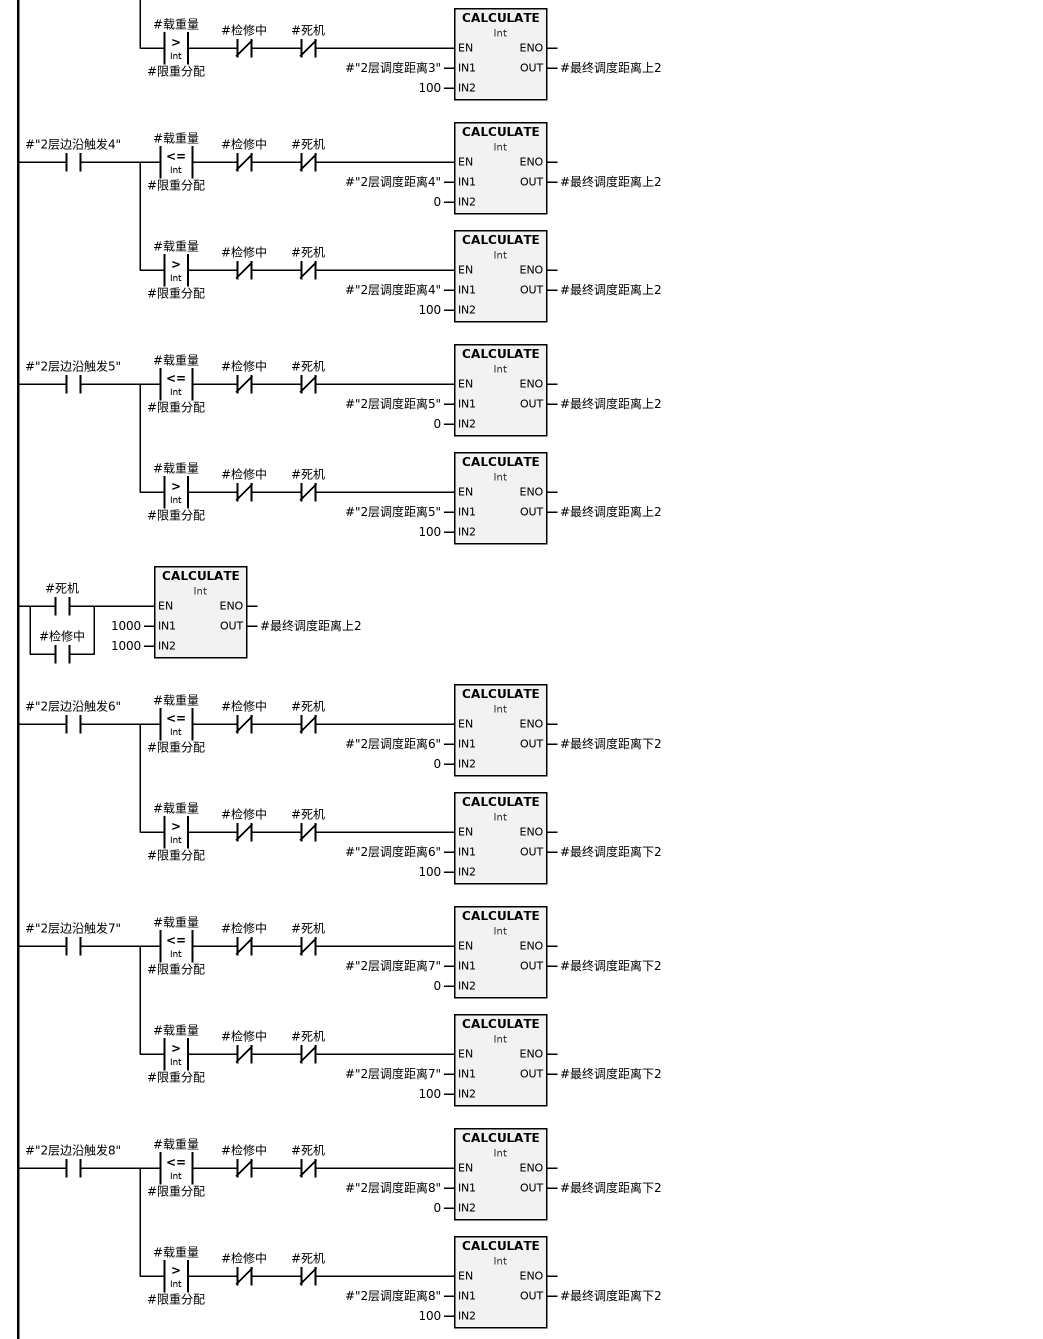
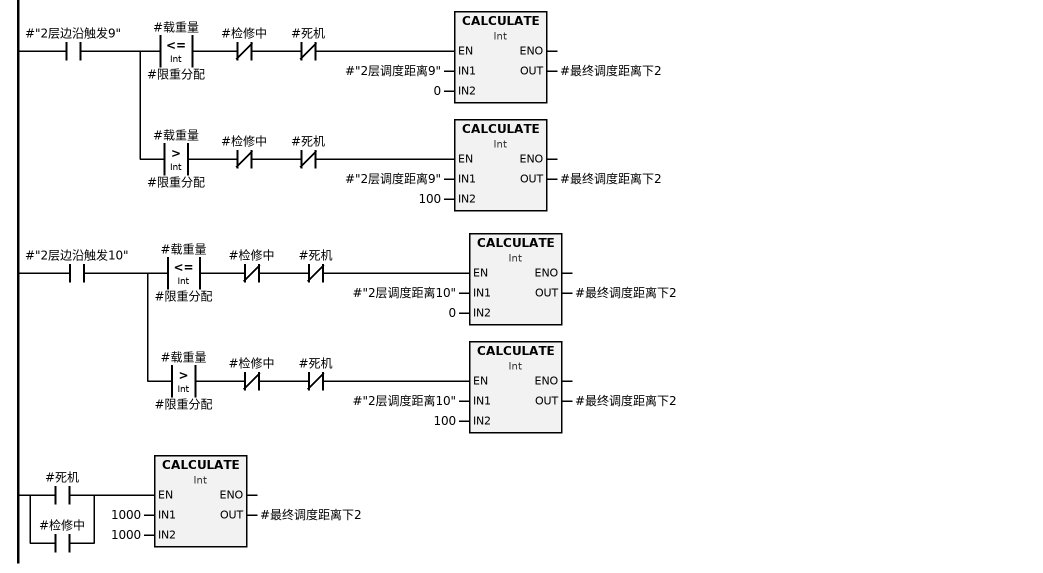
   RUNG wire#powerrail
      Contact( #上呼灯2 )
      wire#w1
      I_Contact( #上行指示 )
      I_Contact( #下行指示 )
      { S7_Templates := "SrcType := Int" } LE_Contact(in1 := #当前楼层, in2 := 2)
      wire#w2
      { S7_Templates := "SrcType := Int"; S7_Expression := "ABS(IN1-IN2)" } Calculate(in1 := #当前楼层, in2 := 2, in3 := 0, out => #"2层调度距离1")
      Coil( #"2层边沿触发1" )
   END_RUNG
   RUNG wire#w1
      Contact( #上行指示 )
      wire#w3
      { S7_Templates := "SrcType := Int" } EQ_Contact(in1 := 2, in2 := #当前楼层)
      Contact( #上下平层都为1 )
   END_RUNG wire#w2
   RUNG wire#w3
      { S7_Templates := "SrcType := Int" } GT_Contact(in1 := 2, in2 := #当前楼层)
   END_RUNG wire#w2
   RUNG wire#w1
      Contact( #下行指示 )
      wire#w4
      Contact( #外呼下面无目标2 )
      { S7_Templates := "SrcType := Int"; S7_Expression := "ABS(IN1-IN2)+IN3+IN3" } Calculate(in1 := #当前楼层, in2 := 2, in3 := #下行停站次数2, out => #"2层调度距离2")
      Coil( #"2层边沿触发2" )
   END_RUNG
   RUNG wire#w1
      I_Contact( #上行指示 )
      I_Contact( #下行指示 )
      { S7_Templates := "SrcType := Int" } GT_Contact(in1 := #当前楼层, in2 := 2)
   END_RUNG wire#w4
   RUNG wire#w1
      Contact( #下行指示 )
      Contact( #外呼下面有目标2 )
      { S7_Templates := "SrcType := Int"; S7_Expression := "ABS(IN3+IN3-IN1-IN2)+IN5+IN4+IN4+IN5+IN6" } Calculate(in1 := #当前楼层, in2 := 2, in3 := #外呼下面有目标最小数2, in4 := 0, in5 := #下行停站次数1, in6 := 2, out => #"2层调度距离3")
      Coil( #"2层边沿触发3" )
   END_RUNG
   RUNG wire#w1
      Contact( #上行指示 )
      wire#w5
      { S7_Templates := "SrcType := Int" } EQ_Contact(in1 := 2, in2 := #当前楼层)
      I_Contact( #上下平层都为1 )
      wire#w6
      Contact( #外呼下面有目标2 )
      { S7_Templates := "SrcType := Int"; S7_Expression := "ABS(IN3-IN1+IN3-IN6+IN2-IN6)+IN5+IN4+IN4+IN5+IN7+IN7+IN8+IN8" } Calculate(in1 := #当前楼层, in2 := 2, in3 := #外呼上面有目标最大数2, in4 := #上行停站次数10, in5 := 0, in6 := #外呼下面有目标最小数2, in7 := #下行停站次数1, in8 := 2, out => #"2层调度距离4")
      Coil( #"2层边沿触发4" )
   END_RUNG
   RUNG wire#w5
      { S7_Templates := "SrcType := Int" } GT_Contact(in1 := #当前楼层, in2 := 2)
   END_RUNG wire#w6
   RUNG wire#w6
      Contact( #外呼下面无目标2 )
      { S7_Templates := "SrcType := Int"; S7_Expression := "ABS(IN3-IN1+IN3-IN2)+IN5+IN4+IN4+IN5+IN6" } Calculate(in1 := #当前楼层, in2 := 2, in3 := #外呼上面有目标最大数2, in4 := #上行停站次数10, in5 := #下行停站次数2, in6 := 2, out => #"2层调度距离5")
      Coil( #"2层边沿触发5" )
   END_RUNG
   RUNG wire#powerrail
      Contact( #下呼灯2 )
      wire#w7
      I_Contact( #上行指示 )
      I_Contact( #下行指示 )
      { S7_Templates := "SrcType := Int" } GE_Contact(in1 := #当前楼层, in2 := 2)
      wire#w8
      { S7_Templates := "SrcType := Int"; S7_Expression := "ABS(IN1-IN2)+IN3+IN3" } Calculate(in1 := #当前楼层, in2 := 2, in3 := #下行停站次数2, out => #"2层调度距离6")
      Coil( #"2层边沿触发6" )
   END_RUNG
   RUNG wire#w7
      Contact( #下行指示 )
      wire#w9
      { S7_Templates := "SrcType := Int" } EQ_Contact(in1 := 2, in2 := #当前楼层)
      Contact( #上下平层都为1 )
   END_RUNG wire#w8
   RUNG wire#w9
      { S7_Templates := "SrcType := Int" } GT_Contact(in1 := #当前楼层, in2 := 2)
   END_RUNG wire#w8
   RUNG wire#w7
      Contact( #上行指示 )
      wire#w10
      Contact( #外呼上面无目标2 )
      { S7_Templates := "SrcType := Int"; S7_Expression := "ABS(IN1-IN2)+IN3+IN3" } Calculate(in1 := #当前楼层, in2 := 2, in3 := 0, out => #"2层调度距离7")
      Coil( #"2层边沿触发7" )
   END_RUNG
   RUNG wire#w7
      I_Contact( #上行指示 )
      I_Contact( #下行指示 )
      { S7_Templates := "SrcType := Int" } LT_Contact(in1 := #当前楼层, in2 := 2)
   END_RUNG wire#w10
   RUNG wire#w7
      Contact( #上行指示 )
      Contact( #外呼上面有目标2 )
      { S7_Templates := "SrcType := Int"; S7_Expression := "ABS(IN3+IN3-IN1-IN2)+IN4+IN5+IN4+IN5+IN6" } Calculate(in1 := #当前楼层, in2 := 2, in3 := #外呼上面有目标最大数2, in4 := #下行停站次数2, in5 := #上行停站次数10, in6 := 2, out => #"2层调度距离8")
      Coil( #"2层边沿触发8" )
   END_RUNG
   RUNG wire#w7
      Contact( #下行指示 )
      wire#w11
      { S7_Templates := "SrcType := Int" } EQ_Contact(in1 := 2, in2 := #当前楼层)
      I_Contact( #上下平层都为1 )
      wire#w12
      Contact( #外呼上面有目标2 )
      { S7_Templates := "SrcType := Int"; S7_Expression := "ABS(IN1-IN6+IN3-IN6+IN3-IN2)+IN5+IN4+IN4+IN5+IN7+IN7+IN8" } Calculate(in1 := #当前楼层, in2 := 2, in3 := #外呼上面有目标最大数2, in4 := #下行停站次数2, in5 := #下行停站次数1, in6 := #外呼下面有目标最小数2, in7 := #上行停站次数10, in8 := 4, out => #"2层调度距离9")
      Coil( #"2层边沿触发9" )
   END_RUNG
   RUNG wire#w11
      { S7_Templates := "SrcType := Int" } GT_Contact(in1 := 2, in2 := #当前楼层)
   END_RUNG wire#w12
   RUNG wire#w12
      Contact( #外呼上面无目标2 )
      { S7_Templates := "SrcType := Int"; S7_Expression := "ABS(IN1-IN3+IN2-IN3)+IN5+IN4+IN4+IN5+IN6" } Calculate(in1 := #当前楼层, in2 := 2, in3 := #外呼下面有目标最小数2, in4 := 0, in5 := #下行停站次数1, in6 := 2, out => #"2层调度距离10")
      Coil( #"2层边沿触发10" )
   END_RUNG
   RUNG wire#powerrail
      Contact( #"2层边沿触发1" )
      wire#w13
      { S7_Templates := "SrcType := Int" } LE_Contact(in1 := #载重量, in2 := #限重分配)
      I_Contact( #检修中 )
      I_Contact( #死机 )
      { S7_Templates := "SrcType := Int"; S7_Expression := "ABS(IN1+IN2)" } Calculate(in1 := #"2层调度距离1", in2 := 0, out => #最终调度距离上2)
   END_RUNG
   RUNG wire#w13
      { S7_Templates := "SrcType := Int" } GT_Contact(in1 := #载重量, in2 := #限重分配)
      I_Contact( #检修中 )
      I_Contact( #死机 )
      { S7_Templates := "SrcType := Int"; S7_Expression := "ABS(IN1+IN2)" } Calculate(in1 := #"2层调度距离1", in2 := 100, out => #最终调度距离上2)
   END_RUNG
   RUNG wire#powerrail
      Contact( #"2层边沿触发2" )
      wire#w14
      { S7_Templates := "SrcType := Int" } LE_Contact(in1 := #载重量, in2 := #限重分配)
      I_Contact( #检修中 )
      I_Contact( #死机 )
      { S7_Templates := "SrcType := Int"; S7_Expression := "ABS(IN1+IN2)" } Calculate(in1 := #"2层调度距离2", in2 := 0, out => #最终调度距离上2)
   END_RUNG
   RUNG wire#w14
      { S7_Templates := "SrcType := Int" } GT_Contact(in1 := #载重量, in2 := #限重分配)
      I_Contact( #检修中 )
      I_Contact( #死机 )
      { S7_Templates := "SrcType := Int"; S7_Expression := "ABS(IN1+IN2)" } Calculate(in1 := #"2层调度距离2", in2 := 100, out => #最终调度距离上2)
   END_RUNG
   RUNG wire#powerrail
      Contact( #"2层边沿触发3" )
      wire#w15
      { S7_Templates := "SrcType := Int" } LE_Contact(in1 := #载重量, in2 := #限重分配)
      I_Contact( #检修中 )
      I_Contact( #死机 )
      { S7_Templates := "SrcType := Int"; S7_Expression := "ABS(IN1+IN2)" } Calculate(in1 := #"2层调度距离3", in2 := 0, out => #最终调度距离上2)
   END_RUNG
   RUNG wire#w15
      { S7_Templates := "SrcType := Int" } GT_Contact(in1 := #载重量, in2 := #限重分配)
      I_Contact( #检修中 )
      I_Contact( #死机 )
      { S7_Templates := "SrcType := Int"; S7_Expression := "ABS(IN1+IN2)" } Calculate(in1 := #"2层调度距离3", in2 := 100, out => #最终调度距离上2)
   END_RUNG
   RUNG wire#powerrail
      Contact( #"2层边沿触发4" )
      wire#w16
      { S7_Templates := "SrcType := Int" } LE_Contact(in1 := #载重量, in2 := #限重分配)
      I_Contact( #检修中 )
      I_Contact( #死机 )
      { S7_Templates := "SrcType := Int"; S7_Expression := "ABS(IN1+IN2)" } Calculate(in1 := #"2层调度距离4", in2 := 0, out => #最终调度距离上2)
   END_RUNG
   RUNG wire#w16
      { S7_Templates := "SrcType := Int" } GT_Contact(in1 := #载重量, in2 := #限重分配)
      I_Contact( #检修中 )
      I_Contact( #死机 )
      { S7_Templates := "SrcType := Int"; S7_Expression := "ABS(IN1+IN2)" } Calculate(in1 := #"2层调度距离4", in2 := 100, out => #最终调度距离上2)
   END_RUNG
   RUNG wire#powerrail
      Contact( #"2层边沿触发5" )
      wire#w17
      { S7_Templates := "SrcType := Int" } LE_Contact(in1 := #载重量, in2 := #限重分配)
      I_Contact( #检修中 )
      I_Contact( #死机 )
      { S7_Templates := "SrcType := Int"; S7_Expression := "ABS(IN1+IN2)" } Calculate(in1 := #"2层调度距离5", in2 := 0, out => #最终调度距离上2)
   END_RUNG
   RUNG wire#w17
      { S7_Templates := "SrcType := Int" } GT_Contact(in1 := #载重量, in2 := #限重分配)
      I_Contact( #检修中 )
      I_Contact( #死机 )
      { S7_Templates := "SrcType := Int"; S7_Expression := "ABS(IN1+IN2)" } Calculate(in1 := #"2层调度距离5", in2 := 100, out => #最终调度距离上2)
   END_RUNG
   RUNG wire#powerrail
      Contact( #死机 )
      wire#w18
      { S7_Templates := "SrcType := Int"; S7_Expression := "ABS(IN1+IN2)" } Calculate(in1 := 1000, in2 := 1000, out => #最终调度距离上2)
   END_RUNG
   RUNG wire#powerrail
      Contact( #检修中 )
   END_RUNG wire#w18
   RUNG wire#powerrail
      Contact( #"2层边沿触发6" )
      wire#w19
      { S7_Templates := "SrcType := Int" } LE_Contact(in1 := #载重量, in2 := #限重分配)
      I_Contact( #检修中 )
      I_Contact( #死机 )
      { S7_Templates := "SrcType := Int"; S7_Expression := "ABS(IN1+IN2)" } Calculate(in1 := #"2层调度距离6", in2 := 0, out => #最终调度距离下2)
   END_RUNG
   RUNG wire#w19
      { S7_Templates := "SrcType := Int" } GT_Contact(in1 := #载重量, in2 := #限重分配)
      I_Contact( #检修中 )
      I_Contact( #死机 )
      { S7_Templates := "SrcType := Int"; S7_Expression := "ABS(IN1+IN2)" } Calculate(in1 := #"2层调度距离6", in2 := 100, out => #最终调度距离下2)
   END_RUNG
   RUNG wire#powerrail
      Contact( #"2层边沿触发7" )
      wire#w20
      { S7_Templates := "SrcType := Int" } LE_Contact(in1 := #载重量, in2 := #限重分配)
      I_Contact( #检修中 )
      I_Contact( #死机 )
      { S7_Templates := "SrcType := Int"; S7_Expression := "ABS(IN1+IN2)" } Calculate(in1 := #"2层调度距离7", in2 := 0, out => #最终调度距离下2)
   END_RUNG
   RUNG wire#w20
      { S7_Templates := "SrcType := Int" } GT_Contact(in1 := #载重量, in2 := #限重分配)
      I_Contact( #检修中 )
      I_Contact( #死机 )
      { S7_Templates := "SrcType := Int"; S7_Expression := "ABS(IN1+IN2)" } Calculate(in1 := #"2层调度距离7", in2 := 100, out => #最终调度距离下2)
   END_RUNG
   RUNG wire#powerrail
      Contact( #"2层边沿触发8" )
      wire#w21
      { S7_Templates := "SrcType := Int" } LE_Contact(in1 := #载重量, in2 := #限重分配)
      I_Contact( #检修中 )
      I_Contact( #死机 )
      { S7_Templates := "SrcType := Int"; S7_Expression := "ABS(IN1+IN2)" } Calculate(in1 := #"2层调度距离8", in2 := 0, out => #最终调度距离下2)
   END_RUNG
   RUNG wire#w21
      { S7_Templates := "SrcType := Int" } GT_Contact(in1 := #载重量, in2 := #限重分配)
      I_Contact( #检修中 )
      I_Contact( #死机 )
      { S7_Templates := "SrcType := Int"; S7_Expression := "ABS(IN1+IN2)" } Calculate(in1 := #"2层调度距离8", in2 := 100, out => #最终调度距离下2)
   END_RUNG
   RUNG wire#powerrail
      Contact( #"2层边沿触发9" )
      wire#w22
      { S7_Templates := "SrcType := Int" } LE_Contact(in1 := #载重量, in2 := #限重分配)
      I_Contact( #检修中 )
      I_Contact( #死机 )
      { S7_Templates := "SrcType := Int"; S7_Expression := "ABS(IN1+IN2)" } Calculate(in1 := #"2层调度距离9", in2 := 0, out => #最终调度距离下2)
   END_RUNG
   RUNG wire#w22
      { S7_Templates := "SrcType := Int" } GT_Contact(in1 := #载重量, in2 := #限重分配)
      I_Contact( #检修中 )
      I_Contact( #死机 )
      { S7_Templates := "SrcType := Int"; S7_Expression := "ABS(IN1+IN2)" } Calculate(in1 := #"2层调度距离9", in2 := 100, out => #最终调度距离下2)
   END_RUNG
   RUNG wire#powerrail
      Contact( #"2层边沿触发10" )
      wire#w23
      { S7_Templates := "SrcType := Int" } LE_Contact(in1 := #载重量, in2 := #限重分配)
      I_Contact( #检修中 )
      I_Contact( #死机 )
      { S7_Templates := "SrcType := Int"; S7_Expression := "ABS(IN1+IN2)" } Calculate(in1 := #"2层调度距离10", in2 := 0, out => #最终调度距离下2)
   END_RUNG
   RUNG wire#w23
      { S7_Templates := "SrcType := Int" } GT_Contact(in1 := #载重量, in2 := #限重分配)
      I_Contact( #检修中 )
      I_Contact( #死机 )
      { S7_Templates := "SrcType := Int"; S7_Expression := "ABS(IN1+IN2)" } Calculate(in1 := #"2层调度距离10", in2 := 100, out => #最终调度距离下2)
   END_RUNG
   RUNG wire#powerrail
      Contact( #死机 )
      wire#w24
      { S7_Templates := "SrcType := Int"; S7_Expression := "ABS(IN1+IN2)" } Calculate(in1 := 1000, in2 := 1000, out => #最终调度距离下2)
   END_RUNG
   RUNG wire#powerrail
      Contact( #检修中 )
   END_RUNG wire#w24
   // the same network as SCL:
   #_w1 := #上呼灯2 AND ((NOT #上行指示 AND NOT #下行指示 AND (#当前楼层 <= 2)) OR (#上行指示 AND (((2 = #当前楼层) AND #上下平层都为1) OR (2 > #当前楼层))));
   IF #_w1 THEN #"2层调度距离1" := ABS(#当前楼层-2); END_IF;
   #"2层边沿触发1" := #_w1;
   #_w2 := #上呼灯2 AND (#下行指示 OR (NOT #上行指示 AND NOT #下行指示 AND (#当前楼层 > 2))) AND #外呼下面无目标2;
   IF #_w2 THEN #"2层调度距离2" := ABS(#当前楼层-2)+#下行停站次数2+#下行停站次数2; END_IF;
   #"2层边沿触发2" := #_w2;
   #_w3 := #上呼灯2 AND #下行指示 AND #外呼下面有目标2;
   IF #_w3 THEN #"2层调度距离3" := ABS(#外呼下面有目标最小数2+#外呼下面有目标最小数2-#当前楼层-2)+#下行停站次数1+0+0+#下行停站次数1+2; END_IF;
   #"2层边沿触发3" := #_w3;
   #_w4 := #上呼灯2 AND #上行指示 AND (((2 = #当前楼层) AND NOT #上下平层都为1) OR (#当前楼层 > 2));
   #_w5 := #_w4 AND #外呼下面有目标2;
   IF #_w5 THEN
       #"2层调度距离4" := ABS(#外呼上面有目标最大数2-#当前楼层+#外呼上面有目标最大数2-#外呼下面有目标最小数2+2-#外呼下面有目标最小数2)+0+#上行停站次数10+#上行停站次数10+0+#下行停站次数1+#下行停站次数1+2+2;
   END_IF;
   #"2层边沿触发4" := #_w5;
   #_w6 := #_w4 AND #外呼下面无目标2;
   IF #_w6 THEN
       #"2层调度距离5" := ABS(#外呼上面有目标最大数2-#当前楼层+#外呼上面有目标最大数2-2)+#下行停站次数2+#上行停站次数10+#上行停站次数10+#下行停站次数2+2;
   END_IF;
   #"2层边沿触发5" := #_w6;
   #_w7 := #下呼灯2 AND ((NOT #上行指示 AND NOT #下行指示 AND (#当前楼层 >= 2)) OR (#下行指示 AND (((2 = #当前楼层) AND #上下平层都为1) OR (#当前楼层 > 2))));
   IF #_w7 THEN #"2层调度距离6" := ABS(#当前楼层-2)+#下行停站次数2+#下行停站次数2; END_IF;
   #"2层边沿触发6" := #_w7;
   #_w8 := #下呼灯2 AND (#上行指示 OR (NOT #上行指示 AND NOT #下行指示 AND (#当前楼层 < 2))) AND #外呼上面无目标2;
   IF #_w8 THEN #"2层调度距离7" := ABS(#当前楼层-2)+0+0; END_IF;
   #"2层边沿触发7" := #_w8;
   #_w9 := #下呼灯2 AND #上行指示 AND #外呼上面有目标2;
   IF #_w9 THEN
       #"2层调度距离8" := ABS(#外呼上面有目标最大数2+#外呼上面有目标最大数2-#当前楼层-2)+#下行停站次数2+#上行停站次数10+#下行停站次数2+#上行停站次数10+2;
   END_IF;
   #"2层边沿触发8" := #_w9;
   #_w10 := #下呼灯2 AND #下行指示 AND (((2 = #当前楼层) AND NOT #上下平层都为1) OR (2 > #当前楼层));
   #_w11 := #_w10 AND #外呼上面有目标2;
   IF #_w11 THEN
       #"2层调度距离9" := ABS(#当前楼层-#外呼下面有目标最小数2+#外呼上面有目标最大数2-#外呼下面有目标最小数2+#外呼上面有目标最大数2-2)+#下行停站次数1+#下行停站次数2+#下行停站次数2+#下行停站次数1+#上行停站次数10+#上行停站次数10+4;
   END_IF;
   #"2层边沿触发9" := #_w11;
   #_w12 := #_w10 AND #外呼上面无目标2;
   IF #_w12 THEN #"2层调度距离10" := ABS(#当前楼层-#外呼下面有目标最小数2+2-#外呼下面有目标最小数2)+#下行停站次数1+0+0+#下行停站次数1+2; END_IF;
   #"2层边沿触发10" := #_w12;
   IF #"2层边沿触发1" AND (#载重量 <= #限重分配) AND NOT #检修中 AND NOT #死机 THEN #最终调度距离上2 := ABS(#"2层调度距离1"+0); END_IF;
   IF #"2层边沿触发1" AND (#载重量 > #限重分配) AND NOT #检修中 AND NOT #死机 THEN #最终调度距离上2 := ABS(#"2层调度距离1"+100); END_IF;
   IF #"2层边沿触发2" AND (#载重量 <= #限重分配) AND NOT #检修中 AND NOT #死机 THEN #最终调度距离上2 := ABS(#"2层调度距离2"+0); END_IF;
   IF #"2层边沿触发2" AND (#载重量 > #限重分配) AND NOT #检修中 AND NOT #死机 THEN #最终调度距离上2 := ABS(#"2层调度距离2"+100); END_IF;
   IF #"2层边沿触发3" AND (#载重量 <= #限重分配) AND NOT #检修中 AND NOT #死机 THEN #最终调度距离上2 := ABS(#"2层调度距离3"+0); END_IF;
   IF #"2层边沿触发3" AND (#载重量 > #限重分配) AND NOT #检修中 AND NOT #死机 THEN #最终调度距离上2 := ABS(#"2层调度距离3"+100); END_IF;
   IF #"2层边沿触发4" AND (#载重量 <= #限重分配) AND NOT #检修中 AND NOT #死机 THEN #最终调度距离上2 := ABS(#"2层调度距离4"+0); END_IF;
   IF #"2层边沿触发4" AND (#载重量 > #限重分配) AND NOT #检修中 AND NOT #死机 THEN #最终调度距离上2 := ABS(#"2层调度距离4"+100); END_IF;
   IF #"2层边沿触发5" AND (#载重量 <= #限重分配) AND NOT #检修中 AND NOT #死机 THEN #最终调度距离上2 := ABS(#"2层调度距离5"+0); END_IF;
   IF #"2层边沿触发5" AND (#载重量 > #限重分配) AND NOT #检修中 AND NOT #死机 THEN #最终调度距离上2 := ABS(#"2层调度距离5"+100); END_IF;
   IF #死机 OR #检修中 THEN #最终调度距离上2 := ABS(1000+1000); END_IF;
   IF #"2层边沿触发6" AND (#载重量 <= #限重分配) AND NOT #检修中 AND NOT #死机 THEN #最终调度距离下2 := ABS(#"2层调度距离6"+0); END_IF;
   IF #"2层边沿触发6" AND (#载重量 > #限重分配) AND NOT #检修中 AND NOT #死机 THEN #最终调度距离下2 := ABS(#"2层调度距离6"+100); END_IF;
   IF #"2层边沿触发7" AND (#载重量 <= #限重分配) AND NOT #检修中 AND NOT #死机 THEN #最终调度距离下2 := ABS(#"2层调度距离7"+0); END_IF;
   IF #"2层边沿触发7" AND (#载重量 > #限重分配) AND NOT #检修中 AND NOT #死机 THEN #最终调度距离下2 := ABS(#"2层调度距离7"+100); END_IF;
   IF #"2层边沿触发8" AND (#载重量 <= #限重分配) AND NOT #检修中 AND NOT #死机 THEN #最终调度距离下2 := ABS(#"2层调度距离8"+0); END_IF;
   IF #"2层边沿触发8" AND (#载重量 > #限重分配) AND NOT #检修中 AND NOT #死机 THEN #最终调度距离下2 := ABS(#"2层调度距离8"+100); END_IF;
   IF #"2层边沿触发9" AND (#载重量 <= #限重分配) AND NOT #检修中 AND NOT #死机 THEN #最终调度距离下2 := ABS(#"2层调度距离9"+0); END_IF;
   IF #"2层边沿触发9" AND (#载重量 > #限重分配) AND NOT #检修中 AND NOT #死机 THEN #最终调度距离下2 := ABS(#"2层调度距离9"+100); END_IF;
   IF #"2层边沿触发10" AND (#载重量 <= #限重分配) AND NOT #检修中 AND NOT #死机 THEN #最终调度距离下2 := ABS(#"2层调度距离10"+0); END_IF;
   IF #"2层边沿触发10" AND (#载重量 > #限重分配) AND NOT #检修中 AND NOT #死机 THEN #最终调度距离下2 := ABS(#"2层调度距离10"+100); END_IF;
   IF #死机 OR #检修中 THEN #最终调度距离下2 := ABS(1000+1000); END_IF;
END_REGION

REGION Network 2: 3层调度距离
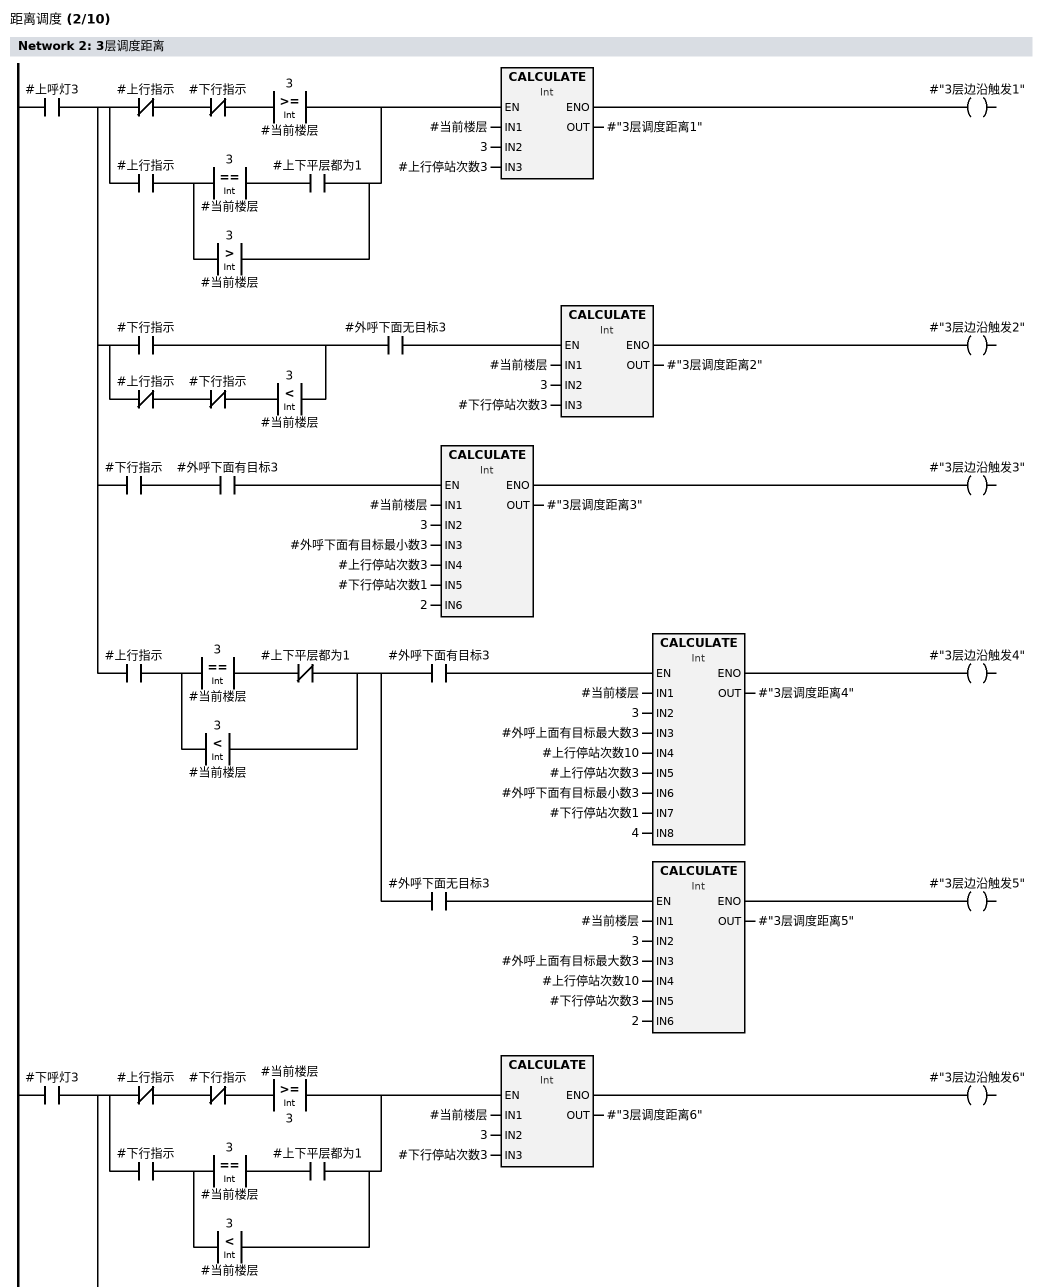
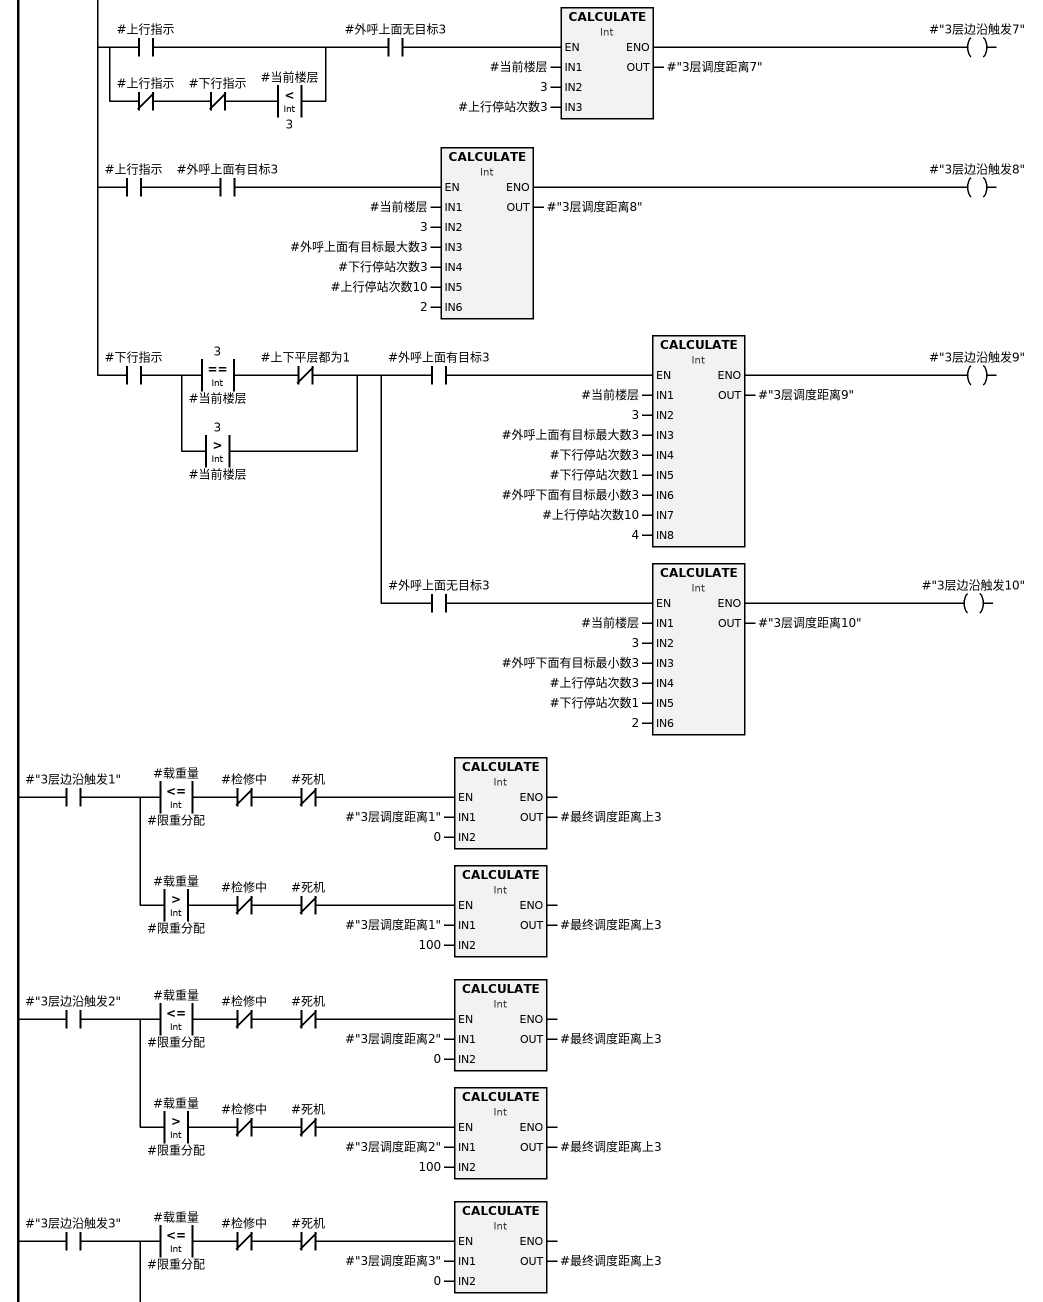
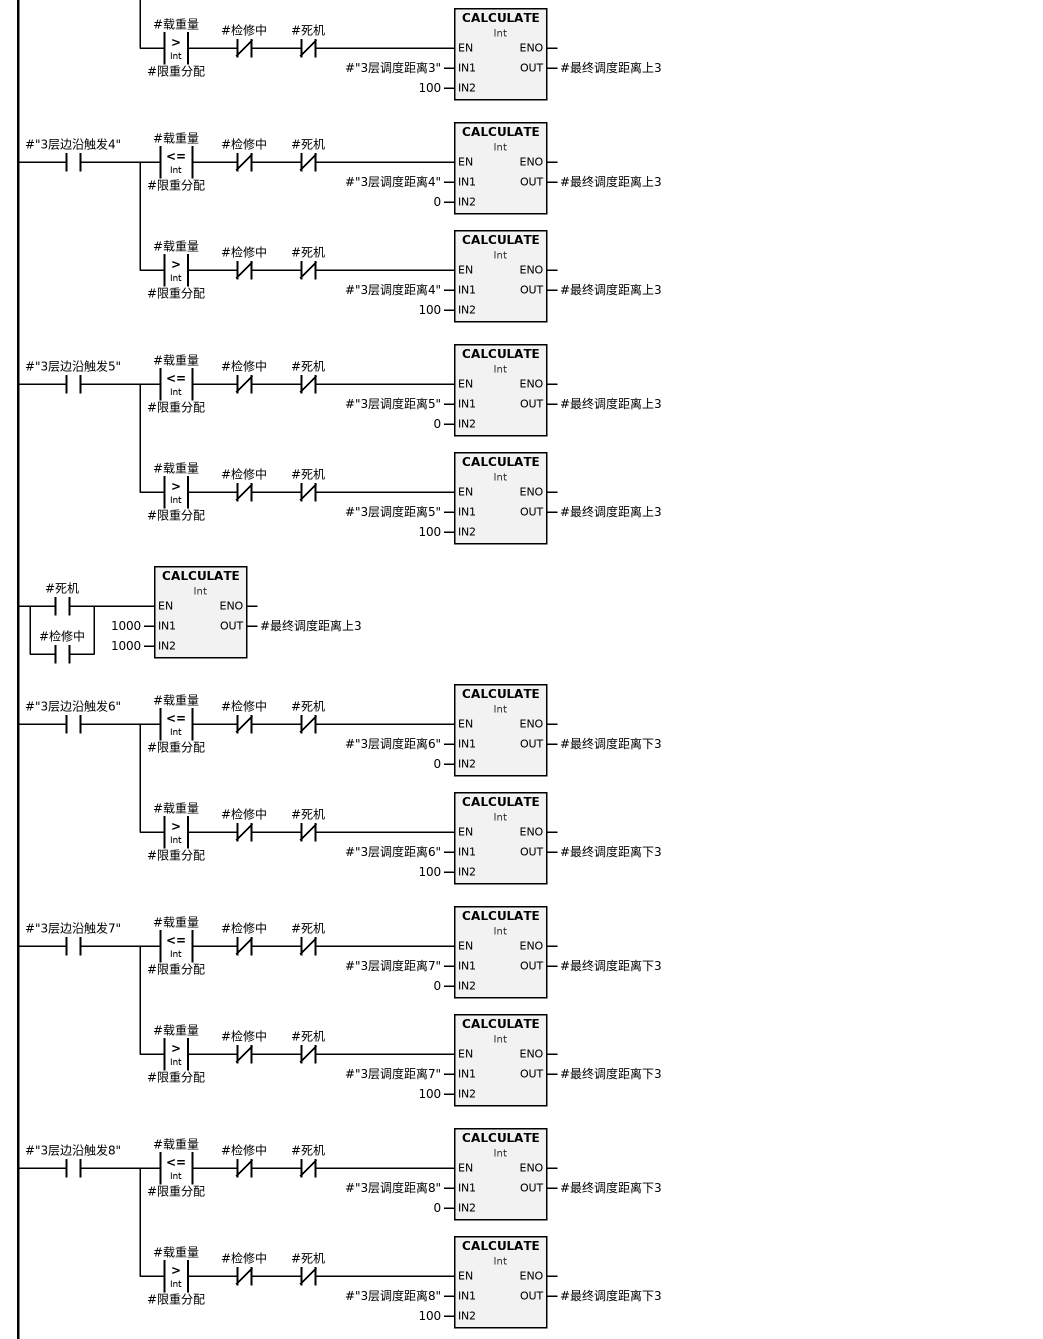
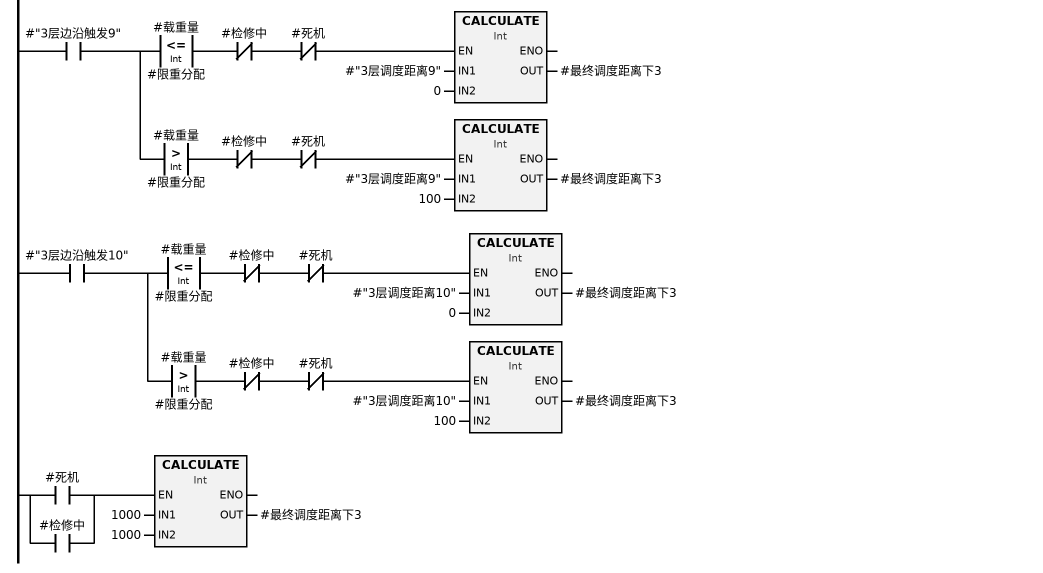
   RUNG wire#powerrail
      Contact( #上呼灯3 )
      wire#w1
      I_Contact( #上行指示 )
      I_Contact( #下行指示 )
      { S7_Templates := "SrcType := Int" } GE_Contact(in1 := 3, in2 := #当前楼层)
      wire#w2
      { S7_Templates := "SrcType := Int"; S7_Expression := "ABS(IN1-IN2)+IN3+IN3" } Calculate(in1 := #当前楼层, in2 := 3, in3 := #上行停站次数3, out => #"3层调度距离1")
      Coil( #"3层边沿触发1" )
   END_RUNG
   RUNG wire#w1
      Contact( #上行指示 )
      wire#w3
      { S7_Templates := "SrcType := Int" } EQ_Contact(in1 := 3, in2 := #当前楼层)
      Contact( #上下平层都为1 )
   END_RUNG wire#w2
   RUNG wire#w3
      { S7_Templates := "SrcType := Int" } GT_Contact(in1 := 3, in2 := #当前楼层)
   END_RUNG wire#w2
   RUNG wire#w1
      Contact( #下行指示 )
      wire#w4
      Contact( #外呼下面无目标3 )
      { S7_Templates := "SrcType := Int"; S7_Expression := "ABS(IN1-IN2)+IN3+IN3" } Calculate(in1 := #当前楼层, in2 := 3, in3 := #下行停站次数3, out => #"3层调度距离2")
      Coil( #"3层边沿触发2" )
   END_RUNG
   RUNG wire#w1
      I_Contact( #上行指示 )
      I_Contact( #下行指示 )
      { S7_Templates := "SrcType := Int" } LT_Contact(in1 := 3, in2 := #当前楼层)
   END_RUNG wire#w4
   RUNG wire#w1
      Contact( #下行指示 )
      Contact( #外呼下面有目标3 )
      { S7_Templates := "SrcType := Int"; S7_Expression := "ABS(IN3+IN3-IN1-IN2)+IN5+IN4+IN4+IN5+IN6" } Calculate(in1 := #当前楼层, in2 := 3, in3 := #外呼下面有目标最小数3, in4 := #上行停站次数3, in5 := #下行停站次数1, in6 := 2, out => #"3层调度距离3")
      Coil( #"3层边沿触发3" )
   END_RUNG
   RUNG wire#w1
      Contact( #上行指示 )
      wire#w5
      { S7_Templates := "SrcType := Int" } EQ_Contact(in1 := 3, in2 := #当前楼层)
      I_Contact( #上下平层都为1 )
      wire#w6
      Contact( #外呼下面有目标3 )
      { S7_Templates := "SrcType := Int"; S7_Expression := "ABS(IN3-IN1+IN3-IN6+IN2-IN6)+IN5+IN4+IN4+IN5+IN7+IN7+IN8" } Calculate(in1 := #当前楼层, in2 := 3, in3 := #外呼上面有目标最大数3, in4 := #上行停站次数10, in5 := #上行停站次数3, in6 := #外呼下面有目标最小数3, in7 := #下行停站次数1, in8 := 4, out => #"3层调度距离4")
      Coil( #"3层边沿触发4" )
   END_RUNG
   RUNG wire#w5
      { S7_Templates := "SrcType := Int" } LT_Contact(in1 := 3, in2 := #当前楼层)
   END_RUNG wire#w6
   RUNG wire#w6
      Contact( #外呼下面无目标3 )
      { S7_Templates := "SrcType := Int"; S7_Expression := "ABS(IN3-IN1+IN3-IN2)+IN5+IN4+IN4+IN5+IN6" } Calculate(in1 := #当前楼层, in2 := 3, in3 := #外呼上面有目标最大数3, in4 := #上行停站次数10, in5 := #下行停站次数3, in6 := 2, out => #"3层调度距离5")
      Coil( #"3层边沿触发5" )
   END_RUNG
   RUNG wire#powerrail
      Contact( #下呼灯3 )
      wire#w7
      I_Contact( #上行指示 )
      I_Contact( #下行指示 )
      { S7_Templates := "SrcType := Int" } GE_Contact(in1 := #当前楼层, in2 := 3)
      wire#w8
      { S7_Templates := "SrcType := Int"; S7_Expression := "ABS(IN1-IN2)+IN3+IN3" } Calculate(in1 := #当前楼层, in2 := 3, in3 := #下行停站次数3, out => #"3层调度距离6")
      Coil( #"3层边沿触发6" )
   END_RUNG
   RUNG wire#w7
      Contact( #下行指示 )
      wire#w9
      { S7_Templates := "SrcType := Int" } EQ_Contact(in1 := 3, in2 := #当前楼层)
      Contact( #上下平层都为1 )
   END_RUNG wire#w8
   RUNG wire#w9
      { S7_Templates := "SrcType := Int" } LT_Contact(in1 := 3, in2 := #当前楼层)
   END_RUNG wire#w8
   RUNG wire#w7
      Contact( #上行指示 )
      wire#w10
      Contact( #外呼上面无目标3 )
      { S7_Templates := "SrcType := Int"; S7_Expression := "ABS(IN1-IN2)+IN3+IN3" } Calculate(in1 := #当前楼层, in2 := 3, in3 := #上行停站次数3, out => #"3层调度距离7")
      Coil( #"3层边沿触发7" )
   END_RUNG
   RUNG wire#w7
      I_Contact( #上行指示 )
      I_Contact( #下行指示 )
      { S7_Templates := "SrcType := Int" } LT_Contact(in1 := #当前楼层, in2 := 3)
   END_RUNG wire#w10
   RUNG wire#w7
      Contact( #上行指示 )
      Contact( #外呼上面有目标3 )
      { S7_Templates := "SrcType := Int"; S7_Expression := "ABS(IN3+IN3-IN1-IN2)+IN4+IN5+IN4+IN5+IN6" } Calculate(in1 := #当前楼层, in2 := 3, in3 := #外呼上面有目标最大数3, in4 := #下行停站次数3, in5 := #上行停站次数10, in6 := 2, out => #"3层调度距离8")
      Coil( #"3层边沿触发8" )
   END_RUNG
   RUNG wire#w7
      Contact( #下行指示 )
      wire#w11
      { S7_Templates := "SrcType := Int" } EQ_Contact(in1 := 3, in2 := #当前楼层)
      I_Contact( #上下平层都为1 )
      wire#w12
      Contact( #外呼上面有目标3 )
      { S7_Templates := "SrcType := Int"; S7_Expression := "ABS(IN1-IN6+IN3-IN6+IN3-IN2)+IN5+IN4+IN4+IN5+IN7+IN7+IN8" } Calculate(in1 := #当前楼层, in2 := 3, in3 := #外呼上面有目标最大数3, in4 := #下行停站次数3, in5 := #下行停站次数1, in6 := #外呼下面有目标最小数3, in7 := #上行停站次数10, in8 := 4, out => #"3层调度距离9")
      Coil( #"3层边沿触发9" )
   END_RUNG
   RUNG wire#w11
      { S7_Templates := "SrcType := Int" } GT_Contact(in1 := 3, in2 := #当前楼层)
   END_RUNG wire#w12
   RUNG wire#w12
      Contact( #外呼上面无目标3 )
      { S7_Templates := "SrcType := Int"; S7_Expression := "ABS(IN1-IN3+IN2-IN3)+IN5+IN4+IN4+IN5+IN6" } Calculate(in1 := #当前楼层, in2 := 3, in3 := #外呼下面有目标最小数3, in4 := #上行停站次数3, in5 := #下行停站次数1, in6 := 2, out => #"3层调度距离10")
      Coil( #"3层边沿触发10" )
   END_RUNG
   RUNG wire#powerrail
      Contact( #"3层边沿触发1" )
      wire#w13
      { S7_Templates := "SrcType := Int" } LE_Contact(in1 := #载重量, in2 := #限重分配)
      I_Contact( #检修中 )
      I_Contact( #死机 )
      { S7_Templates := "SrcType := Int"; S7_Expression := "ABS(IN1+IN2)" } Calculate(in1 := #"3层调度距离1", in2 := 0, out => #最终调度距离上3)
   END_RUNG
   RUNG wire#w13
      { S7_Templates := "SrcType := Int" } GT_Contact(in1 := #载重量, in2 := #限重分配)
      I_Contact( #检修中 )
      I_Contact( #死机 )
      { S7_Templates := "SrcType := Int"; S7_Expression := "ABS(IN1+IN2)" } Calculate(in1 := #"3层调度距离1", in2 := 100, out => #最终调度距离上3)
   END_RUNG
   RUNG wire#powerrail
      Contact( #"3层边沿触发2" )
      wire#w14
      { S7_Templates := "SrcType := Int" } LE_Contact(in1 := #载重量, in2 := #限重分配)
      I_Contact( #检修中 )
      I_Contact( #死机 )
      { S7_Templates := "SrcType := Int"; S7_Expression := "ABS(IN1+IN2)" } Calculate(in1 := #"3层调度距离2", in2 := 0, out => #最终调度距离上3)
   END_RUNG
   RUNG wire#w14
      { S7_Templates := "SrcType := Int" } GT_Contact(in1 := #载重量, in2 := #限重分配)
      I_Contact( #检修中 )
      I_Contact( #死机 )
      { S7_Templates := "SrcType := Int"; S7_Expression := "ABS(IN1+IN2)" } Calculate(in1 := #"3层调度距离2", in2 := 100, out => #最终调度距离上3)
   END_RUNG
   RUNG wire#powerrail
      Contact( #"3层边沿触发3" )
      wire#w15
      { S7_Templates := "SrcType := Int" } LE_Contact(in1 := #载重量, in2 := #限重分配)
      I_Contact( #检修中 )
      I_Contact( #死机 )
      { S7_Templates := "SrcType := Int"; S7_Expression := "ABS(IN1+IN2)" } Calculate(in1 := #"3层调度距离3", in2 := 0, out => #最终调度距离上3)
   END_RUNG
   RUNG wire#w15
      { S7_Templates := "SrcType := Int" } GT_Contact(in1 := #载重量, in2 := #限重分配)
      I_Contact( #检修中 )
      I_Contact( #死机 )
      { S7_Templates := "SrcType := Int"; S7_Expression := "ABS(IN1+IN2)" } Calculate(in1 := #"3层调度距离3", in2 := 100, out => #最终调度距离上3)
   END_RUNG
   RUNG wire#powerrail
      Contact( #"3层边沿触发4" )
      wire#w16
      { S7_Templates := "SrcType := Int" } LE_Contact(in1 := #载重量, in2 := #限重分配)
      I_Contact( #检修中 )
      I_Contact( #死机 )
      { S7_Templates := "SrcType := Int"; S7_Expression := "ABS(IN1+IN2)" } Calculate(in1 := #"3层调度距离4", in2 := 0, out => #最终调度距离上3)
   END_RUNG
   RUNG wire#w16
      { S7_Templates := "SrcType := Int" } GT_Contact(in1 := #载重量, in2 := #限重分配)
      I_Contact( #检修中 )
      I_Contact( #死机 )
      { S7_Templates := "SrcType := Int"; S7_Expression := "ABS(IN1+IN2)" } Calculate(in1 := #"3层调度距离4", in2 := 100, out => #最终调度距离上3)
   END_RUNG
   RUNG wire#powerrail
      Contact( #"3层边沿触发5" )
      wire#w17
      { S7_Templates := "SrcType := Int" } LE_Contact(in1 := #载重量, in2 := #限重分配)
      I_Contact( #检修中 )
      I_Contact( #死机 )
      { S7_Templates := "SrcType := Int"; S7_Expression := "ABS(IN1+IN2)" } Calculate(in1 := #"3层调度距离5", in2 := 0, out => #最终调度距离上3)
   END_RUNG
   RUNG wire#w17
      { S7_Templates := "SrcType := Int" } GT_Contact(in1 := #载重量, in2 := #限重分配)
      I_Contact( #检修中 )
      I_Contact( #死机 )
      { S7_Templates := "SrcType := Int"; S7_Expression := "ABS(IN1+IN2)" } Calculate(in1 := #"3层调度距离5", in2 := 100, out => #最终调度距离上3)
   END_RUNG
   RUNG wire#powerrail
      Contact( #死机 )
      wire#w18
      { S7_Templates := "SrcType := Int"; S7_Expression := "ABS(IN1+IN2)" } Calculate(in1 := 1000, in2 := 1000, out => #最终调度距离上3)
   END_RUNG
   RUNG wire#powerrail
      Contact( #检修中 )
   END_RUNG wire#w18
   RUNG wire#powerrail
      Contact( #"3层边沿触发6" )
      wire#w19
      { S7_Templates := "SrcType := Int" } LE_Contact(in1 := #载重量, in2 := #限重分配)
      I_Contact( #检修中 )
      I_Contact( #死机 )
      { S7_Templates := "SrcType := Int"; S7_Expression := "ABS(IN1+IN2)" } Calculate(in1 := #"3层调度距离6", in2 := 0, out => #最终调度距离下3)
   END_RUNG
   RUNG wire#w19
      { S7_Templates := "SrcType := Int" } GT_Contact(in1 := #载重量, in2 := #限重分配)
      I_Contact( #检修中 )
      I_Contact( #死机 )
      { S7_Templates := "SrcType := Int"; S7_Expression := "ABS(IN1+IN2)" } Calculate(in1 := #"3层调度距离6", in2 := 100, out => #最终调度距离下3)
   END_RUNG
   RUNG wire#powerrail
      Contact( #"3层边沿触发7" )
      wire#w20
      { S7_Templates := "SrcType := Int" } LE_Contact(in1 := #载重量, in2 := #限重分配)
      I_Contact( #检修中 )
      I_Contact( #死机 )
      { S7_Templates := "SrcType := Int"; S7_Expression := "ABS(IN1+IN2)" } Calculate(in1 := #"3层调度距离7", in2 := 0, out => #最终调度距离下3)
   END_RUNG
   RUNG wire#w20
      { S7_Templates := "SrcType := Int" } GT_Contact(in1 := #载重量, in2 := #限重分配)
      I_Contact( #检修中 )
      I_Contact( #死机 )
      { S7_Templates := "SrcType := Int"; S7_Expression := "ABS(IN1+IN2)" } Calculate(in1 := #"3层调度距离7", in2 := 100, out => #最终调度距离下3)
   END_RUNG
   RUNG wire#powerrail
      Contact( #"3层边沿触发8" )
      wire#w21
      { S7_Templates := "SrcType := Int" } LE_Contact(in1 := #载重量, in2 := #限重分配)
      I_Contact( #检修中 )
      I_Contact( #死机 )
      { S7_Templates := "SrcType := Int"; S7_Expression := "ABS(IN1+IN2)" } Calculate(in1 := #"3层调度距离8", in2 := 0, out => #最终调度距离下3)
   END_RUNG
   RUNG wire#w21
      { S7_Templates := "SrcType := Int" } GT_Contact(in1 := #载重量, in2 := #限重分配)
      I_Contact( #检修中 )
      I_Contact( #死机 )
      { S7_Templates := "SrcType := Int"; S7_Expression := "ABS(IN1+IN2)" } Calculate(in1 := #"3层调度距离8", in2 := 100, out => #最终调度距离下3)
   END_RUNG
   RUNG wire#powerrail
      Contact( #"3层边沿触发9" )
      wire#w22
      { S7_Templates := "SrcType := Int" } LE_Contact(in1 := #载重量, in2 := #限重分配)
      I_Contact( #检修中 )
      I_Contact( #死机 )
      { S7_Templates := "SrcType := Int"; S7_Expression := "ABS(IN1+IN2)" } Calculate(in1 := #"3层调度距离9", in2 := 0, out => #最终调度距离下3)
   END_RUNG
   RUNG wire#w22
      { S7_Templates := "SrcType := Int" } GT_Contact(in1 := #载重量, in2 := #限重分配)
      I_Contact( #检修中 )
      I_Contact( #死机 )
      { S7_Templates := "SrcType := Int"; S7_Expression := "ABS(IN1+IN2)" } Calculate(in1 := #"3层调度距离9", in2 := 100, out => #最终调度距离下3)
   END_RUNG
   RUNG wire#powerrail
      Contact( #"3层边沿触发10" )
      wire#w23
      { S7_Templates := "SrcType := Int" } LE_Contact(in1 := #载重量, in2 := #限重分配)
      I_Contact( #检修中 )
      I_Contact( #死机 )
      { S7_Templates := "SrcType := Int"; S7_Expression := "ABS(IN1+IN2)" } Calculate(in1 := #"3层调度距离10", in2 := 0, out => #最终调度距离下3)
   END_RUNG
   RUNG wire#w23
      { S7_Templates := "SrcType := Int" } GT_Contact(in1 := #载重量, in2 := #限重分配)
      I_Contact( #检修中 )
      I_Contact( #死机 )
      { S7_Templates := "SrcType := Int"; S7_Expression := "ABS(IN1+IN2)" } Calculate(in1 := #"3层调度距离10", in2 := 100, out => #最终调度距离下3)
   END_RUNG
   RUNG wire#powerrail
      Contact( #死机 )
      wire#w24
      { S7_Templates := "SrcType := Int"; S7_Expression := "ABS(IN1+IN2)" } Calculate(in1 := 1000, in2 := 1000, out => #最终调度距离下3)
   END_RUNG
   RUNG wire#powerrail
      Contact( #检修中 )
   END_RUNG wire#w24
   // the same network as SCL:
   #_w1 := #上呼灯3 AND ((NOT #上行指示 AND NOT #下行指示 AND (3 >= #当前楼层)) OR (#上行指示 AND (((3 = #当前楼层) AND #上下平层都为1) OR (3 > #当前楼层))));
   IF #_w1 THEN #"3层调度距离1" := ABS(#当前楼层-3)+#上行停站次数3+#上行停站次数3; END_IF;
   #"3层边沿触发1" := #_w1;
   #_w2 := #上呼灯3 AND (#下行指示 OR (NOT #上行指示 AND NOT #下行指示 AND (3 < #当前楼层))) AND #外呼下面无目标3;
   IF #_w2 THEN #"3层调度距离2" := ABS(#当前楼层-3)+#下行停站次数3+#下行停站次数3; END_IF;
   #"3层边沿触发2" := #_w2;
   #_w3 := #上呼灯3 AND #下行指示 AND #外呼下面有目标3;
   IF #_w3 THEN
       #"3层调度距离3" := ABS(#外呼下面有目标最小数3+#外呼下面有目标最小数3-#当前楼层-3)+#下行停站次数1+#上行停站次数3+#上行停站次数3+#下行停站次数1+2;
   END_IF;
   #"3层边沿触发3" := #_w3;
   #_w4 := #上呼灯3 AND #上行指示 AND (((3 = #当前楼层) AND NOT #上下平层都为1) OR (3 < #当前楼层));
   #_w5 := #_w4 AND #外呼下面有目标3;
   IF #_w5 THEN
       #"3层调度距离4" := ABS(#外呼上面有目标最大数3-#当前楼层+#外呼上面有目标最大数3-#外呼下面有目标最小数3+3-#外呼下面有目标最小数3)+#上行停站次数3+#上行停站次数10+#上行停站次数10+#上行停站次数3+#下行停站次数1+#下行停站次数1+4;
   END_IF;
   #"3层边沿触发4" := #_w5;
   #_w6 := #_w4 AND #外呼下面无目标3;
   IF #_w6 THEN
       #"3层调度距离5" := ABS(#外呼上面有目标最大数3-#当前楼层+#外呼上面有目标最大数3-3)+#下行停站次数3+#上行停站次数10+#上行停站次数10+#下行停站次数3+2;
   END_IF;
   #"3层边沿触发5" := #_w6;
   #_w7 := #下呼灯3 AND ((NOT #上行指示 AND NOT #下行指示 AND (#当前楼层 >= 3)) OR (#下行指示 AND (((3 = #当前楼层) AND #上下平层都为1) OR (3 < #当前楼层))));
   IF #_w7 THEN #"3层调度距离6" := ABS(#当前楼层-3)+#下行停站次数3+#下行停站次数3; END_IF;
   #"3层边沿触发6" := #_w7;
   #_w8 := #下呼灯3 AND (#上行指示 OR (NOT #上行指示 AND NOT #下行指示 AND (#当前楼层 < 3))) AND #外呼上面无目标3;
   IF #_w8 THEN #"3层调度距离7" := ABS(#当前楼层-3)+#上行停站次数3+#上行停站次数3; END_IF;
   #"3层边沿触发7" := #_w8;
   #_w9 := #下呼灯3 AND #上行指示 AND #外呼上面有目标3;
   IF #_w9 THEN
       #"3层调度距离8" := ABS(#外呼上面有目标最大数3+#外呼上面有目标最大数3-#当前楼层-3)+#下行停站次数3+#上行停站次数10+#下行停站次数3+#上行停站次数10+2;
   END_IF;
   #"3层边沿触发8" := #_w9;
   #_w10 := #下呼灯3 AND #下行指示 AND (((3 = #当前楼层) AND NOT #上下平层都为1) OR (3 > #当前楼层));
   #_w11 := #_w10 AND #外呼上面有目标3;
   IF #_w11 THEN
       #"3层调度距离9" := ABS(#当前楼层-#外呼下面有目标最小数3+#外呼上面有目标最大数3-#外呼下面有目标最小数3+#外呼上面有目标最大数3-3)+#下行停站次数1+#下行停站次数3+#下行停站次数3+#下行停站次数1+#上行停站次数10+#上行停站次数10+4;
   END_IF;
   #"3层边沿触发9" := #_w11;
   #_w12 := #_w10 AND #外呼上面无目标3;
   IF #_w12 THEN
       #"3层调度距离10" := ABS(#当前楼层-#外呼下面有目标最小数3+3-#外呼下面有目标最小数3)+#下行停站次数1+#上行停站次数3+#上行停站次数3+#下行停站次数1+2;
   END_IF;
   #"3层边沿触发10" := #_w12;
   IF #"3层边沿触发1" AND (#载重量 <= #限重分配) AND NOT #检修中 AND NOT #死机 THEN #最终调度距离上3 := ABS(#"3层调度距离1"+0); END_IF;
   IF #"3层边沿触发1" AND (#载重量 > #限重分配) AND NOT #检修中 AND NOT #死机 THEN #最终调度距离上3 := ABS(#"3层调度距离1"+100); END_IF;
   IF #"3层边沿触发2" AND (#载重量 <= #限重分配) AND NOT #检修中 AND NOT #死机 THEN #最终调度距离上3 := ABS(#"3层调度距离2"+0); END_IF;
   IF #"3层边沿触发2" AND (#载重量 > #限重分配) AND NOT #检修中 AND NOT #死机 THEN #最终调度距离上3 := ABS(#"3层调度距离2"+100); END_IF;
   IF #"3层边沿触发3" AND (#载重量 <= #限重分配) AND NOT #检修中 AND NOT #死机 THEN #最终调度距离上3 := ABS(#"3层调度距离3"+0); END_IF;
   IF #"3层边沿触发3" AND (#载重量 > #限重分配) AND NOT #检修中 AND NOT #死机 THEN #最终调度距离上3 := ABS(#"3层调度距离3"+100); END_IF;
   IF #"3层边沿触发4" AND (#载重量 <= #限重分配) AND NOT #检修中 AND NOT #死机 THEN #最终调度距离上3 := ABS(#"3层调度距离4"+0); END_IF;
   IF #"3层边沿触发4" AND (#载重量 > #限重分配) AND NOT #检修中 AND NOT #死机 THEN #最终调度距离上3 := ABS(#"3层调度距离4"+100); END_IF;
   IF #"3层边沿触发5" AND (#载重量 <= #限重分配) AND NOT #检修中 AND NOT #死机 THEN #最终调度距离上3 := ABS(#"3层调度距离5"+0); END_IF;
   IF #"3层边沿触发5" AND (#载重量 > #限重分配) AND NOT #检修中 AND NOT #死机 THEN #最终调度距离上3 := ABS(#"3层调度距离5"+100); END_IF;
   IF #死机 OR #检修中 THEN #最终调度距离上3 := ABS(1000+1000); END_IF;
   IF #"3层边沿触发6" AND (#载重量 <= #限重分配) AND NOT #检修中 AND NOT #死机 THEN #最终调度距离下3 := ABS(#"3层调度距离6"+0); END_IF;
   IF #"3层边沿触发6" AND (#载重量 > #限重分配) AND NOT #检修中 AND NOT #死机 THEN #最终调度距离下3 := ABS(#"3层调度距离6"+100); END_IF;
   IF #"3层边沿触发7" AND (#载重量 <= #限重分配) AND NOT #检修中 AND NOT #死机 THEN #最终调度距离下3 := ABS(#"3层调度距离7"+0); END_IF;
   IF #"3层边沿触发7" AND (#载重量 > #限重分配) AND NOT #检修中 AND NOT #死机 THEN #最终调度距离下3 := ABS(#"3层调度距离7"+100); END_IF;
   IF #"3层边沿触发8" AND (#载重量 <= #限重分配) AND NOT #检修中 AND NOT #死机 THEN #最终调度距离下3 := ABS(#"3层调度距离8"+0); END_IF;
   IF #"3层边沿触发8" AND (#载重量 > #限重分配) AND NOT #检修中 AND NOT #死机 THEN #最终调度距离下3 := ABS(#"3层调度距离8"+100); END_IF;
   IF #"3层边沿触发9" AND (#载重量 <= #限重分配) AND NOT #检修中 AND NOT #死机 THEN #最终调度距离下3 := ABS(#"3层调度距离9"+0); END_IF;
   IF #"3层边沿触发9" AND (#载重量 > #限重分配) AND NOT #检修中 AND NOT #死机 THEN #最终调度距离下3 := ABS(#"3层调度距离9"+100); END_IF;
   IF #"3层边沿触发10" AND (#载重量 <= #限重分配) AND NOT #检修中 AND NOT #死机 THEN #最终调度距离下3 := ABS(#"3层调度距离10"+0); END_IF;
   IF #"3层边沿触发10" AND (#载重量 > #限重分配) AND NOT #检修中 AND NOT #死机 THEN #最终调度距离下3 := ABS(#"3层调度距离10"+100); END_IF;
   IF #死机 OR #检修中 THEN #最终调度距离下3 := ABS(1000+1000); END_IF;
END_REGION

REGION Network 3: 4层调度距离
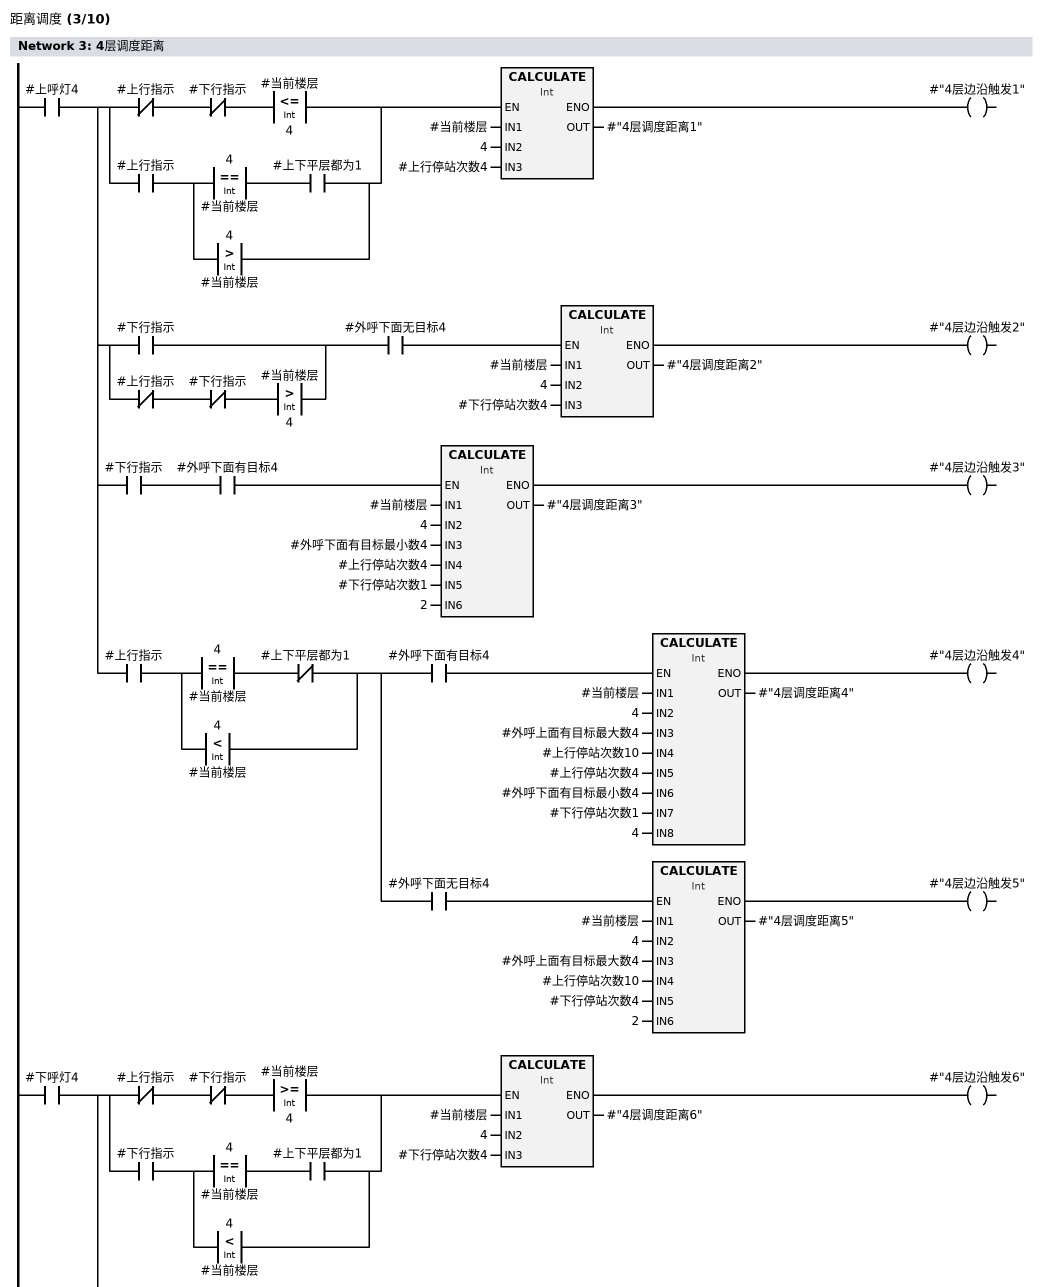
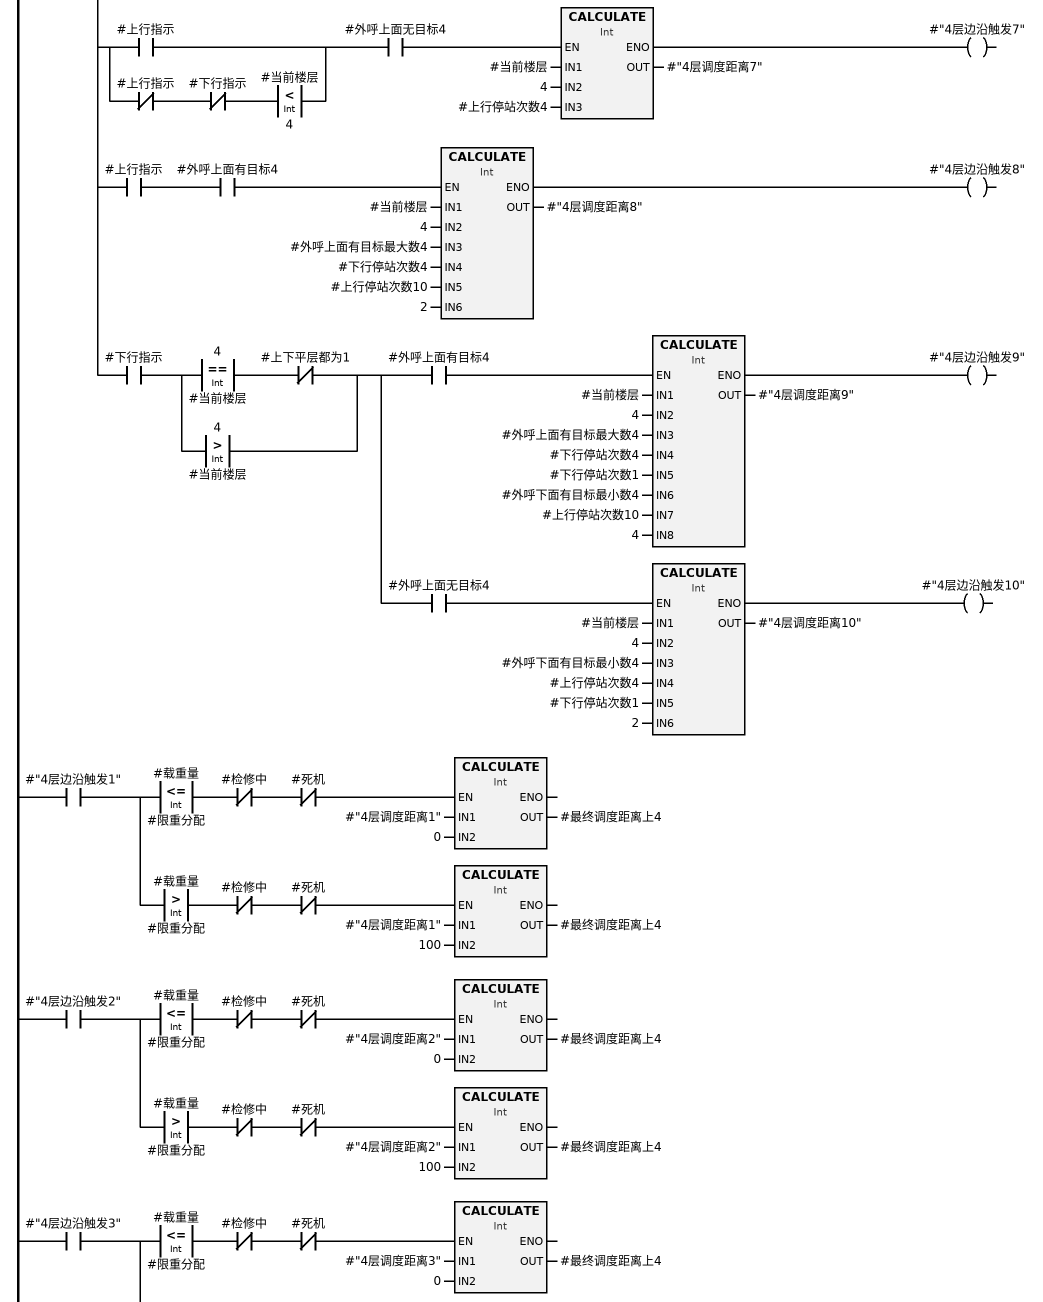
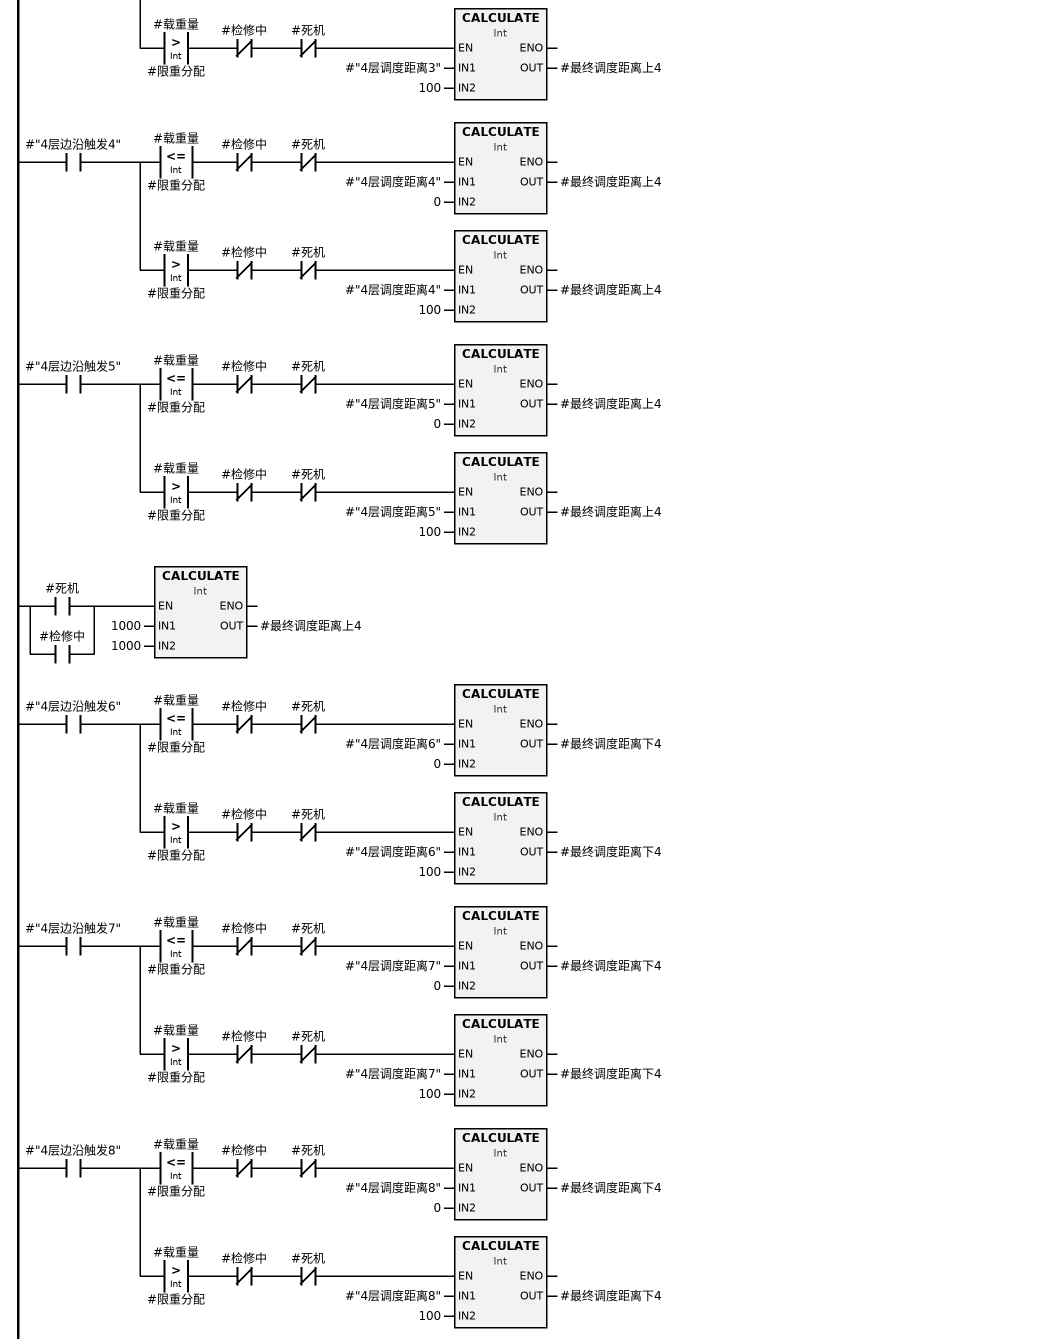
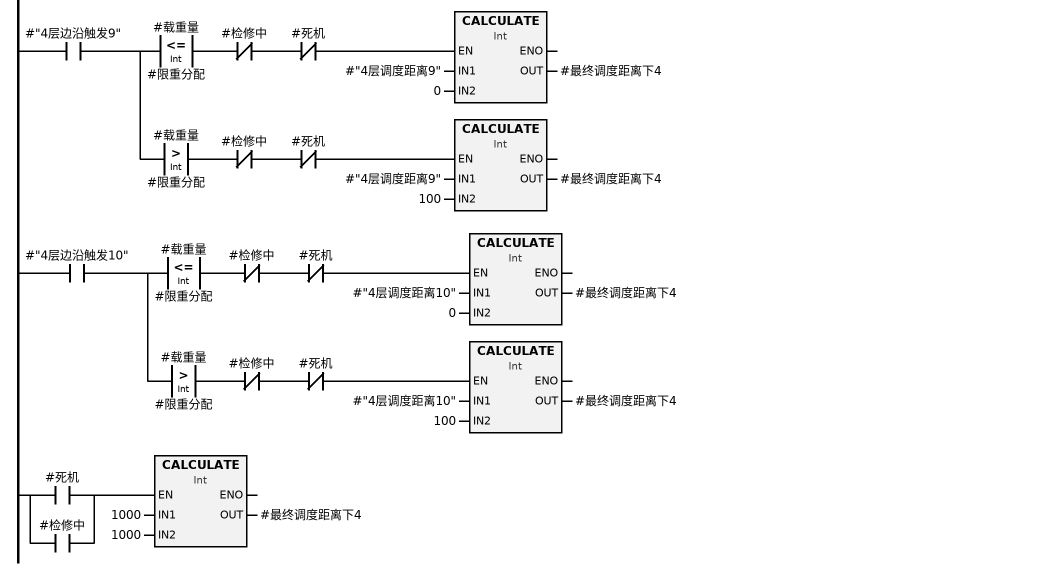
   RUNG wire#powerrail
      Contact( #上呼灯4 )
      wire#w1
      I_Contact( #上行指示 )
      I_Contact( #下行指示 )
      { S7_Templates := "SrcType := Int" } LE_Contact(in1 := #当前楼层, in2 := 4)
      wire#w2
      { S7_Templates := "SrcType := Int"; S7_Expression := "ABS(IN1-IN2)+IN3+IN3" } Calculate(in1 := #当前楼层, in2 := 4, in3 := #上行停站次数4, out => #"4层调度距离1")
      Coil( #"4层边沿触发1" )
   END_RUNG
   RUNG wire#w1
      Contact( #上行指示 )
      wire#w3
      { S7_Templates := "SrcType := Int" } EQ_Contact(in1 := 4, in2 := #当前楼层)
      Contact( #上下平层都为1 )
   END_RUNG wire#w2
   RUNG wire#w3
      { S7_Templates := "SrcType := Int" } GT_Contact(in1 := 4, in2 := #当前楼层)
   END_RUNG wire#w2
   RUNG wire#w1
      Contact( #下行指示 )
      wire#w4
      Contact( #外呼下面无目标4 )
      { S7_Templates := "SrcType := Int"; S7_Expression := "ABS(IN1-IN2)+IN3+IN3" } Calculate(in1 := #当前楼层, in2 := 4, in3 := #下行停站次数4, out => #"4层调度距离2")
      Coil( #"4层边沿触发2" )
   END_RUNG
   RUNG wire#w1
      I_Contact( #上行指示 )
      I_Contact( #下行指示 )
      { S7_Templates := "SrcType := Int" } GT_Contact(in1 := #当前楼层, in2 := 4)
   END_RUNG wire#w4
   RUNG wire#w1
      Contact( #下行指示 )
      Contact( #外呼下面有目标4 )
      { S7_Templates := "SrcType := Int"; S7_Expression := "ABS(IN3+IN3-IN1-IN2)+IN5+IN4+IN4+IN5+IN6" } Calculate(in1 := #当前楼层, in2 := 4, in3 := #外呼下面有目标最小数4, in4 := #上行停站次数4, in5 := #下行停站次数1, in6 := 2, out => #"4层调度距离3")
      Coil( #"4层边沿触发3" )
   END_RUNG
   RUNG wire#w1
      Contact( #上行指示 )
      wire#w5
      { S7_Templates := "SrcType := Int" } EQ_Contact(in1 := 4, in2 := #当前楼层)
      I_Contact( #上下平层都为1 )
      wire#w6
      Contact( #外呼下面有目标4 )
      { S7_Templates := "SrcType := Int"; S7_Expression := "ABS(IN3-IN1+IN3-IN6+IN2-IN6)+IN5+IN4+IN4+IN5+IN7+IN7+IN8" } Calculate(in1 := #当前楼层, in2 := 4, in3 := #外呼上面有目标最大数4, in4 := #上行停站次数10, in5 := #上行停站次数4, in6 := #外呼下面有目标最小数4, in7 := #下行停站次数1, in8 := 4, out => #"4层调度距离4")
      Coil( #"4层边沿触发4" )
   END_RUNG
   RUNG wire#w5
      { S7_Templates := "SrcType := Int" } LT_Contact(in1 := 4, in2 := #当前楼层)
   END_RUNG wire#w6
   RUNG wire#w6
      Contact( #外呼下面无目标4 )
      { S7_Templates := "SrcType := Int"; S7_Expression := "ABS(IN3-IN1+IN3-IN2)+IN5+IN4+IN4+IN5+IN6" } Calculate(in1 := #当前楼层, in2 := 4, in3 := #外呼上面有目标最大数4, in4 := #上行停站次数10, in5 := #下行停站次数4, in6 := 2, out => #"4层调度距离5")
      Coil( #"4层边沿触发5" )
   END_RUNG
   RUNG wire#powerrail
      Contact( #下呼灯4 )
      wire#w7
      I_Contact( #上行指示 )
      I_Contact( #下行指示 )
      { S7_Templates := "SrcType := Int" } GE_Contact(in1 := #当前楼层, in2 := 4)
      wire#w8
      { S7_Templates := "SrcType := Int"; S7_Expression := "ABS(IN1-IN2)+IN3+IN3" } Calculate(in1 := #当前楼层, in2 := 4, in3 := #下行停站次数4, out => #"4层调度距离6")
      Coil( #"4层边沿触发6" )
   END_RUNG
   RUNG wire#w7
      Contact( #下行指示 )
      wire#w9
      { S7_Templates := "SrcType := Int" } EQ_Contact(in1 := 4, in2 := #当前楼层)
      Contact( #上下平层都为1 )
   END_RUNG wire#w8
   RUNG wire#w9
      { S7_Templates := "SrcType := Int" } LT_Contact(in1 := 4, in2 := #当前楼层)
   END_RUNG wire#w8
   RUNG wire#w7
      Contact( #上行指示 )
      wire#w10
      Contact( #外呼上面无目标4 )
      { S7_Templates := "SrcType := Int"; S7_Expression := "ABS(IN1-IN2)+IN3+IN3" } Calculate(in1 := #当前楼层, in2 := 4, in3 := #上行停站次数4, out => #"4层调度距离7")
      Coil( #"4层边沿触发7" )
   END_RUNG
   RUNG wire#w7
      I_Contact( #上行指示 )
      I_Contact( #下行指示 )
      { S7_Templates := "SrcType := Int" } LT_Contact(in1 := #当前楼层, in2 := 4)
   END_RUNG wire#w10
   RUNG wire#w7
      Contact( #上行指示 )
      Contact( #外呼上面有目标4 )
      { S7_Templates := "SrcType := Int"; S7_Expression := "ABS(IN3+IN3-IN1-IN2)+IN4+IN5+IN4+IN5+IN6" } Calculate(in1 := #当前楼层, in2 := 4, in3 := #外呼上面有目标最大数4, in4 := #下行停站次数4, in5 := #上行停站次数10, in6 := 2, out => #"4层调度距离8")
      Coil( #"4层边沿触发8" )
   END_RUNG
   RUNG wire#w7
      Contact( #下行指示 )
      wire#w11
      { S7_Templates := "SrcType := Int" } EQ_Contact(in1 := 4, in2 := #当前楼层)
      I_Contact( #上下平层都为1 )
      wire#w12
      Contact( #外呼上面有目标4 )
      { S7_Templates := "SrcType := Int"; S7_Expression := "ABS(IN1-IN6+IN3-IN6+IN3-IN2)+IN5+IN4+IN4+IN5+IN7+IN7+IN8" } Calculate(in1 := #当前楼层, in2 := 4, in3 := #外呼上面有目标最大数4, in4 := #下行停站次数4, in5 := #下行停站次数1, in6 := #外呼下面有目标最小数4, in7 := #上行停站次数10, in8 := 4, out => #"4层调度距离9")
      Coil( #"4层边沿触发9" )
   END_RUNG
   RUNG wire#w11
      { S7_Templates := "SrcType := Int" } GT_Contact(in1 := 4, in2 := #当前楼层)
   END_RUNG wire#w12
   RUNG wire#w12
      Contact( #外呼上面无目标4 )
      { S7_Templates := "SrcType := Int"; S7_Expression := "ABS(IN1-IN3+IN2-IN3)+IN5+IN4+IN4+IN5+IN6" } Calculate(in1 := #当前楼层, in2 := 4, in3 := #外呼下面有目标最小数4, in4 := #上行停站次数4, in5 := #下行停站次数1, in6 := 2, out => #"4层调度距离10")
      Coil( #"4层边沿触发10" )
   END_RUNG
   RUNG wire#powerrail
      Contact( #"4层边沿触发1" )
      wire#w13
      { S7_Templates := "SrcType := Int" } LE_Contact(in1 := #载重量, in2 := #限重分配)
      I_Contact( #检修中 )
      I_Contact( #死机 )
      { S7_Templates := "SrcType := Int"; S7_Expression := "ABS(IN1+IN2)" } Calculate(in1 := #"4层调度距离1", in2 := 0, out => #最终调度距离上4)
   END_RUNG
   RUNG wire#w13
      { S7_Templates := "SrcType := Int" } GT_Contact(in1 := #载重量, in2 := #限重分配)
      I_Contact( #检修中 )
      I_Contact( #死机 )
      { S7_Templates := "SrcType := Int"; S7_Expression := "ABS(IN1+IN2)" } Calculate(in1 := #"4层调度距离1", in2 := 100, out => #最终调度距离上4)
   END_RUNG
   RUNG wire#powerrail
      Contact( #"4层边沿触发2" )
      wire#w14
      { S7_Templates := "SrcType := Int" } LE_Contact(in1 := #载重量, in2 := #限重分配)
      I_Contact( #检修中 )
      I_Contact( #死机 )
      { S7_Templates := "SrcType := Int"; S7_Expression := "ABS(IN1+IN2)" } Calculate(in1 := #"4层调度距离2", in2 := 0, out => #最终调度距离上4)
   END_RUNG
   RUNG wire#w14
      { S7_Templates := "SrcType := Int" } GT_Contact(in1 := #载重量, in2 := #限重分配)
      I_Contact( #检修中 )
      I_Contact( #死机 )
      { S7_Templates := "SrcType := Int"; S7_Expression := "ABS(IN1+IN2)" } Calculate(in1 := #"4层调度距离2", in2 := 100, out => #最终调度距离上4)
   END_RUNG
   RUNG wire#powerrail
      Contact( #"4层边沿触发3" )
      wire#w15
      { S7_Templates := "SrcType := Int" } LE_Contact(in1 := #载重量, in2 := #限重分配)
      I_Contact( #检修中 )
      I_Contact( #死机 )
      { S7_Templates := "SrcType := Int"; S7_Expression := "ABS(IN1+IN2)" } Calculate(in1 := #"4层调度距离3", in2 := 0, out => #最终调度距离上4)
   END_RUNG
   RUNG wire#w15
      { S7_Templates := "SrcType := Int" } GT_Contact(in1 := #载重量, in2 := #限重分配)
      I_Contact( #检修中 )
      I_Contact( #死机 )
      { S7_Templates := "SrcType := Int"; S7_Expression := "ABS(IN1+IN2)" } Calculate(in1 := #"4层调度距离3", in2 := 100, out => #最终调度距离上4)
   END_RUNG
   RUNG wire#powerrail
      Contact( #"4层边沿触发4" )
      wire#w16
      { S7_Templates := "SrcType := Int" } LE_Contact(in1 := #载重量, in2 := #限重分配)
      I_Contact( #检修中 )
      I_Contact( #死机 )
      { S7_Templates := "SrcType := Int"; S7_Expression := "ABS(IN1+IN2)" } Calculate(in1 := #"4层调度距离4", in2 := 0, out => #最终调度距离上4)
   END_RUNG
   RUNG wire#w16
      { S7_Templates := "SrcType := Int" } GT_Contact(in1 := #载重量, in2 := #限重分配)
      I_Contact( #检修中 )
      I_Contact( #死机 )
      { S7_Templates := "SrcType := Int"; S7_Expression := "ABS(IN1+IN2)" } Calculate(in1 := #"4层调度距离4", in2 := 100, out => #最终调度距离上4)
   END_RUNG
   RUNG wire#powerrail
      Contact( #"4层边沿触发5" )
      wire#w17
      { S7_Templates := "SrcType := Int" } LE_Contact(in1 := #载重量, in2 := #限重分配)
      I_Contact( #检修中 )
      I_Contact( #死机 )
      { S7_Templates := "SrcType := Int"; S7_Expression := "ABS(IN1+IN2)" } Calculate(in1 := #"4层调度距离5", in2 := 0, out => #最终调度距离上4)
   END_RUNG
   RUNG wire#w17
      { S7_Templates := "SrcType := Int" } GT_Contact(in1 := #载重量, in2 := #限重分配)
      I_Contact( #检修中 )
      I_Contact( #死机 )
      { S7_Templates := "SrcType := Int"; S7_Expression := "ABS(IN1+IN2)" } Calculate(in1 := #"4层调度距离5", in2 := 100, out => #最终调度距离上4)
   END_RUNG
   RUNG wire#powerrail
      Contact( #死机 )
      wire#w18
      { S7_Templates := "SrcType := Int"; S7_Expression := "ABS(IN1+IN2)" } Calculate(in1 := 1000, in2 := 1000, out => #最终调度距离上4)
   END_RUNG
   RUNG wire#powerrail
      Contact( #检修中 )
   END_RUNG wire#w18
   RUNG wire#powerrail
      Contact( #"4层边沿触发6" )
      wire#w19
      { S7_Templates := "SrcType := Int" } LE_Contact(in1 := #载重量, in2 := #限重分配)
      I_Contact( #检修中 )
      I_Contact( #死机 )
      { S7_Templates := "SrcType := Int"; S7_Expression := "ABS(IN1+IN2)" } Calculate(in1 := #"4层调度距离6", in2 := 0, out => #最终调度距离下4)
   END_RUNG
   RUNG wire#w19
      { S7_Templates := "SrcType := Int" } GT_Contact(in1 := #载重量, in2 := #限重分配)
      I_Contact( #检修中 )
      I_Contact( #死机 )
      { S7_Templates := "SrcType := Int"; S7_Expression := "ABS(IN1+IN2)" } Calculate(in1 := #"4层调度距离6", in2 := 100, out => #最终调度距离下4)
   END_RUNG
   RUNG wire#powerrail
      Contact( #"4层边沿触发7" )
      wire#w20
      { S7_Templates := "SrcType := Int" } LE_Contact(in1 := #载重量, in2 := #限重分配)
      I_Contact( #检修中 )
      I_Contact( #死机 )
      { S7_Templates := "SrcType := Int"; S7_Expression := "ABS(IN1+IN2)" } Calculate(in1 := #"4层调度距离7", in2 := 0, out => #最终调度距离下4)
   END_RUNG
   RUNG wire#w20
      { S7_Templates := "SrcType := Int" } GT_Contact(in1 := #载重量, in2 := #限重分配)
      I_Contact( #检修中 )
      I_Contact( #死机 )
      { S7_Templates := "SrcType := Int"; S7_Expression := "ABS(IN1+IN2)" } Calculate(in1 := #"4层调度距离7", in2 := 100, out => #最终调度距离下4)
   END_RUNG
   RUNG wire#powerrail
      Contact( #"4层边沿触发8" )
      wire#w21
      { S7_Templates := "SrcType := Int" } LE_Contact(in1 := #载重量, in2 := #限重分配)
      I_Contact( #检修中 )
      I_Contact( #死机 )
      { S7_Templates := "SrcType := Int"; S7_Expression := "ABS(IN1+IN2)" } Calculate(in1 := #"4层调度距离8", in2 := 0, out => #最终调度距离下4)
   END_RUNG
   RUNG wire#w21
      { S7_Templates := "SrcType := Int" } GT_Contact(in1 := #载重量, in2 := #限重分配)
      I_Contact( #检修中 )
      I_Contact( #死机 )
      { S7_Templates := "SrcType := Int"; S7_Expression := "ABS(IN1+IN2)" } Calculate(in1 := #"4层调度距离8", in2 := 100, out => #最终调度距离下4)
   END_RUNG
   RUNG wire#powerrail
      Contact( #"4层边沿触发9" )
      wire#w22
      { S7_Templates := "SrcType := Int" } LE_Contact(in1 := #载重量, in2 := #限重分配)
      I_Contact( #检修中 )
      I_Contact( #死机 )
      { S7_Templates := "SrcType := Int"; S7_Expression := "ABS(IN1+IN2)" } Calculate(in1 := #"4层调度距离9", in2 := 0, out => #最终调度距离下4)
   END_RUNG
   RUNG wire#w22
      { S7_Templates := "SrcType := Int" } GT_Contact(in1 := #载重量, in2 := #限重分配)
      I_Contact( #检修中 )
      I_Contact( #死机 )
      { S7_Templates := "SrcType := Int"; S7_Expression := "ABS(IN1+IN2)" } Calculate(in1 := #"4层调度距离9", in2 := 100, out => #最终调度距离下4)
   END_RUNG
   RUNG wire#powerrail
      Contact( #"4层边沿触发10" )
      wire#w23
      { S7_Templates := "SrcType := Int" } LE_Contact(in1 := #载重量, in2 := #限重分配)
      I_Contact( #检修中 )
      I_Contact( #死机 )
      { S7_Templates := "SrcType := Int"; S7_Expression := "ABS(IN1+IN2)" } Calculate(in1 := #"4层调度距离10", in2 := 0, out => #最终调度距离下4)
   END_RUNG
   RUNG wire#w23
      { S7_Templates := "SrcType := Int" } GT_Contact(in1 := #载重量, in2 := #限重分配)
      I_Contact( #检修中 )
      I_Contact( #死机 )
      { S7_Templates := "SrcType := Int"; S7_Expression := "ABS(IN1+IN2)" } Calculate(in1 := #"4层调度距离10", in2 := 100, out => #最终调度距离下4)
   END_RUNG
   RUNG wire#powerrail
      Contact( #死机 )
      wire#w24
      { S7_Templates := "SrcType := Int"; S7_Expression := "ABS(IN1+IN2)" } Calculate(in1 := 1000, in2 := 1000, out => #最终调度距离下4)
   END_RUNG
   RUNG wire#powerrail
      Contact( #检修中 )
   END_RUNG wire#w24
   // the same network as SCL:
   #_w1 := #上呼灯4 AND ((NOT #上行指示 AND NOT #下行指示 AND (#当前楼层 <= 4)) OR (#上行指示 AND (((4 = #当前楼层) AND #上下平层都为1) OR (4 > #当前楼层))));
   IF #_w1 THEN #"4层调度距离1" := ABS(#当前楼层-4)+#上行停站次数4+#上行停站次数4; END_IF;
   #"4层边沿触发1" := #_w1;
   #_w2 := #上呼灯4 AND (#下行指示 OR (NOT #上行指示 AND NOT #下行指示 AND (#当前楼层 > 4))) AND #外呼下面无目标4;
   IF #_w2 THEN #"4层调度距离2" := ABS(#当前楼层-4)+#下行停站次数4+#下行停站次数4; END_IF;
   #"4层边沿触发2" := #_w2;
   #_w3 := #上呼灯4 AND #下行指示 AND #外呼下面有目标4;
   IF #_w3 THEN
       #"4层调度距离3" := ABS(#外呼下面有目标最小数4+#外呼下面有目标最小数4-#当前楼层-4)+#下行停站次数1+#上行停站次数4+#上行停站次数4+#下行停站次数1+2;
   END_IF;
   #"4层边沿触发3" := #_w3;
   #_w4 := #上呼灯4 AND #上行指示 AND (((4 = #当前楼层) AND NOT #上下平层都为1) OR (4 < #当前楼层));
   #_w5 := #_w4 AND #外呼下面有目标4;
   IF #_w5 THEN
       #"4层调度距离4" := ABS(#外呼上面有目标最大数4-#当前楼层+#外呼上面有目标最大数4-#外呼下面有目标最小数4+4-#外呼下面有目标最小数4)+#上行停站次数4+#上行停站次数10+#上行停站次数10+#上行停站次数4+#下行停站次数1+#下行停站次数1+4;
   END_IF;
   #"4层边沿触发4" := #_w5;
   #_w6 := #_w4 AND #外呼下面无目标4;
   IF #_w6 THEN
       #"4层调度距离5" := ABS(#外呼上面有目标最大数4-#当前楼层+#外呼上面有目标最大数4-4)+#下行停站次数4+#上行停站次数10+#上行停站次数10+#下行停站次数4+2;
   END_IF;
   #"4层边沿触发5" := #_w6;
   #_w7 := #下呼灯4 AND ((NOT #上行指示 AND NOT #下行指示 AND (#当前楼层 >= 4)) OR (#下行指示 AND (((4 = #当前楼层) AND #上下平层都为1) OR (4 < #当前楼层))));
   IF #_w7 THEN #"4层调度距离6" := ABS(#当前楼层-4)+#下行停站次数4+#下行停站次数4; END_IF;
   #"4层边沿触发6" := #_w7;
   #_w8 := #下呼灯4 AND (#上行指示 OR (NOT #上行指示 AND NOT #下行指示 AND (#当前楼层 < 4))) AND #外呼上面无目标4;
   IF #_w8 THEN #"4层调度距离7" := ABS(#当前楼层-4)+#上行停站次数4+#上行停站次数4; END_IF;
   #"4层边沿触发7" := #_w8;
   #_w9 := #下呼灯4 AND #上行指示 AND #外呼上面有目标4;
   IF #_w9 THEN
       #"4层调度距离8" := ABS(#外呼上面有目标最大数4+#外呼上面有目标最大数4-#当前楼层-4)+#下行停站次数4+#上行停站次数10+#下行停站次数4+#上行停站次数10+2;
   END_IF;
   #"4层边沿触发8" := #_w9;
   #_w10 := #下呼灯4 AND #下行指示 AND (((4 = #当前楼层) AND NOT #上下平层都为1) OR (4 > #当前楼层));
   #_w11 := #_w10 AND #外呼上面有目标4;
   IF #_w11 THEN
       #"4层调度距离9" := ABS(#当前楼层-#外呼下面有目标最小数4+#外呼上面有目标最大数4-#外呼下面有目标最小数4+#外呼上面有目标最大数4-4)+#下行停站次数1+#下行停站次数4+#下行停站次数4+#下行停站次数1+#上行停站次数10+#上行停站次数10+4;
   END_IF;
   #"4层边沿触发9" := #_w11;
   #_w12 := #_w10 AND #外呼上面无目标4;
   IF #_w12 THEN
       #"4层调度距离10" := ABS(#当前楼层-#外呼下面有目标最小数4+4-#外呼下面有目标最小数4)+#下行停站次数1+#上行停站次数4+#上行停站次数4+#下行停站次数1+2;
   END_IF;
   #"4层边沿触发10" := #_w12;
   IF #"4层边沿触发1" AND (#载重量 <= #限重分配) AND NOT #检修中 AND NOT #死机 THEN #最终调度距离上4 := ABS(#"4层调度距离1"+0); END_IF;
   IF #"4层边沿触发1" AND (#载重量 > #限重分配) AND NOT #检修中 AND NOT #死机 THEN #最终调度距离上4 := ABS(#"4层调度距离1"+100); END_IF;
   IF #"4层边沿触发2" AND (#载重量 <= #限重分配) AND NOT #检修中 AND NOT #死机 THEN #最终调度距离上4 := ABS(#"4层调度距离2"+0); END_IF;
   IF #"4层边沿触发2" AND (#载重量 > #限重分配) AND NOT #检修中 AND NOT #死机 THEN #最终调度距离上4 := ABS(#"4层调度距离2"+100); END_IF;
   IF #"4层边沿触发3" AND (#载重量 <= #限重分配) AND NOT #检修中 AND NOT #死机 THEN #最终调度距离上4 := ABS(#"4层调度距离3"+0); END_IF;
   IF #"4层边沿触发3" AND (#载重量 > #限重分配) AND NOT #检修中 AND NOT #死机 THEN #最终调度距离上4 := ABS(#"4层调度距离3"+100); END_IF;
   IF #"4层边沿触发4" AND (#载重量 <= #限重分配) AND NOT #检修中 AND NOT #死机 THEN #最终调度距离上4 := ABS(#"4层调度距离4"+0); END_IF;
   IF #"4层边沿触发4" AND (#载重量 > #限重分配) AND NOT #检修中 AND NOT #死机 THEN #最终调度距离上4 := ABS(#"4层调度距离4"+100); END_IF;
   IF #"4层边沿触发5" AND (#载重量 <= #限重分配) AND NOT #检修中 AND NOT #死机 THEN #最终调度距离上4 := ABS(#"4层调度距离5"+0); END_IF;
   IF #"4层边沿触发5" AND (#载重量 > #限重分配) AND NOT #检修中 AND NOT #死机 THEN #最终调度距离上4 := ABS(#"4层调度距离5"+100); END_IF;
   IF #死机 OR #检修中 THEN #最终调度距离上4 := ABS(1000+1000); END_IF;
   IF #"4层边沿触发6" AND (#载重量 <= #限重分配) AND NOT #检修中 AND NOT #死机 THEN #最终调度距离下4 := ABS(#"4层调度距离6"+0); END_IF;
   IF #"4层边沿触发6" AND (#载重量 > #限重分配) AND NOT #检修中 AND NOT #死机 THEN #最终调度距离下4 := ABS(#"4层调度距离6"+100); END_IF;
   IF #"4层边沿触发7" AND (#载重量 <= #限重分配) AND NOT #检修中 AND NOT #死机 THEN #最终调度距离下4 := ABS(#"4层调度距离7"+0); END_IF;
   IF #"4层边沿触发7" AND (#载重量 > #限重分配) AND NOT #检修中 AND NOT #死机 THEN #最终调度距离下4 := ABS(#"4层调度距离7"+100); END_IF;
   IF #"4层边沿触发8" AND (#载重量 <= #限重分配) AND NOT #检修中 AND NOT #死机 THEN #最终调度距离下4 := ABS(#"4层调度距离8"+0); END_IF;
   IF #"4层边沿触发8" AND (#载重量 > #限重分配) AND NOT #检修中 AND NOT #死机 THEN #最终调度距离下4 := ABS(#"4层调度距离8"+100); END_IF;
   IF #"4层边沿触发9" AND (#载重量 <= #限重分配) AND NOT #检修中 AND NOT #死机 THEN #最终调度距离下4 := ABS(#"4层调度距离9"+0); END_IF;
   IF #"4层边沿触发9" AND (#载重量 > #限重分配) AND NOT #检修中 AND NOT #死机 THEN #最终调度距离下4 := ABS(#"4层调度距离9"+100); END_IF;
   IF #"4层边沿触发10" AND (#载重量 <= #限重分配) AND NOT #检修中 AND NOT #死机 THEN #最终调度距离下4 := ABS(#"4层调度距离10"+0); END_IF;
   IF #"4层边沿触发10" AND (#载重量 > #限重分配) AND NOT #检修中 AND NOT #死机 THEN #最终调度距离下4 := ABS(#"4层调度距离10"+100); END_IF;
   IF #死机 OR #检修中 THEN #最终调度距离下4 := ABS(1000+1000); END_IF;
END_REGION

REGION Network 4: 5层调度距离
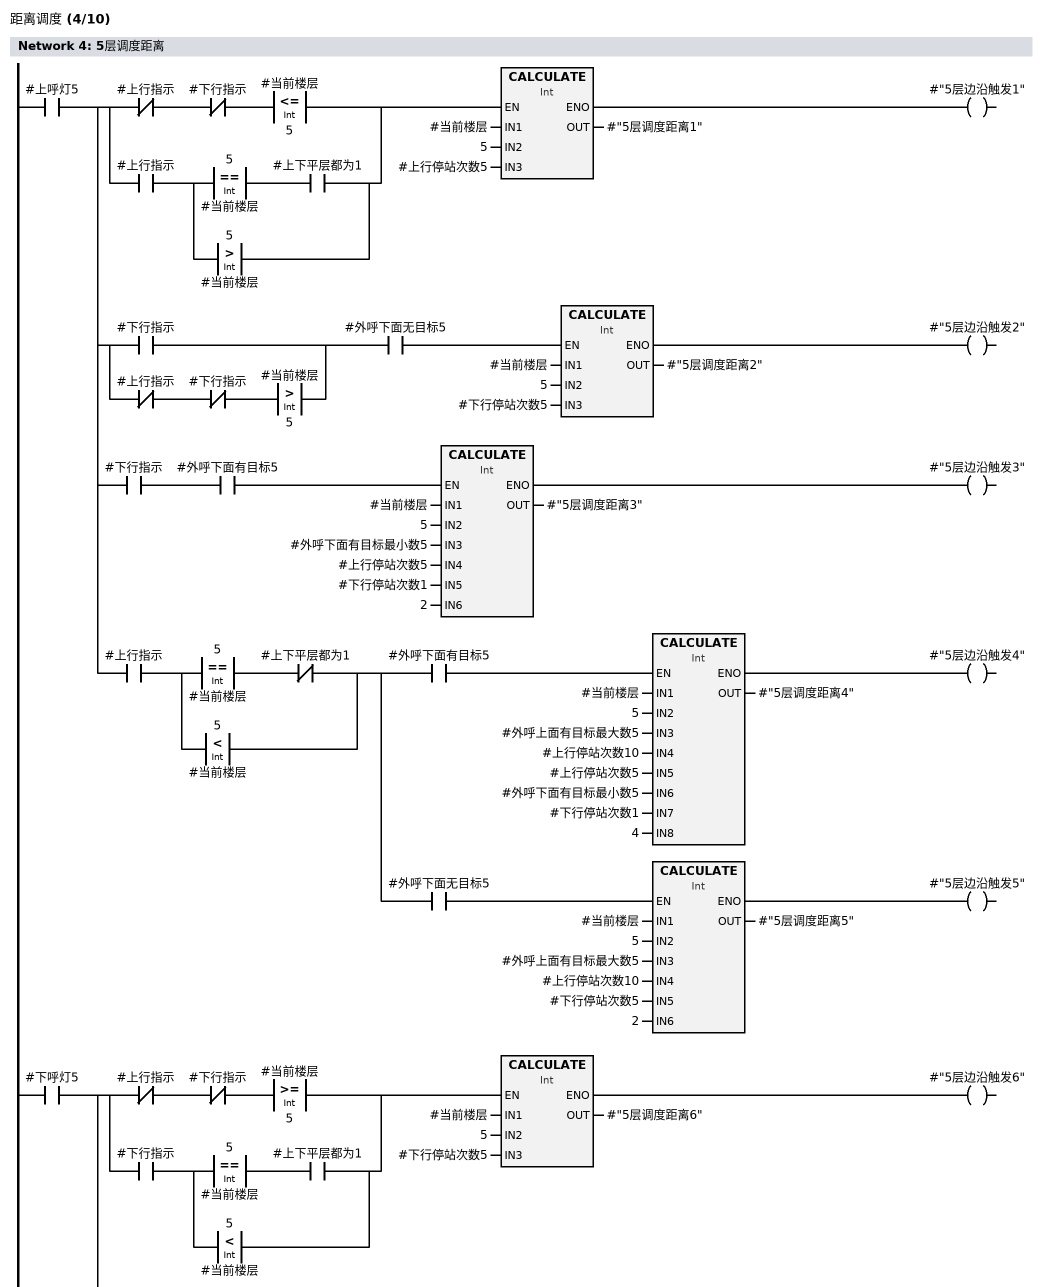
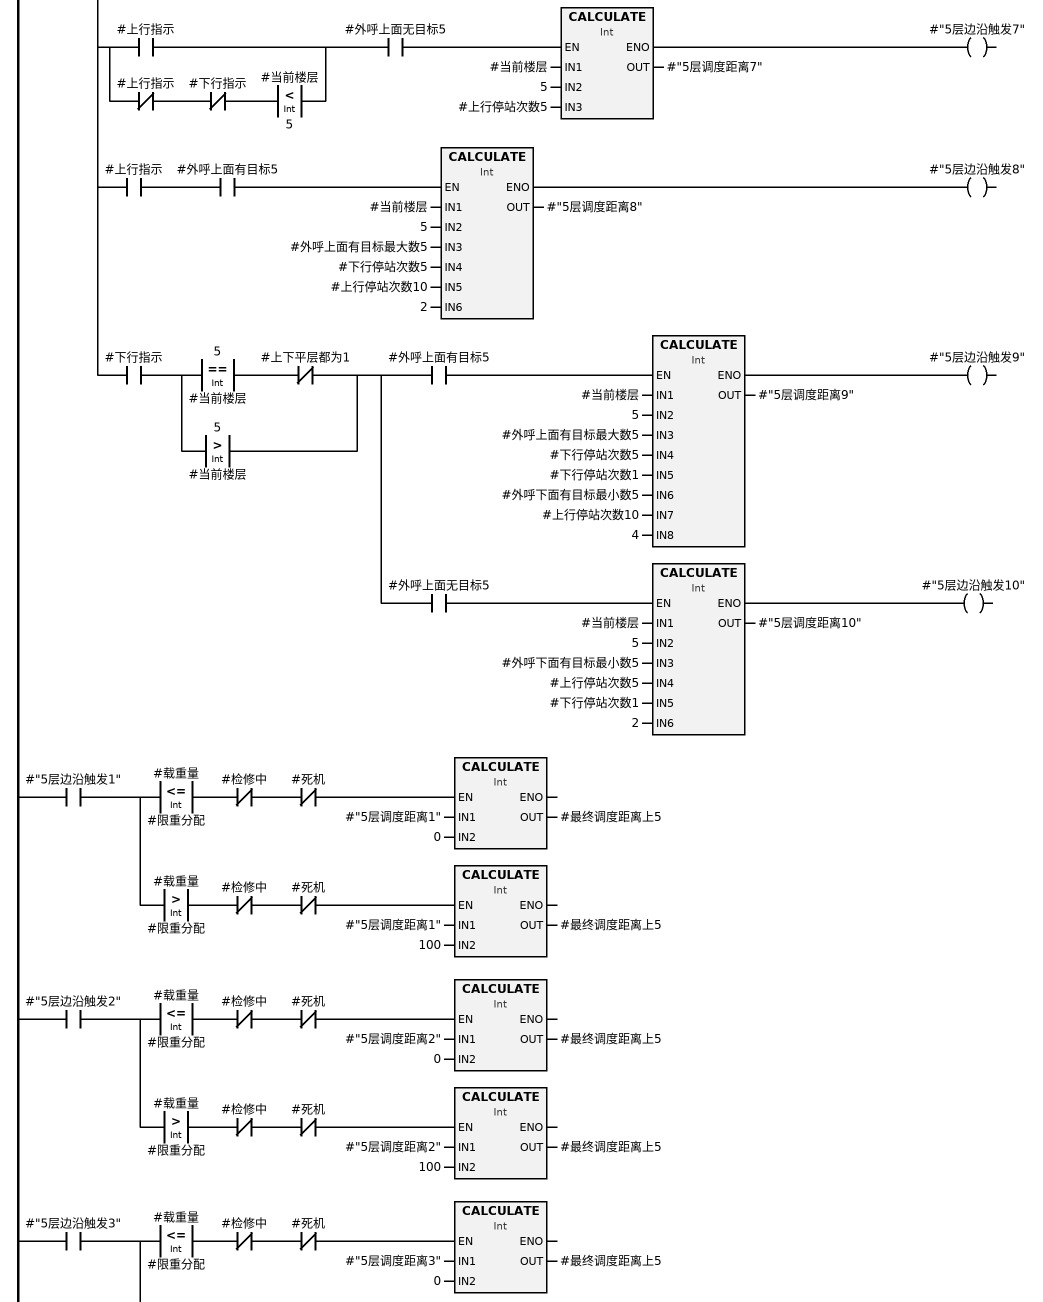
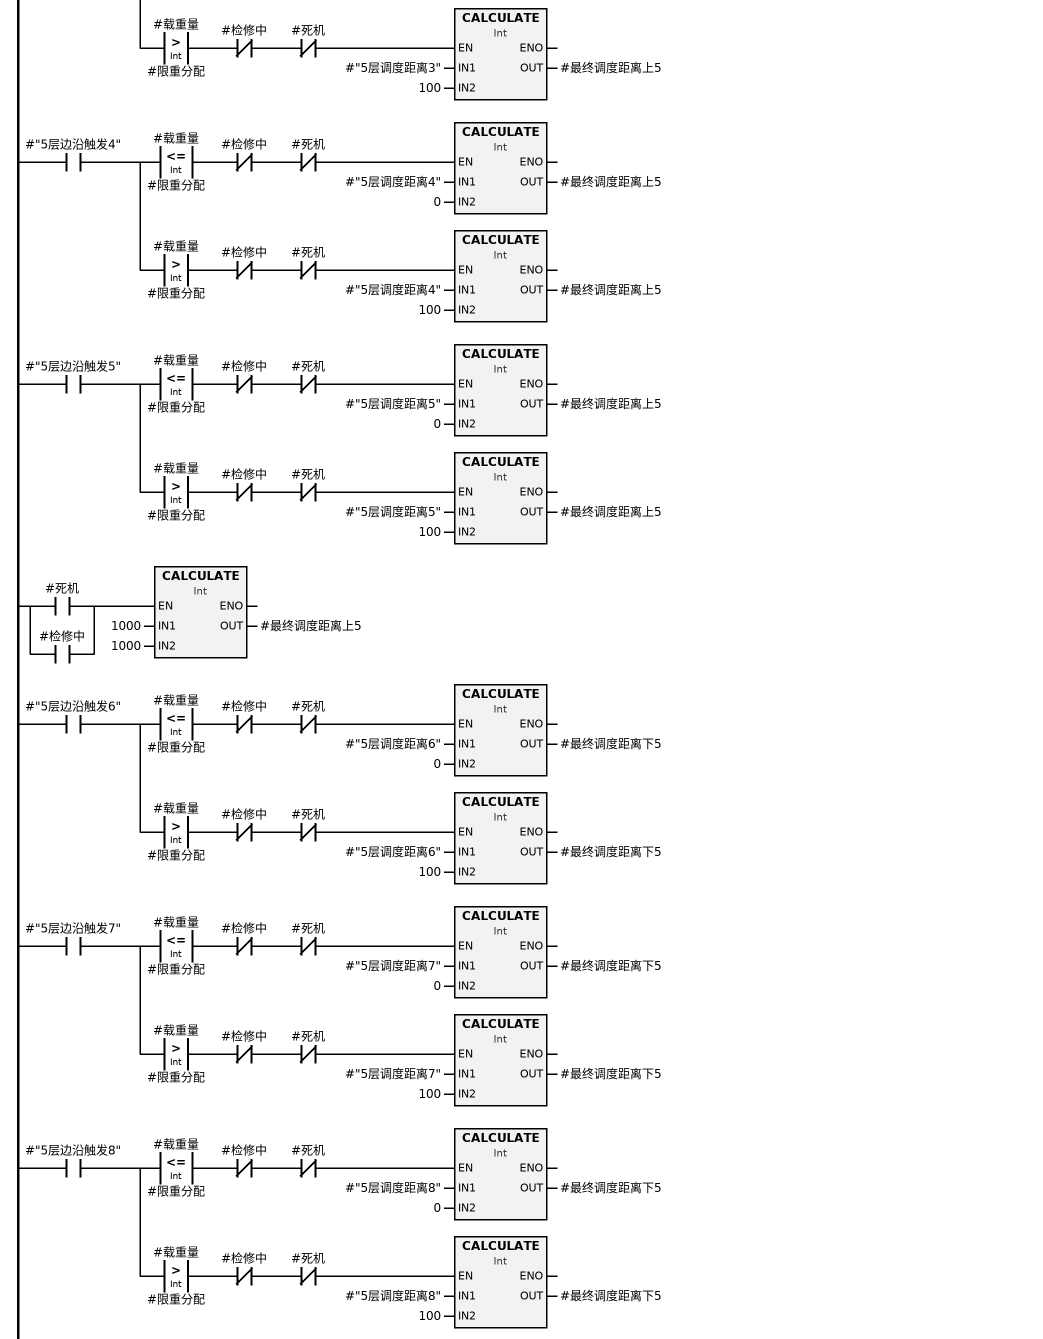
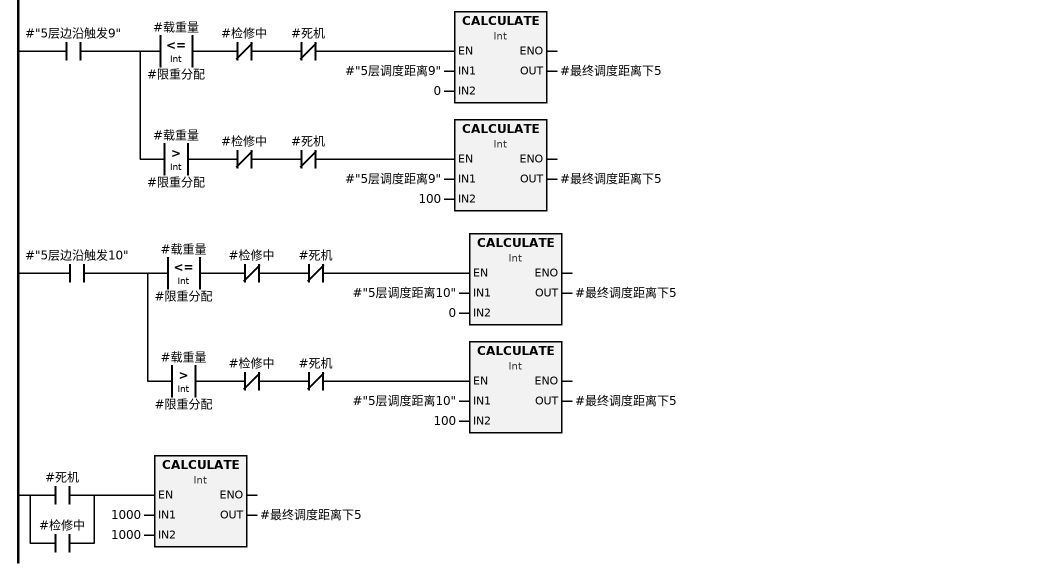
   RUNG wire#powerrail
      Contact( #上呼灯5 )
      wire#w1
      I_Contact( #上行指示 )
      I_Contact( #下行指示 )
      { S7_Templates := "SrcType := Int" } LE_Contact(in1 := #当前楼层, in2 := 5)
      wire#w2
      { S7_Templates := "SrcType := Int"; S7_Expression := "ABS(IN1-IN2)+IN3+IN3" } Calculate(in1 := #当前楼层, in2 := 5, in3 := #上行停站次数5, out => #"5层调度距离1")
      Coil( #"5层边沿触发1" )
   END_RUNG
   RUNG wire#w1
      Contact( #上行指示 )
      wire#w3
      { S7_Templates := "SrcType := Int" } EQ_Contact(in1 := 5, in2 := #当前楼层)
      Contact( #上下平层都为1 )
   END_RUNG wire#w2
   RUNG wire#w3
      { S7_Templates := "SrcType := Int" } GT_Contact(in1 := 5, in2 := #当前楼层)
   END_RUNG wire#w2
   RUNG wire#w1
      Contact( #下行指示 )
      wire#w4
      Contact( #外呼下面无目标5 )
      { S7_Templates := "SrcType := Int"; S7_Expression := "ABS(IN1-IN2)+IN3+IN3" } Calculate(in1 := #当前楼层, in2 := 5, in3 := #下行停站次数5, out => #"5层调度距离2")
      Coil( #"5层边沿触发2" )
   END_RUNG
   RUNG wire#w1
      I_Contact( #上行指示 )
      I_Contact( #下行指示 )
      { S7_Templates := "SrcType := Int" } GT_Contact(in1 := #当前楼层, in2 := 5)
   END_RUNG wire#w4
   RUNG wire#w1
      Contact( #下行指示 )
      Contact( #外呼下面有目标5 )
      { S7_Templates := "SrcType := Int"; S7_Expression := "ABS(IN3+IN3-IN1-IN2)+IN5+IN4+IN4+IN5+IN6" } Calculate(in1 := #当前楼层, in2 := 5, in3 := #外呼下面有目标最小数5, in4 := #上行停站次数5, in5 := #下行停站次数1, in6 := 2, out => #"5层调度距离3")
      Coil( #"5层边沿触发3" )
   END_RUNG
   RUNG wire#w1
      Contact( #上行指示 )
      wire#w5
      { S7_Templates := "SrcType := Int" } EQ_Contact(in1 := 5, in2 := #当前楼层)
      I_Contact( #上下平层都为1 )
      wire#w6
      Contact( #外呼下面有目标5 )
      { S7_Templates := "SrcType := Int"; S7_Expression := "ABS(IN3-IN1+IN3-IN6+IN2-IN6)+IN5+IN4+IN4+IN5+IN7+IN7+IN8" } Calculate(in1 := #当前楼层, in2 := 5, in3 := #外呼上面有目标最大数5, in4 := #上行停站次数10, in5 := #上行停站次数5, in6 := #外呼下面有目标最小数5, in7 := #下行停站次数1, in8 := 4, out => #"5层调度距离4")
      Coil( #"5层边沿触发4" )
   END_RUNG
   RUNG wire#w5
      { S7_Templates := "SrcType := Int" } LT_Contact(in1 := 5, in2 := #当前楼层)
   END_RUNG wire#w6
   RUNG wire#w6
      Contact( #外呼下面无目标5 )
      { S7_Templates := "SrcType := Int"; S7_Expression := "ABS(IN3-IN1+IN3-IN2)+IN5+IN4+IN4+IN5+IN6" } Calculate(in1 := #当前楼层, in2 := 5, in3 := #外呼上面有目标最大数5, in4 := #上行停站次数10, in5 := #下行停站次数5, in6 := 2, out => #"5层调度距离5")
      Coil( #"5层边沿触发5" )
   END_RUNG
   RUNG wire#powerrail
      Contact( #下呼灯5 )
      wire#w7
      I_Contact( #上行指示 )
      I_Contact( #下行指示 )
      { S7_Templates := "SrcType := Int" } GE_Contact(in1 := #当前楼层, in2 := 5)
      wire#w8
      { S7_Templates := "SrcType := Int"; S7_Expression := "ABS(IN1-IN2)+IN3+IN3" } Calculate(in1 := #当前楼层, in2 := 5, in3 := #下行停站次数5, out => #"5层调度距离6")
      Coil( #"5层边沿触发6" )
   END_RUNG
   RUNG wire#w7
      Contact( #下行指示 )
      wire#w9
      { S7_Templates := "SrcType := Int" } EQ_Contact(in1 := 5, in2 := #当前楼层)
      Contact( #上下平层都为1 )
   END_RUNG wire#w8
   RUNG wire#w9
      { S7_Templates := "SrcType := Int" } LT_Contact(in1 := 5, in2 := #当前楼层)
   END_RUNG wire#w8
   RUNG wire#w7
      Contact( #上行指示 )
      wire#w10
      Contact( #外呼上面无目标5 )
      { S7_Templates := "SrcType := Int"; S7_Expression := "ABS(IN1-IN2)+IN3+IN3" } Calculate(in1 := #当前楼层, in2 := 5, in3 := #上行停站次数5, out => #"5层调度距离7")
      Coil( #"5层边沿触发7" )
   END_RUNG
   RUNG wire#w7
      I_Contact( #上行指示 )
      I_Contact( #下行指示 )
      { S7_Templates := "SrcType := Int" } LT_Contact(in1 := #当前楼层, in2 := 5)
   END_RUNG wire#w10
   RUNG wire#w7
      Contact( #上行指示 )
      Contact( #外呼上面有目标5 )
      { S7_Templates := "SrcType := Int"; S7_Expression := "ABS(IN3+IN3-IN1-IN2)+IN4+IN5+IN4+IN5+IN6" } Calculate(in1 := #当前楼层, in2 := 5, in3 := #外呼上面有目标最大数5, in4 := #下行停站次数5, in5 := #上行停站次数10, in6 := 2, out => #"5层调度距离8")
      Coil( #"5层边沿触发8" )
   END_RUNG
   RUNG wire#w7
      Contact( #下行指示 )
      wire#w11
      { S7_Templates := "SrcType := Int" } EQ_Contact(in1 := 5, in2 := #当前楼层)
      I_Contact( #上下平层都为1 )
      wire#w12
      Contact( #外呼上面有目标5 )
      { S7_Templates := "SrcType := Int"; S7_Expression := "ABS(IN1-IN6+IN3-IN6+IN3-IN2)+IN5+IN4+IN4+IN5+IN7+IN7+IN8" } Calculate(in1 := #当前楼层, in2 := 5, in3 := #外呼上面有目标最大数5, in4 := #下行停站次数5, in5 := #下行停站次数1, in6 := #外呼下面有目标最小数5, in7 := #上行停站次数10, in8 := 4, out => #"5层调度距离9")
      Coil( #"5层边沿触发9" )
   END_RUNG
   RUNG wire#w11
      { S7_Templates := "SrcType := Int" } GT_Contact(in1 := 5, in2 := #当前楼层)
   END_RUNG wire#w12
   RUNG wire#w12
      Contact( #外呼上面无目标5 )
      { S7_Templates := "SrcType := Int"; S7_Expression := "ABS(IN1-IN3+IN2-IN3)+IN5+IN4+IN4+IN5+IN6" } Calculate(in1 := #当前楼层, in2 := 5, in3 := #外呼下面有目标最小数5, in4 := #上行停站次数5, in5 := #下行停站次数1, in6 := 2, out => #"5层调度距离10")
      Coil( #"5层边沿触发10" )
   END_RUNG
   RUNG wire#powerrail
      Contact( #"5层边沿触发1" )
      wire#w13
      { S7_Templates := "SrcType := Int" } LE_Contact(in1 := #载重量, in2 := #限重分配)
      I_Contact( #检修中 )
      I_Contact( #死机 )
      { S7_Templates := "SrcType := Int"; S7_Expression := "ABS(IN1+IN2)" } Calculate(in1 := #"5层调度距离1", in2 := 0, out => #最终调度距离上5)
   END_RUNG
   RUNG wire#w13
      { S7_Templates := "SrcType := Int" } GT_Contact(in1 := #载重量, in2 := #限重分配)
      I_Contact( #检修中 )
      I_Contact( #死机 )
      { S7_Templates := "SrcType := Int"; S7_Expression := "ABS(IN1+IN2)" } Calculate(in1 := #"5层调度距离1", in2 := 100, out => #最终调度距离上5)
   END_RUNG
   RUNG wire#powerrail
      Contact( #"5层边沿触发2" )
      wire#w14
      { S7_Templates := "SrcType := Int" } LE_Contact(in1 := #载重量, in2 := #限重分配)
      I_Contact( #检修中 )
      I_Contact( #死机 )
      { S7_Templates := "SrcType := Int"; S7_Expression := "ABS(IN1+IN2)" } Calculate(in1 := #"5层调度距离2", in2 := 0, out => #最终调度距离上5)
   END_RUNG
   RUNG wire#w14
      { S7_Templates := "SrcType := Int" } GT_Contact(in1 := #载重量, in2 := #限重分配)
      I_Contact( #检修中 )
      I_Contact( #死机 )
      { S7_Templates := "SrcType := Int"; S7_Expression := "ABS(IN1+IN2)" } Calculate(in1 := #"5层调度距离2", in2 := 100, out => #最终调度距离上5)
   END_RUNG
   RUNG wire#powerrail
      Contact( #"5层边沿触发3" )
      wire#w15
      { S7_Templates := "SrcType := Int" } LE_Contact(in1 := #载重量, in2 := #限重分配)
      I_Contact( #检修中 )
      I_Contact( #死机 )
      { S7_Templates := "SrcType := Int"; S7_Expression := "ABS(IN1+IN2)" } Calculate(in1 := #"5层调度距离3", in2 := 0, out => #最终调度距离上5)
   END_RUNG
   RUNG wire#w15
      { S7_Templates := "SrcType := Int" } GT_Contact(in1 := #载重量, in2 := #限重分配)
      I_Contact( #检修中 )
      I_Contact( #死机 )
      { S7_Templates := "SrcType := Int"; S7_Expression := "ABS(IN1+IN2)" } Calculate(in1 := #"5层调度距离3", in2 := 100, out => #最终调度距离上5)
   END_RUNG
   RUNG wire#powerrail
      Contact( #"5层边沿触发4" )
      wire#w16
      { S7_Templates := "SrcType := Int" } LE_Contact(in1 := #载重量, in2 := #限重分配)
      I_Contact( #检修中 )
      I_Contact( #死机 )
      { S7_Templates := "SrcType := Int"; S7_Expression := "ABS(IN1+IN2)" } Calculate(in1 := #"5层调度距离4", in2 := 0, out => #最终调度距离上5)
   END_RUNG
   RUNG wire#w16
      { S7_Templates := "SrcType := Int" } GT_Contact(in1 := #载重量, in2 := #限重分配)
      I_Contact( #检修中 )
      I_Contact( #死机 )
      { S7_Templates := "SrcType := Int"; S7_Expression := "ABS(IN1+IN2)" } Calculate(in1 := #"5层调度距离4", in2 := 100, out => #最终调度距离上5)
   END_RUNG
   RUNG wire#powerrail
      Contact( #"5层边沿触发5" )
      wire#w17
      { S7_Templates := "SrcType := Int" } LE_Contact(in1 := #载重量, in2 := #限重分配)
      I_Contact( #检修中 )
      I_Contact( #死机 )
      { S7_Templates := "SrcType := Int"; S7_Expression := "ABS(IN1+IN2)" } Calculate(in1 := #"5层调度距离5", in2 := 0, out => #最终调度距离上5)
   END_RUNG
   RUNG wire#w17
      { S7_Templates := "SrcType := Int" } GT_Contact(in1 := #载重量, in2 := #限重分配)
      I_Contact( #检修中 )
      I_Contact( #死机 )
      { S7_Templates := "SrcType := Int"; S7_Expression := "ABS(IN1+IN2)" } Calculate(in1 := #"5层调度距离5", in2 := 100, out => #最终调度距离上5)
   END_RUNG
   RUNG wire#powerrail
      Contact( #死机 )
      wire#w18
      { S7_Templates := "SrcType := Int"; S7_Expression := "ABS(IN1+IN2)" } Calculate(in1 := 1000, in2 := 1000, out => #最终调度距离上5)
   END_RUNG
   RUNG wire#powerrail
      Contact( #检修中 )
   END_RUNG wire#w18
   RUNG wire#powerrail
      Contact( #"5层边沿触发6" )
      wire#w19
      { S7_Templates := "SrcType := Int" } LE_Contact(in1 := #载重量, in2 := #限重分配)
      I_Contact( #检修中 )
      I_Contact( #死机 )
      { S7_Templates := "SrcType := Int"; S7_Expression := "ABS(IN1+IN2)" } Calculate(in1 := #"5层调度距离6", in2 := 0, out => #最终调度距离下5)
   END_RUNG
   RUNG wire#w19
      { S7_Templates := "SrcType := Int" } GT_Contact(in1 := #载重量, in2 := #限重分配)
      I_Contact( #检修中 )
      I_Contact( #死机 )
      { S7_Templates := "SrcType := Int"; S7_Expression := "ABS(IN1+IN2)" } Calculate(in1 := #"5层调度距离6", in2 := 100, out => #最终调度距离下5)
   END_RUNG
   RUNG wire#powerrail
      Contact( #"5层边沿触发7" )
      wire#w20
      { S7_Templates := "SrcType := Int" } LE_Contact(in1 := #载重量, in2 := #限重分配)
      I_Contact( #检修中 )
      I_Contact( #死机 )
      { S7_Templates := "SrcType := Int"; S7_Expression := "ABS(IN1+IN2)" } Calculate(in1 := #"5层调度距离7", in2 := 0, out => #最终调度距离下5)
   END_RUNG
   RUNG wire#w20
      { S7_Templates := "SrcType := Int" } GT_Contact(in1 := #载重量, in2 := #限重分配)
      I_Contact( #检修中 )
      I_Contact( #死机 )
      { S7_Templates := "SrcType := Int"; S7_Expression := "ABS(IN1+IN2)" } Calculate(in1 := #"5层调度距离7", in2 := 100, out => #最终调度距离下5)
   END_RUNG
   RUNG wire#powerrail
      Contact( #"5层边沿触发8" )
      wire#w21
      { S7_Templates := "SrcType := Int" } LE_Contact(in1 := #载重量, in2 := #限重分配)
      I_Contact( #检修中 )
      I_Contact( #死机 )
      { S7_Templates := "SrcType := Int"; S7_Expression := "ABS(IN1+IN2)" } Calculate(in1 := #"5层调度距离8", in2 := 0, out => #最终调度距离下5)
   END_RUNG
   RUNG wire#w21
      { S7_Templates := "SrcType := Int" } GT_Contact(in1 := #载重量, in2 := #限重分配)
      I_Contact( #检修中 )
      I_Contact( #死机 )
      { S7_Templates := "SrcType := Int"; S7_Expression := "ABS(IN1+IN2)" } Calculate(in1 := #"5层调度距离8", in2 := 100, out => #最终调度距离下5)
   END_RUNG
   RUNG wire#powerrail
      Contact( #"5层边沿触发9" )
      wire#w22
      { S7_Templates := "SrcType := Int" } LE_Contact(in1 := #载重量, in2 := #限重分配)
      I_Contact( #检修中 )
      I_Contact( #死机 )
      { S7_Templates := "SrcType := Int"; S7_Expression := "ABS(IN1+IN2)" } Calculate(in1 := #"5层调度距离9", in2 := 0, out => #最终调度距离下5)
   END_RUNG
   RUNG wire#w22
      { S7_Templates := "SrcType := Int" } GT_Contact(in1 := #载重量, in2 := #限重分配)
      I_Contact( #检修中 )
      I_Contact( #死机 )
      { S7_Templates := "SrcType := Int"; S7_Expression := "ABS(IN1+IN2)" } Calculate(in1 := #"5层调度距离9", in2 := 100, out => #最终调度距离下5)
   END_RUNG
   RUNG wire#powerrail
      Contact( #"5层边沿触发10" )
      wire#w23
      { S7_Templates := "SrcType := Int" } LE_Contact(in1 := #载重量, in2 := #限重分配)
      I_Contact( #检修中 )
      I_Contact( #死机 )
      { S7_Templates := "SrcType := Int"; S7_Expression := "ABS(IN1+IN2)" } Calculate(in1 := #"5层调度距离10", in2 := 0, out => #最终调度距离下5)
   END_RUNG
   RUNG wire#w23
      { S7_Templates := "SrcType := Int" } GT_Contact(in1 := #载重量, in2 := #限重分配)
      I_Contact( #检修中 )
      I_Contact( #死机 )
      { S7_Templates := "SrcType := Int"; S7_Expression := "ABS(IN1+IN2)" } Calculate(in1 := #"5层调度距离10", in2 := 100, out => #最终调度距离下5)
   END_RUNG
   RUNG wire#powerrail
      Contact( #死机 )
      wire#w24
      { S7_Templates := "SrcType := Int"; S7_Expression := "ABS(IN1+IN2)" } Calculate(in1 := 1000, in2 := 1000, out => #最终调度距离下5)
   END_RUNG
   RUNG wire#powerrail
      Contact( #检修中 )
   END_RUNG wire#w24
   // the same network as SCL:
   #_w1 := #上呼灯5 AND ((NOT #上行指示 AND NOT #下行指示 AND (#当前楼层 <= 5)) OR (#上行指示 AND (((5 = #当前楼层) AND #上下平层都为1) OR (5 > #当前楼层))));
   IF #_w1 THEN #"5层调度距离1" := ABS(#当前楼层-5)+#上行停站次数5+#上行停站次数5; END_IF;
   #"5层边沿触发1" := #_w1;
   #_w2 := #上呼灯5 AND (#下行指示 OR (NOT #上行指示 AND NOT #下行指示 AND (#当前楼层 > 5))) AND #外呼下面无目标5;
   IF #_w2 THEN #"5层调度距离2" := ABS(#当前楼层-5)+#下行停站次数5+#下行停站次数5; END_IF;
   #"5层边沿触发2" := #_w2;
   #_w3 := #上呼灯5 AND #下行指示 AND #外呼下面有目标5;
   IF #_w3 THEN
       #"5层调度距离3" := ABS(#外呼下面有目标最小数5+#外呼下面有目标最小数5-#当前楼层-5)+#下行停站次数1+#上行停站次数5+#上行停站次数5+#下行停站次数1+2;
   END_IF;
   #"5层边沿触发3" := #_w3;
   #_w4 := #上呼灯5 AND #上行指示 AND (((5 = #当前楼层) AND NOT #上下平层都为1) OR (5 < #当前楼层));
   #_w5 := #_w4 AND #外呼下面有目标5;
   IF #_w5 THEN
       #"5层调度距离4" := ABS(#外呼上面有目标最大数5-#当前楼层+#外呼上面有目标最大数5-#外呼下面有目标最小数5+5-#外呼下面有目标最小数5)+#上行停站次数5+#上行停站次数10+#上行停站次数10+#上行停站次数5+#下行停站次数1+#下行停站次数1+4;
   END_IF;
   #"5层边沿触发4" := #_w5;
   #_w6 := #_w4 AND #外呼下面无目标5;
   IF #_w6 THEN
       #"5层调度距离5" := ABS(#外呼上面有目标最大数5-#当前楼层+#外呼上面有目标最大数5-5)+#下行停站次数5+#上行停站次数10+#上行停站次数10+#下行停站次数5+2;
   END_IF;
   #"5层边沿触发5" := #_w6;
   #_w7 := #下呼灯5 AND ((NOT #上行指示 AND NOT #下行指示 AND (#当前楼层 >= 5)) OR (#下行指示 AND (((5 = #当前楼层) AND #上下平层都为1) OR (5 < #当前楼层))));
   IF #_w7 THEN #"5层调度距离6" := ABS(#当前楼层-5)+#下行停站次数5+#下行停站次数5; END_IF;
   #"5层边沿触发6" := #_w7;
   #_w8 := #下呼灯5 AND (#上行指示 OR (NOT #上行指示 AND NOT #下行指示 AND (#当前楼层 < 5))) AND #外呼上面无目标5;
   IF #_w8 THEN #"5层调度距离7" := ABS(#当前楼层-5)+#上行停站次数5+#上行停站次数5; END_IF;
   #"5层边沿触发7" := #_w8;
   #_w9 := #下呼灯5 AND #上行指示 AND #外呼上面有目标5;
   IF #_w9 THEN
       #"5层调度距离8" := ABS(#外呼上面有目标最大数5+#外呼上面有目标最大数5-#当前楼层-5)+#下行停站次数5+#上行停站次数10+#下行停站次数5+#上行停站次数10+2;
   END_IF;
   #"5层边沿触发8" := #_w9;
   #_w10 := #下呼灯5 AND #下行指示 AND (((5 = #当前楼层) AND NOT #上下平层都为1) OR (5 > #当前楼层));
   #_w11 := #_w10 AND #外呼上面有目标5;
   IF #_w11 THEN
       #"5层调度距离9" := ABS(#当前楼层-#外呼下面有目标最小数5+#外呼上面有目标最大数5-#外呼下面有目标最小数5+#外呼上面有目标最大数5-5)+#下行停站次数1+#下行停站次数5+#下行停站次数5+#下行停站次数1+#上行停站次数10+#上行停站次数10+4;
   END_IF;
   #"5层边沿触发9" := #_w11;
   #_w12 := #_w10 AND #外呼上面无目标5;
   IF #_w12 THEN
       #"5层调度距离10" := ABS(#当前楼层-#外呼下面有目标最小数5+5-#外呼下面有目标最小数5)+#下行停站次数1+#上行停站次数5+#上行停站次数5+#下行停站次数1+2;
   END_IF;
   #"5层边沿触发10" := #_w12;
   IF #"5层边沿触发1" AND (#载重量 <= #限重分配) AND NOT #检修中 AND NOT #死机 THEN #最终调度距离上5 := ABS(#"5层调度距离1"+0); END_IF;
   IF #"5层边沿触发1" AND (#载重量 > #限重分配) AND NOT #检修中 AND NOT #死机 THEN #最终调度距离上5 := ABS(#"5层调度距离1"+100); END_IF;
   IF #"5层边沿触发2" AND (#载重量 <= #限重分配) AND NOT #检修中 AND NOT #死机 THEN #最终调度距离上5 := ABS(#"5层调度距离2"+0); END_IF;
   IF #"5层边沿触发2" AND (#载重量 > #限重分配) AND NOT #检修中 AND NOT #死机 THEN #最终调度距离上5 := ABS(#"5层调度距离2"+100); END_IF;
   IF #"5层边沿触发3" AND (#载重量 <= #限重分配) AND NOT #检修中 AND NOT #死机 THEN #最终调度距离上5 := ABS(#"5层调度距离3"+0); END_IF;
   IF #"5层边沿触发3" AND (#载重量 > #限重分配) AND NOT #检修中 AND NOT #死机 THEN #最终调度距离上5 := ABS(#"5层调度距离3"+100); END_IF;
   IF #"5层边沿触发4" AND (#载重量 <= #限重分配) AND NOT #检修中 AND NOT #死机 THEN #最终调度距离上5 := ABS(#"5层调度距离4"+0); END_IF;
   IF #"5层边沿触发4" AND (#载重量 > #限重分配) AND NOT #检修中 AND NOT #死机 THEN #最终调度距离上5 := ABS(#"5层调度距离4"+100); END_IF;
   IF #"5层边沿触发5" AND (#载重量 <= #限重分配) AND NOT #检修中 AND NOT #死机 THEN #最终调度距离上5 := ABS(#"5层调度距离5"+0); END_IF;
   IF #"5层边沿触发5" AND (#载重量 > #限重分配) AND NOT #检修中 AND NOT #死机 THEN #最终调度距离上5 := ABS(#"5层调度距离5"+100); END_IF;
   IF #死机 OR #检修中 THEN #最终调度距离上5 := ABS(1000+1000); END_IF;
   IF #"5层边沿触发6" AND (#载重量 <= #限重分配) AND NOT #检修中 AND NOT #死机 THEN #最终调度距离下5 := ABS(#"5层调度距离6"+0); END_IF;
   IF #"5层边沿触发6" AND (#载重量 > #限重分配) AND NOT #检修中 AND NOT #死机 THEN #最终调度距离下5 := ABS(#"5层调度距离6"+100); END_IF;
   IF #"5层边沿触发7" AND (#载重量 <= #限重分配) AND NOT #检修中 AND NOT #死机 THEN #最终调度距离下5 := ABS(#"5层调度距离7"+0); END_IF;
   IF #"5层边沿触发7" AND (#载重量 > #限重分配) AND NOT #检修中 AND NOT #死机 THEN #最终调度距离下5 := ABS(#"5层调度距离7"+100); END_IF;
   IF #"5层边沿触发8" AND (#载重量 <= #限重分配) AND NOT #检修中 AND NOT #死机 THEN #最终调度距离下5 := ABS(#"5层调度距离8"+0); END_IF;
   IF #"5层边沿触发8" AND (#载重量 > #限重分配) AND NOT #检修中 AND NOT #死机 THEN #最终调度距离下5 := ABS(#"5层调度距离8"+100); END_IF;
   IF #"5层边沿触发9" AND (#载重量 <= #限重分配) AND NOT #检修中 AND NOT #死机 THEN #最终调度距离下5 := ABS(#"5层调度距离9"+0); END_IF;
   IF #"5层边沿触发9" AND (#载重量 > #限重分配) AND NOT #检修中 AND NOT #死机 THEN #最终调度距离下5 := ABS(#"5层调度距离9"+100); END_IF;
   IF #"5层边沿触发10" AND (#载重量 <= #限重分配) AND NOT #检修中 AND NOT #死机 THEN #最终调度距离下5 := ABS(#"5层调度距离10"+0); END_IF;
   IF #"5层边沿触发10" AND (#载重量 > #限重分配) AND NOT #检修中 AND NOT #死机 THEN #最终调度距离下5 := ABS(#"5层调度距离10"+100); END_IF;
   IF #死机 OR #检修中 THEN #最终调度距离下5 := ABS(1000+1000); END_IF;
END_REGION

REGION Network 5: 6层调度距离
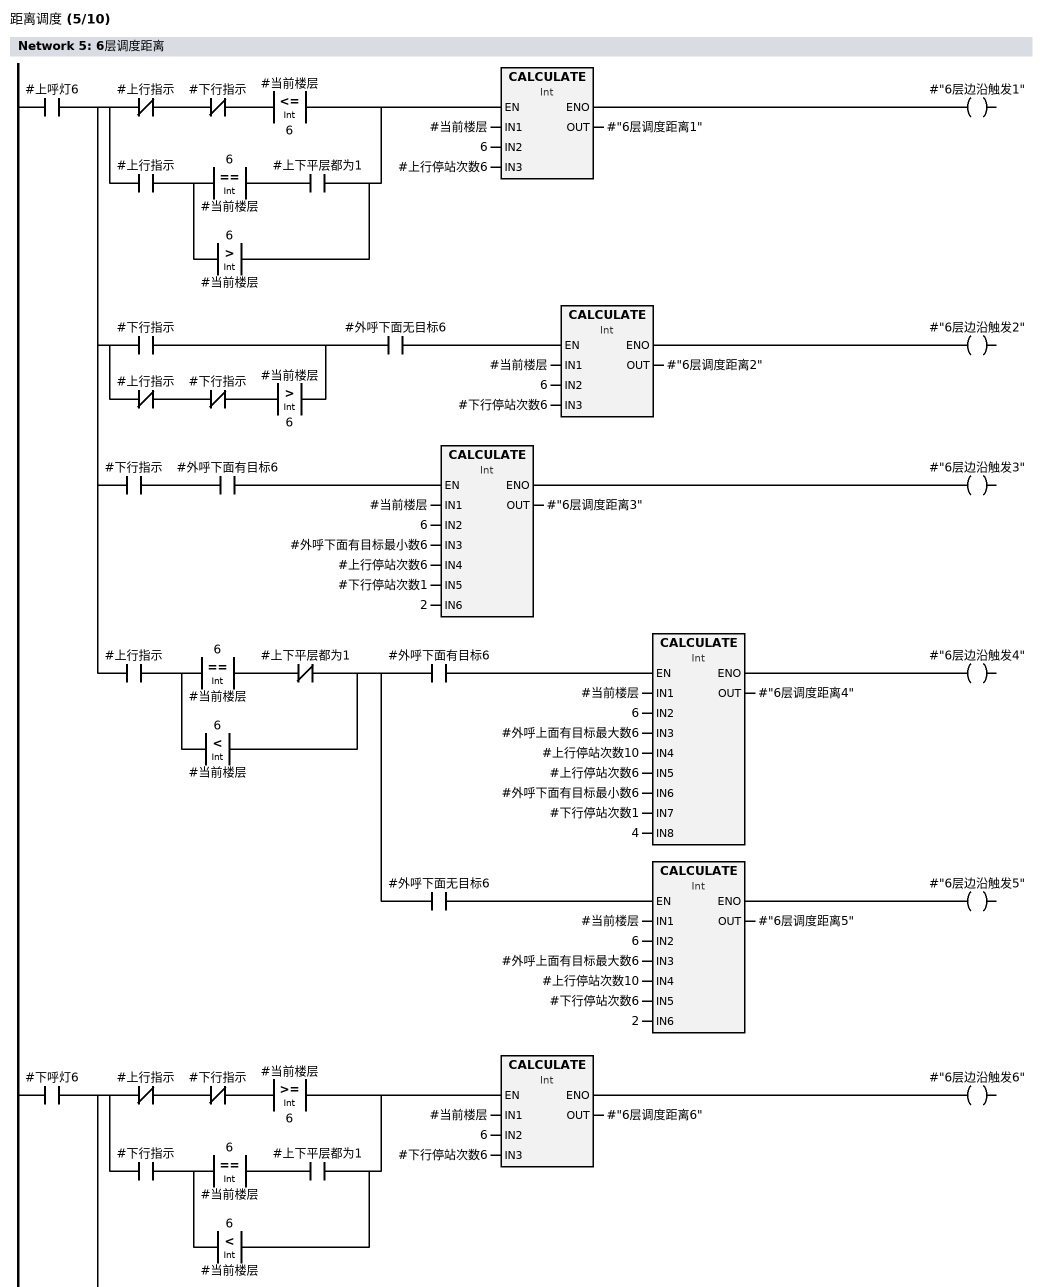
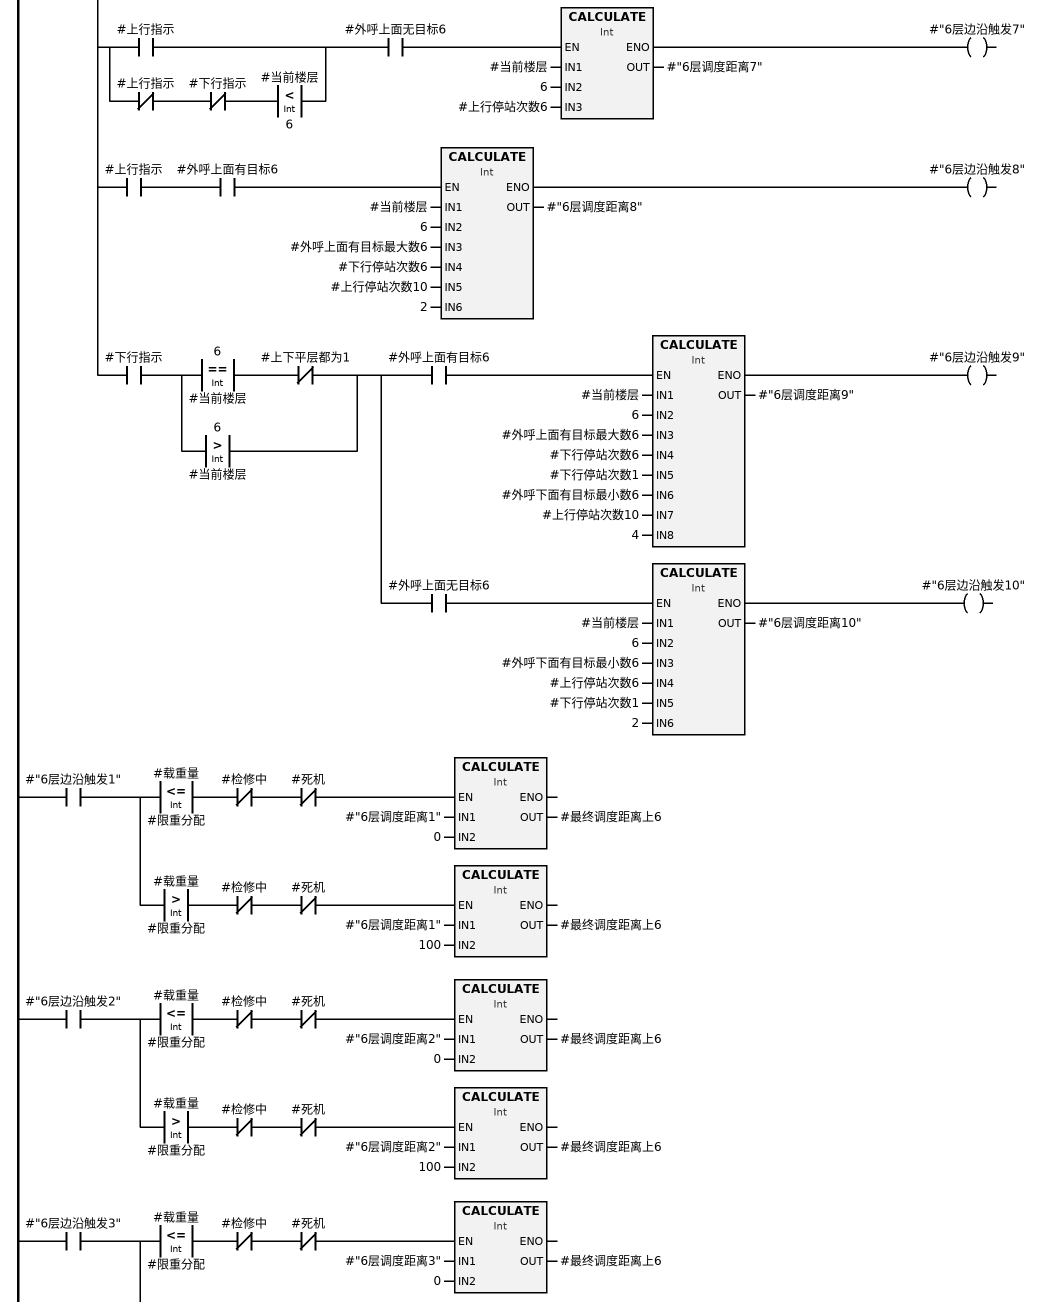
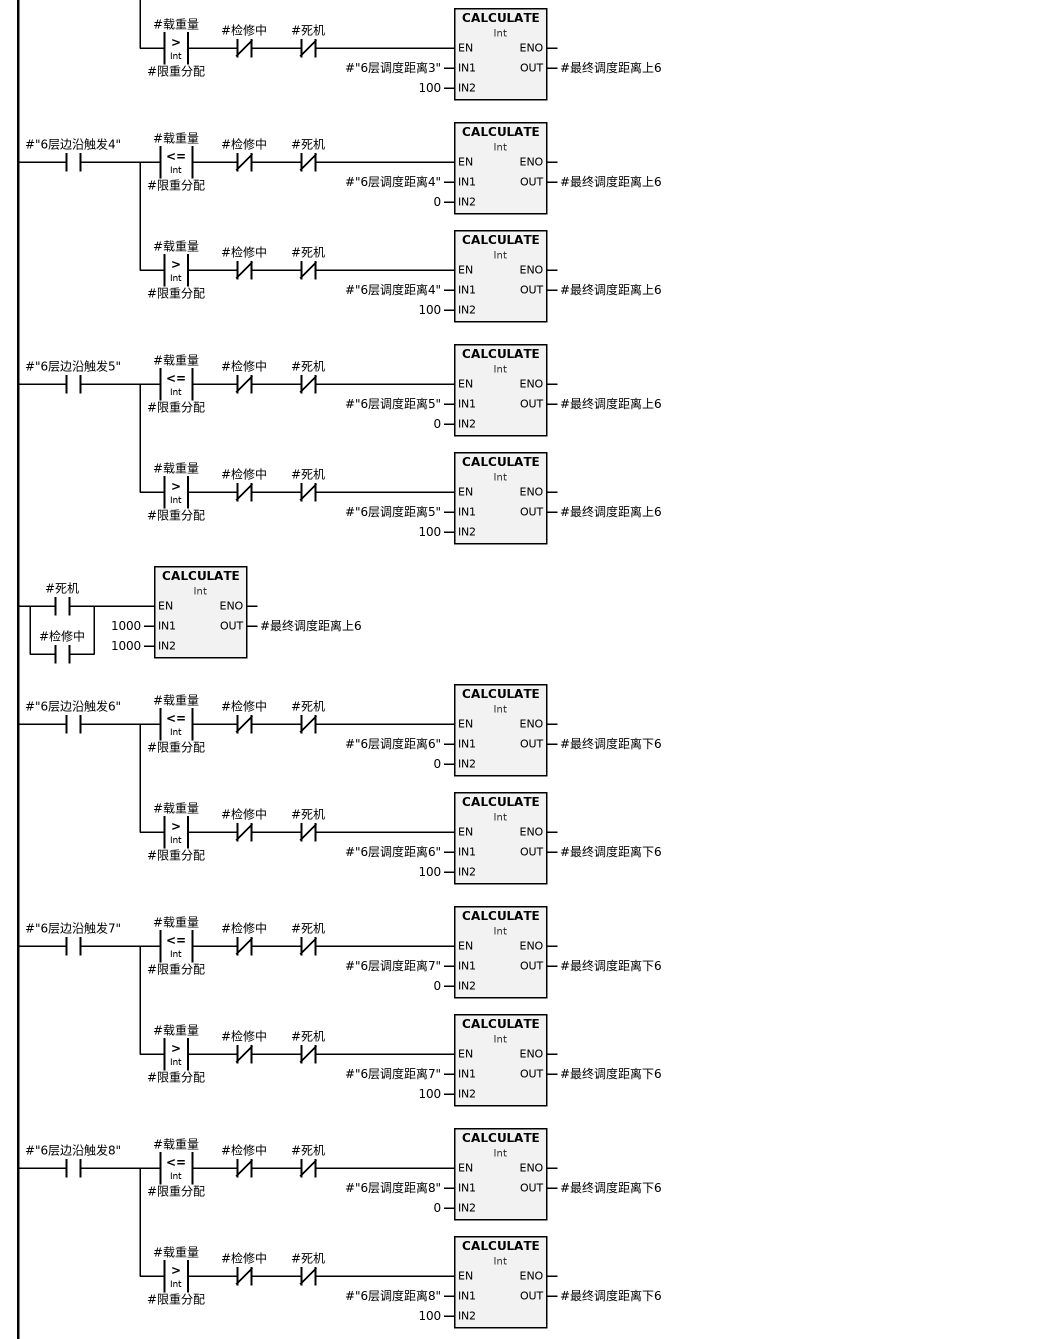
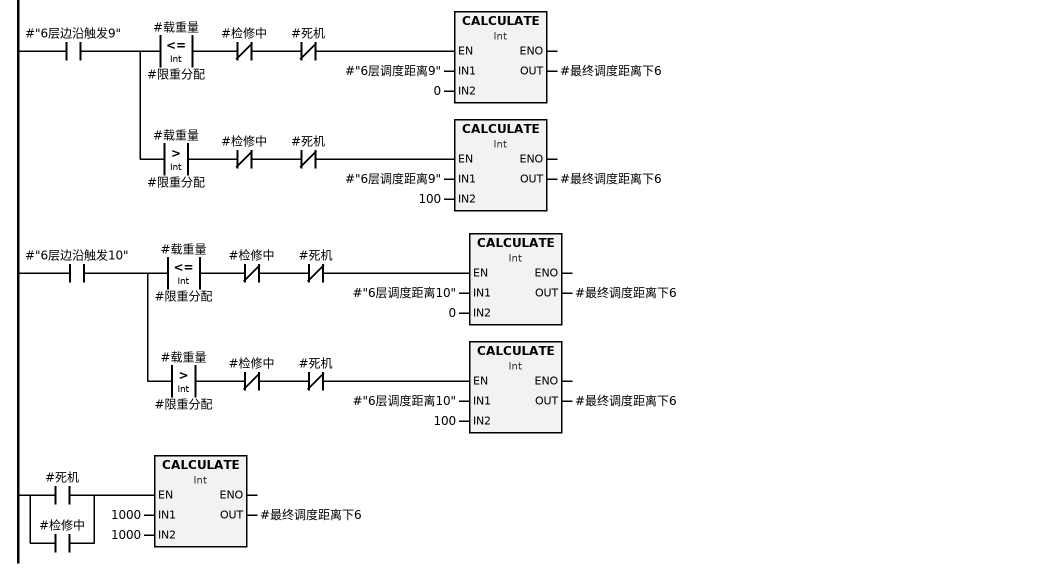
   RUNG wire#powerrail
      Contact( #上呼灯6 )
      wire#w1
      I_Contact( #上行指示 )
      I_Contact( #下行指示 )
      { S7_Templates := "SrcType := Int" } LE_Contact(in1 := #当前楼层, in2 := 6)
      wire#w2
      { S7_Templates := "SrcType := Int"; S7_Expression := "ABS(IN1-IN2)+IN3+IN3" } Calculate(in1 := #当前楼层, in2 := 6, in3 := #上行停站次数6, out => #"6层调度距离1")
      Coil( #"6层边沿触发1" )
   END_RUNG
   RUNG wire#w1
      Contact( #上行指示 )
      wire#w3
      { S7_Templates := "SrcType := Int" } EQ_Contact(in1 := 6, in2 := #当前楼层)
      Contact( #上下平层都为1 )
   END_RUNG wire#w2
   RUNG wire#w3
      { S7_Templates := "SrcType := Int" } GT_Contact(in1 := 6, in2 := #当前楼层)
   END_RUNG wire#w2
   RUNG wire#w1
      Contact( #下行指示 )
      wire#w4
      Contact( #外呼下面无目标6 )
      { S7_Templates := "SrcType := Int"; S7_Expression := "ABS(IN1-IN2)+IN3+IN3" } Calculate(in1 := #当前楼层, in2 := 6, in3 := #下行停站次数6, out => #"6层调度距离2")
      Coil( #"6层边沿触发2" )
   END_RUNG
   RUNG wire#w1
      I_Contact( #上行指示 )
      I_Contact( #下行指示 )
      { S7_Templates := "SrcType := Int" } GT_Contact(in1 := #当前楼层, in2 := 6)
   END_RUNG wire#w4
   RUNG wire#w1
      Contact( #下行指示 )
      Contact( #外呼下面有目标6 )
      { S7_Templates := "SrcType := Int"; S7_Expression := "ABS(IN3+IN3-IN1-IN2)+IN5+IN4+IN4+IN5+IN2" } Calculate(in1 := #当前楼层, in2 := 6, in3 := #外呼下面有目标最小数6, in4 := #上行停站次数6, in5 := #下行停站次数1, in6 := 2, out => #"6层调度距离3")
      Coil( #"6层边沿触发3" )
   END_RUNG
   RUNG wire#w1
      Contact( #上行指示 )
      wire#w5
      { S7_Templates := "SrcType := Int" } EQ_Contact(in1 := 6, in2 := #当前楼层)
      I_Contact( #上下平层都为1 )
      wire#w6
      Contact( #外呼下面有目标6 )
      { S7_Templates := "SrcType := Int"; S7_Expression := "ABS(IN3-IN1+IN3-IN6+IN2-IN6)+IN5+IN4+IN4+IN5+IN7+IN7+IN8" } Calculate(in1 := #当前楼层, in2 := 6, in3 := #外呼上面有目标最大数6, in4 := #上行停站次数10, in5 := #上行停站次数6, in6 := #外呼下面有目标最小数6, in7 := #下行停站次数1, in8 := 4, out => #"6层调度距离4")
      Coil( #"6层边沿触发4" )
   END_RUNG
   RUNG wire#w5
      { S7_Templates := "SrcType := Int" } LT_Contact(in1 := 6, in2 := #当前楼层)
   END_RUNG wire#w6
   RUNG wire#w6
      Contact( #外呼下面无目标6 )
      { S7_Templates := "SrcType := Int"; S7_Expression := "ABS(IN3-IN1+IN3-IN2)+IN5+IN4+IN4+IN5+IN6" } Calculate(in1 := #当前楼层, in2 := 6, in3 := #外呼上面有目标最大数6, in4 := #上行停站次数10, in5 := #下行停站次数6, in6 := 2, out => #"6层调度距离5")
      Coil( #"6层边沿触发5" )
   END_RUNG
   RUNG wire#powerrail
      Contact( #下呼灯6 )
      wire#w7
      I_Contact( #上行指示 )
      I_Contact( #下行指示 )
      { S7_Templates := "SrcType := Int" } GE_Contact(in1 := #当前楼层, in2 := 6)
      wire#w8
      { S7_Templates := "SrcType := Int"; S7_Expression := "ABS(IN1-IN2)+IN3+IN3" } Calculate(in1 := #当前楼层, in2 := 6, in3 := #下行停站次数6, out => #"6层调度距离6")
      Coil( #"6层边沿触发6" )
   END_RUNG
   RUNG wire#w7
      Contact( #下行指示 )
      wire#w9
      { S7_Templates := "SrcType := Int" } EQ_Contact(in1 := 6, in2 := #当前楼层)
      Contact( #上下平层都为1 )
   END_RUNG wire#w8
   RUNG wire#w9
      { S7_Templates := "SrcType := Int" } LT_Contact(in1 := 6, in2 := #当前楼层)
   END_RUNG wire#w8
   RUNG wire#w7
      Contact( #上行指示 )
      wire#w10
      Contact( #外呼上面无目标6 )
      { S7_Templates := "SrcType := Int"; S7_Expression := "ABS(IN1-IN2)+IN3+IN3" } Calculate(in1 := #当前楼层, in2 := 6, in3 := #上行停站次数6, out => #"6层调度距离7")
      Coil( #"6层边沿触发7" )
   END_RUNG
   RUNG wire#w7
      I_Contact( #上行指示 )
      I_Contact( #下行指示 )
      { S7_Templates := "SrcType := Int" } LT_Contact(in1 := #当前楼层, in2 := 6)
   END_RUNG wire#w10
   RUNG wire#w7
      Contact( #上行指示 )
      Contact( #外呼上面有目标6 )
      { S7_Templates := "SrcType := Int"; S7_Expression := "ABS(IN3+IN3-IN1-IN2)+IN4+IN5+IN4+IN5+IN6" } Calculate(in1 := #当前楼层, in2 := 6, in3 := #外呼上面有目标最大数6, in4 := #下行停站次数6, in5 := #上行停站次数10, in6 := 2, out => #"6层调度距离8")
      Coil( #"6层边沿触发8" )
   END_RUNG
   RUNG wire#w7
      Contact( #下行指示 )
      wire#w11
      { S7_Templates := "SrcType := Int" } EQ_Contact(in1 := 6, in2 := #当前楼层)
      I_Contact( #上下平层都为1 )
      wire#w12
      Contact( #外呼上面有目标6 )
      { S7_Templates := "SrcType := Int"; S7_Expression := "ABS(IN1-IN6+IN3-IN6+IN3-IN2)+IN5+IN4+IN4+IN5+IN7+IN7+IN8" } Calculate(in1 := #当前楼层, in2 := 6, in3 := #外呼上面有目标最大数6, in4 := #下行停站次数6, in5 := #下行停站次数1, in6 := #外呼下面有目标最小数6, in7 := #上行停站次数10, in8 := 4, out => #"6层调度距离9")
      Coil( #"6层边沿触发9" )
   END_RUNG
   RUNG wire#w11
      { S7_Templates := "SrcType := Int" } GT_Contact(in1 := 6, in2 := #当前楼层)
   END_RUNG wire#w12
   RUNG wire#w12
      Contact( #外呼上面无目标6 )
      { S7_Templates := "SrcType := Int"; S7_Expression := "ABS(IN1-IN3+IN2-IN3)+IN5+IN4+IN4+IN5+IN6" } Calculate(in1 := #当前楼层, in2 := 6, in3 := #外呼下面有目标最小数6, in4 := #上行停站次数6, in5 := #下行停站次数1, in6 := 2, out => #"6层调度距离10")
      Coil( #"6层边沿触发10" )
   END_RUNG
   RUNG wire#powerrail
      Contact( #"6层边沿触发1" )
      wire#w13
      { S7_Templates := "SrcType := Int" } LE_Contact(in1 := #载重量, in2 := #限重分配)
      I_Contact( #检修中 )
      I_Contact( #死机 )
      { S7_Templates := "SrcType := Int"; S7_Expression := "ABS(IN1+IN2)" } Calculate(in1 := #"6层调度距离1", in2 := 0, out => #最终调度距离上6)
   END_RUNG
   RUNG wire#w13
      { S7_Templates := "SrcType := Int" } GT_Contact(in1 := #载重量, in2 := #限重分配)
      I_Contact( #检修中 )
      I_Contact( #死机 )
      { S7_Templates := "SrcType := Int"; S7_Expression := "ABS(IN1+IN2)" } Calculate(in1 := #"6层调度距离1", in2 := 100, out => #最终调度距离上6)
   END_RUNG
   RUNG wire#powerrail
      Contact( #"6层边沿触发2" )
      wire#w14
      { S7_Templates := "SrcType := Int" } LE_Contact(in1 := #载重量, in2 := #限重分配)
      I_Contact( #检修中 )
      I_Contact( #死机 )
      { S7_Templates := "SrcType := Int"; S7_Expression := "ABS(IN1+IN2)" } Calculate(in1 := #"6层调度距离2", in2 := 0, out => #最终调度距离上6)
   END_RUNG
   RUNG wire#w14
      { S7_Templates := "SrcType := Int" } GT_Contact(in1 := #载重量, in2 := #限重分配)
      I_Contact( #检修中 )
      I_Contact( #死机 )
      { S7_Templates := "SrcType := Int"; S7_Expression := "ABS(IN1+IN2)" } Calculate(in1 := #"6层调度距离2", in2 := 100, out => #最终调度距离上6)
   END_RUNG
   RUNG wire#powerrail
      Contact( #"6层边沿触发3" )
      wire#w15
      { S7_Templates := "SrcType := Int" } LE_Contact(in1 := #载重量, in2 := #限重分配)
      I_Contact( #检修中 )
      I_Contact( #死机 )
      { S7_Templates := "SrcType := Int"; S7_Expression := "ABS(IN1+IN2)" } Calculate(in1 := #"6层调度距离3", in2 := 0, out => #最终调度距离上6)
   END_RUNG
   RUNG wire#w15
      { S7_Templates := "SrcType := Int" } GT_Contact(in1 := #载重量, in2 := #限重分配)
      I_Contact( #检修中 )
      I_Contact( #死机 )
      { S7_Templates := "SrcType := Int"; S7_Expression := "ABS(IN1+IN2)" } Calculate(in1 := #"6层调度距离3", in2 := 100, out => #最终调度距离上6)
   END_RUNG
   RUNG wire#powerrail
      Contact( #"6层边沿触发4" )
      wire#w16
      { S7_Templates := "SrcType := Int" } LE_Contact(in1 := #载重量, in2 := #限重分配)
      I_Contact( #检修中 )
      I_Contact( #死机 )
      { S7_Templates := "SrcType := Int"; S7_Expression := "ABS(IN1+IN2)" } Calculate(in1 := #"6层调度距离4", in2 := 0, out => #最终调度距离上6)
   END_RUNG
   RUNG wire#w16
      { S7_Templates := "SrcType := Int" } GT_Contact(in1 := #载重量, in2 := #限重分配)
      I_Contact( #检修中 )
      I_Contact( #死机 )
      { S7_Templates := "SrcType := Int"; S7_Expression := "ABS(IN1+IN2)" } Calculate(in1 := #"6层调度距离4", in2 := 100, out => #最终调度距离上6)
   END_RUNG
   RUNG wire#powerrail
      Contact( #"6层边沿触发5" )
      wire#w17
      { S7_Templates := "SrcType := Int" } LE_Contact(in1 := #载重量, in2 := #限重分配)
      I_Contact( #检修中 )
      I_Contact( #死机 )
      { S7_Templates := "SrcType := Int"; S7_Expression := "ABS(IN1+IN2)" } Calculate(in1 := #"6层调度距离5", in2 := 0, out => #最终调度距离上6)
   END_RUNG
   RUNG wire#w17
      { S7_Templates := "SrcType := Int" } GT_Contact(in1 := #载重量, in2 := #限重分配)
      I_Contact( #检修中 )
      I_Contact( #死机 )
      { S7_Templates := "SrcType := Int"; S7_Expression := "ABS(IN1+IN2)" } Calculate(in1 := #"6层调度距离5", in2 := 100, out => #最终调度距离上6)
   END_RUNG
   RUNG wire#powerrail
      Contact( #死机 )
      wire#w18
      { S7_Templates := "SrcType := Int"; S7_Expression := "ABS(IN1+IN2)" } Calculate(in1 := 1000, in2 := 1000, out => #最终调度距离上6)
   END_RUNG
   RUNG wire#powerrail
      Contact( #检修中 )
   END_RUNG wire#w18
   RUNG wire#powerrail
      Contact( #"6层边沿触发6" )
      wire#w19
      { S7_Templates := "SrcType := Int" } LE_Contact(in1 := #载重量, in2 := #限重分配)
      I_Contact( #检修中 )
      I_Contact( #死机 )
      { S7_Templates := "SrcType := Int"; S7_Expression := "ABS(IN1+IN2)" } Calculate(in1 := #"6层调度距离6", in2 := 0, out => #最终调度距离下6)
   END_RUNG
   RUNG wire#w19
      { S7_Templates := "SrcType := Int" } GT_Contact(in1 := #载重量, in2 := #限重分配)
      I_Contact( #检修中 )
      I_Contact( #死机 )
      { S7_Templates := "SrcType := Int"; S7_Expression := "ABS(IN1+IN2)" } Calculate(in1 := #"6层调度距离6", in2 := 100, out => #最终调度距离下6)
   END_RUNG
   RUNG wire#powerrail
      Contact( #"6层边沿触发7" )
      wire#w20
      { S7_Templates := "SrcType := Int" } LE_Contact(in1 := #载重量, in2 := #限重分配)
      I_Contact( #检修中 )
      I_Contact( #死机 )
      { S7_Templates := "SrcType := Int"; S7_Expression := "ABS(IN1+IN2)" } Calculate(in1 := #"6层调度距离7", in2 := 0, out => #最终调度距离下6)
   END_RUNG
   RUNG wire#w20
      { S7_Templates := "SrcType := Int" } GT_Contact(in1 := #载重量, in2 := #限重分配)
      I_Contact( #检修中 )
      I_Contact( #死机 )
      { S7_Templates := "SrcType := Int"; S7_Expression := "ABS(IN1+IN2)" } Calculate(in1 := #"6层调度距离7", in2 := 100, out => #最终调度距离下6)
   END_RUNG
   RUNG wire#powerrail
      Contact( #"6层边沿触发8" )
      wire#w21
      { S7_Templates := "SrcType := Int" } LE_Contact(in1 := #载重量, in2 := #限重分配)
      I_Contact( #检修中 )
      I_Contact( #死机 )
      { S7_Templates := "SrcType := Int"; S7_Expression := "ABS(IN1+IN2)" } Calculate(in1 := #"6层调度距离8", in2 := 0, out => #最终调度距离下6)
   END_RUNG
   RUNG wire#w21
      { S7_Templates := "SrcType := Int" } GT_Contact(in1 := #载重量, in2 := #限重分配)
      I_Contact( #检修中 )
      I_Contact( #死机 )
      { S7_Templates := "SrcType := Int"; S7_Expression := "ABS(IN1+IN2)" } Calculate(in1 := #"6层调度距离8", in2 := 100, out => #最终调度距离下6)
   END_RUNG
   RUNG wire#powerrail
      Contact( #"6层边沿触发9" )
      wire#w22
      { S7_Templates := "SrcType := Int" } LE_Contact(in1 := #载重量, in2 := #限重分配)
      I_Contact( #检修中 )
      I_Contact( #死机 )
      { S7_Templates := "SrcType := Int"; S7_Expression := "ABS(IN1+IN2)" } Calculate(in1 := #"6层调度距离9", in2 := 0, out => #最终调度距离下6)
   END_RUNG
   RUNG wire#w22
      { S7_Templates := "SrcType := Int" } GT_Contact(in1 := #载重量, in2 := #限重分配)
      I_Contact( #检修中 )
      I_Contact( #死机 )
      { S7_Templates := "SrcType := Int"; S7_Expression := "ABS(IN1+IN2)" } Calculate(in1 := #"6层调度距离9", in2 := 100, out => #最终调度距离下6)
   END_RUNG
   RUNG wire#powerrail
      Contact( #"6层边沿触发10" )
      wire#w23
      { S7_Templates := "SrcType := Int" } LE_Contact(in1 := #载重量, in2 := #限重分配)
      I_Contact( #检修中 )
      I_Contact( #死机 )
      { S7_Templates := "SrcType := Int"; S7_Expression := "ABS(IN1+IN2)" } Calculate(in1 := #"6层调度距离10", in2 := 0, out => #最终调度距离下6)
   END_RUNG
   RUNG wire#w23
      { S7_Templates := "SrcType := Int" } GT_Contact(in1 := #载重量, in2 := #限重分配)
      I_Contact( #检修中 )
      I_Contact( #死机 )
      { S7_Templates := "SrcType := Int"; S7_Expression := "ABS(IN1+IN2)" } Calculate(in1 := #"6层调度距离10", in2 := 100, out => #最终调度距离下6)
   END_RUNG
   RUNG wire#powerrail
      Contact( #死机 )
      wire#w24
      { S7_Templates := "SrcType := Int"; S7_Expression := "ABS(IN1+IN2)" } Calculate(in1 := 1000, in2 := 1000, out => #最终调度距离下6)
   END_RUNG
   RUNG wire#powerrail
      Contact( #检修中 )
   END_RUNG wire#w24
   // the same network as SCL:
   #_w1 := #上呼灯6 AND ((NOT #上行指示 AND NOT #下行指示 AND (#当前楼层 <= 6)) OR (#上行指示 AND (((6 = #当前楼层) AND #上下平层都为1) OR (6 > #当前楼层))));
   IF #_w1 THEN #"6层调度距离1" := ABS(#当前楼层-6)+#上行停站次数6+#上行停站次数6; END_IF;
   #"6层边沿触发1" := #_w1;
   #_w2 := #上呼灯6 AND (#下行指示 OR (NOT #上行指示 AND NOT #下行指示 AND (#当前楼层 > 6))) AND #外呼下面无目标6;
   IF #_w2 THEN #"6层调度距离2" := ABS(#当前楼层-6)+#下行停站次数6+#下行停站次数6; END_IF;
   #"6层边沿触发2" := #_w2;
   #_w3 := #上呼灯6 AND #下行指示 AND #外呼下面有目标6;
   IF #_w3 THEN
       #"6层调度距离3" := ABS(#外呼下面有目标最小数6+#外呼下面有目标最小数6-#当前楼层-6)+#下行停站次数1+#上行停站次数6+#上行停站次数6+#下行停站次数1+6;
   END_IF;
   #"6层边沿触发3" := #_w3;
   #_w4 := #上呼灯6 AND #上行指示 AND (((6 = #当前楼层) AND NOT #上下平层都为1) OR (6 < #当前楼层));
   #_w5 := #_w4 AND #外呼下面有目标6;
   IF #_w5 THEN
       #"6层调度距离4" := ABS(#外呼上面有目标最大数6-#当前楼层+#外呼上面有目标最大数6-#外呼下面有目标最小数6+6-#外呼下面有目标最小数6)+#上行停站次数6+#上行停站次数10+#上行停站次数10+#上行停站次数6+#下行停站次数1+#下行停站次数1+4;
   END_IF;
   #"6层边沿触发4" := #_w5;
   #_w6 := #_w4 AND #外呼下面无目标6;
   IF #_w6 THEN
       #"6层调度距离5" := ABS(#外呼上面有目标最大数6-#当前楼层+#外呼上面有目标最大数6-6)+#下行停站次数6+#上行停站次数10+#上行停站次数10+#下行停站次数6+2;
   END_IF;
   #"6层边沿触发5" := #_w6;
   #_w7 := #下呼灯6 AND ((NOT #上行指示 AND NOT #下行指示 AND (#当前楼层 >= 6)) OR (#下行指示 AND (((6 = #当前楼层) AND #上下平层都为1) OR (6 < #当前楼层))));
   IF #_w7 THEN #"6层调度距离6" := ABS(#当前楼层-6)+#下行停站次数6+#下行停站次数6; END_IF;
   #"6层边沿触发6" := #_w7;
   #_w8 := #下呼灯6 AND (#上行指示 OR (NOT #上行指示 AND NOT #下行指示 AND (#当前楼层 < 6))) AND #外呼上面无目标6;
   IF #_w8 THEN #"6层调度距离7" := ABS(#当前楼层-6)+#上行停站次数6+#上行停站次数6; END_IF;
   #"6层边沿触发7" := #_w8;
   #_w9 := #下呼灯6 AND #上行指示 AND #外呼上面有目标6;
   IF #_w9 THEN
       #"6层调度距离8" := ABS(#外呼上面有目标最大数6+#外呼上面有目标最大数6-#当前楼层-6)+#下行停站次数6+#上行停站次数10+#下行停站次数6+#上行停站次数10+2;
   END_IF;
   #"6层边沿触发8" := #_w9;
   #_w10 := #下呼灯6 AND #下行指示 AND (((6 = #当前楼层) AND NOT #上下平层都为1) OR (6 > #当前楼层));
   #_w11 := #_w10 AND #外呼上面有目标6;
   IF #_w11 THEN
       #"6层调度距离9" := ABS(#当前楼层-#外呼下面有目标最小数6+#外呼上面有目标最大数6-#外呼下面有目标最小数6+#外呼上面有目标最大数6-6)+#下行停站次数1+#下行停站次数6+#下行停站次数6+#下行停站次数1+#上行停站次数10+#上行停站次数10+4;
   END_IF;
   #"6层边沿触发9" := #_w11;
   #_w12 := #_w10 AND #外呼上面无目标6;
   IF #_w12 THEN
       #"6层调度距离10" := ABS(#当前楼层-#外呼下面有目标最小数6+6-#外呼下面有目标最小数6)+#下行停站次数1+#上行停站次数6+#上行停站次数6+#下行停站次数1+2;
   END_IF;
   #"6层边沿触发10" := #_w12;
   IF #"6层边沿触发1" AND (#载重量 <= #限重分配) AND NOT #检修中 AND NOT #死机 THEN #最终调度距离上6 := ABS(#"6层调度距离1"+0); END_IF;
   IF #"6层边沿触发1" AND (#载重量 > #限重分配) AND NOT #检修中 AND NOT #死机 THEN #最终调度距离上6 := ABS(#"6层调度距离1"+100); END_IF;
   IF #"6层边沿触发2" AND (#载重量 <= #限重分配) AND NOT #检修中 AND NOT #死机 THEN #最终调度距离上6 := ABS(#"6层调度距离2"+0); END_IF;
   IF #"6层边沿触发2" AND (#载重量 > #限重分配) AND NOT #检修中 AND NOT #死机 THEN #最终调度距离上6 := ABS(#"6层调度距离2"+100); END_IF;
   IF #"6层边沿触发3" AND (#载重量 <= #限重分配) AND NOT #检修中 AND NOT #死机 THEN #最终调度距离上6 := ABS(#"6层调度距离3"+0); END_IF;
   IF #"6层边沿触发3" AND (#载重量 > #限重分配) AND NOT #检修中 AND NOT #死机 THEN #最终调度距离上6 := ABS(#"6层调度距离3"+100); END_IF;
   IF #"6层边沿触发4" AND (#载重量 <= #限重分配) AND NOT #检修中 AND NOT #死机 THEN #最终调度距离上6 := ABS(#"6层调度距离4"+0); END_IF;
   IF #"6层边沿触发4" AND (#载重量 > #限重分配) AND NOT #检修中 AND NOT #死机 THEN #最终调度距离上6 := ABS(#"6层调度距离4"+100); END_IF;
   IF #"6层边沿触发5" AND (#载重量 <= #限重分配) AND NOT #检修中 AND NOT #死机 THEN #最终调度距离上6 := ABS(#"6层调度距离5"+0); END_IF;
   IF #"6层边沿触发5" AND (#载重量 > #限重分配) AND NOT #检修中 AND NOT #死机 THEN #最终调度距离上6 := ABS(#"6层调度距离5"+100); END_IF;
   IF #死机 OR #检修中 THEN #最终调度距离上6 := ABS(1000+1000); END_IF;
   IF #"6层边沿触发6" AND (#载重量 <= #限重分配) AND NOT #检修中 AND NOT #死机 THEN #最终调度距离下6 := ABS(#"6层调度距离6"+0); END_IF;
   IF #"6层边沿触发6" AND (#载重量 > #限重分配) AND NOT #检修中 AND NOT #死机 THEN #最终调度距离下6 := ABS(#"6层调度距离6"+100); END_IF;
   IF #"6层边沿触发7" AND (#载重量 <= #限重分配) AND NOT #检修中 AND NOT #死机 THEN #最终调度距离下6 := ABS(#"6层调度距离7"+0); END_IF;
   IF #"6层边沿触发7" AND (#载重量 > #限重分配) AND NOT #检修中 AND NOT #死机 THEN #最终调度距离下6 := ABS(#"6层调度距离7"+100); END_IF;
   IF #"6层边沿触发8" AND (#载重量 <= #限重分配) AND NOT #检修中 AND NOT #死机 THEN #最终调度距离下6 := ABS(#"6层调度距离8"+0); END_IF;
   IF #"6层边沿触发8" AND (#载重量 > #限重分配) AND NOT #检修中 AND NOT #死机 THEN #最终调度距离下6 := ABS(#"6层调度距离8"+100); END_IF;
   IF #"6层边沿触发9" AND (#载重量 <= #限重分配) AND NOT #检修中 AND NOT #死机 THEN #最终调度距离下6 := ABS(#"6层调度距离9"+0); END_IF;
   IF #"6层边沿触发9" AND (#载重量 > #限重分配) AND NOT #检修中 AND NOT #死机 THEN #最终调度距离下6 := ABS(#"6层调度距离9"+100); END_IF;
   IF #"6层边沿触发10" AND (#载重量 <= #限重分配) AND NOT #检修中 AND NOT #死机 THEN #最终调度距离下6 := ABS(#"6层调度距离10"+0); END_IF;
   IF #"6层边沿触发10" AND (#载重量 > #限重分配) AND NOT #检修中 AND NOT #死机 THEN #最终调度距离下6 := ABS(#"6层调度距离10"+100); END_IF;
   IF #死机 OR #检修中 THEN #最终调度距离下6 := ABS(1000+1000); END_IF;
END_REGION

REGION Network 6: 7层调度距离
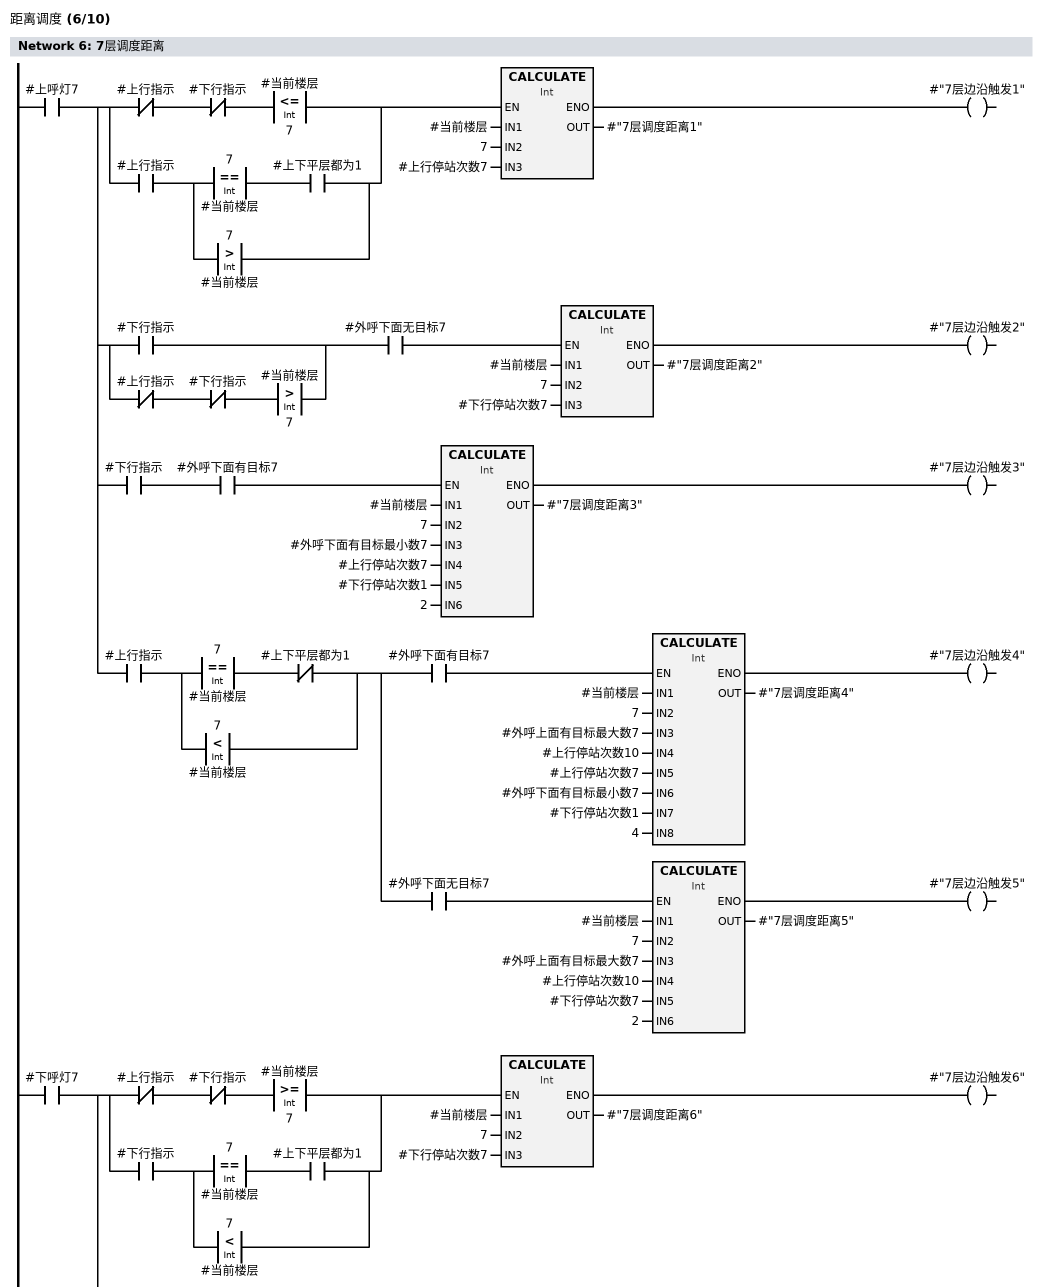
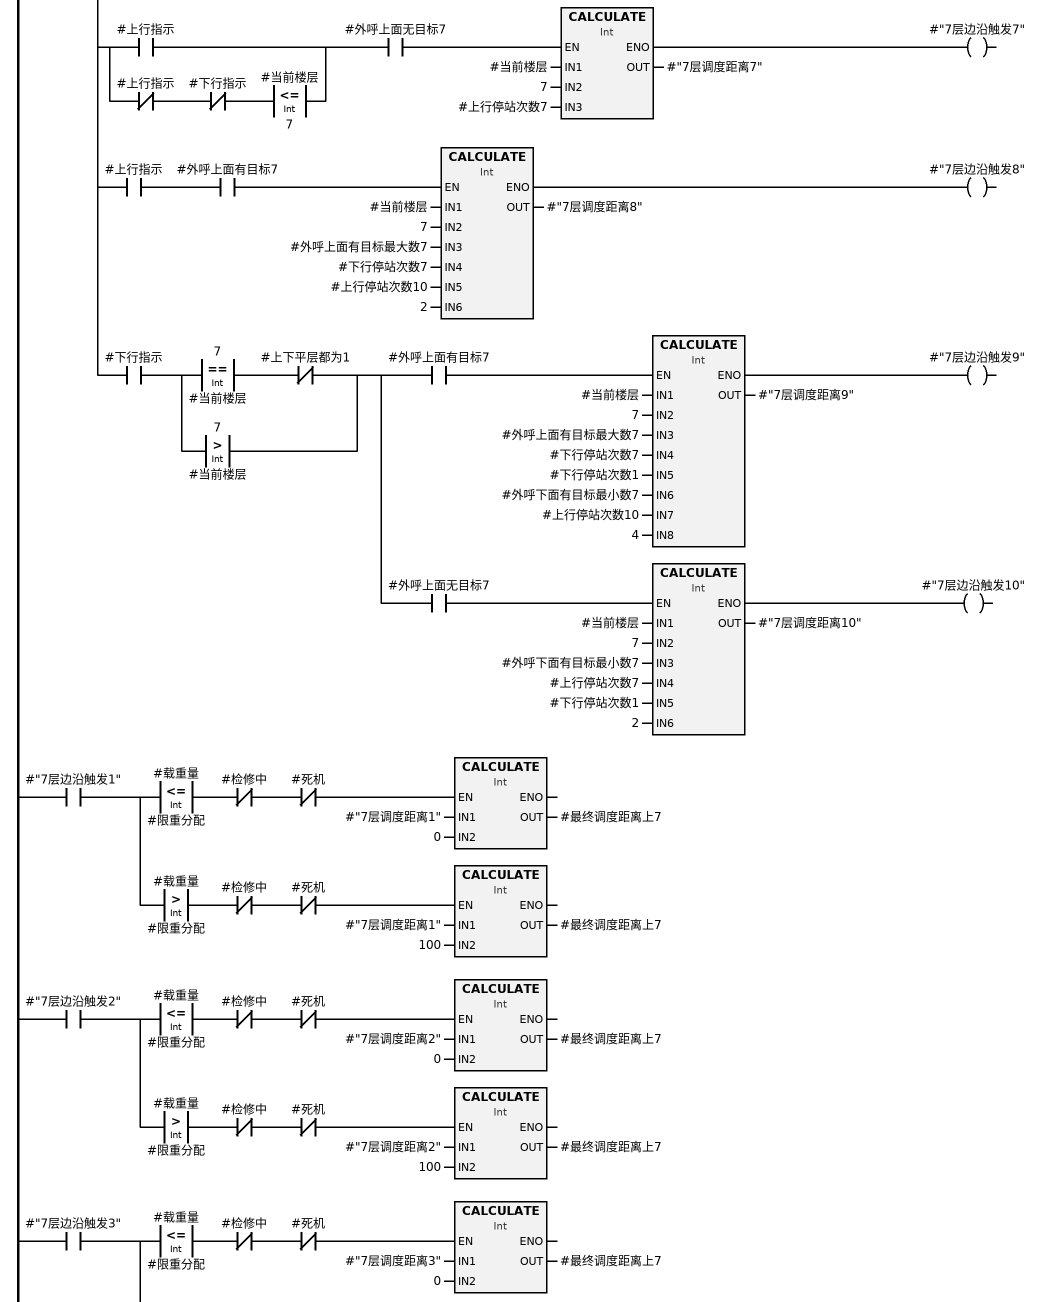
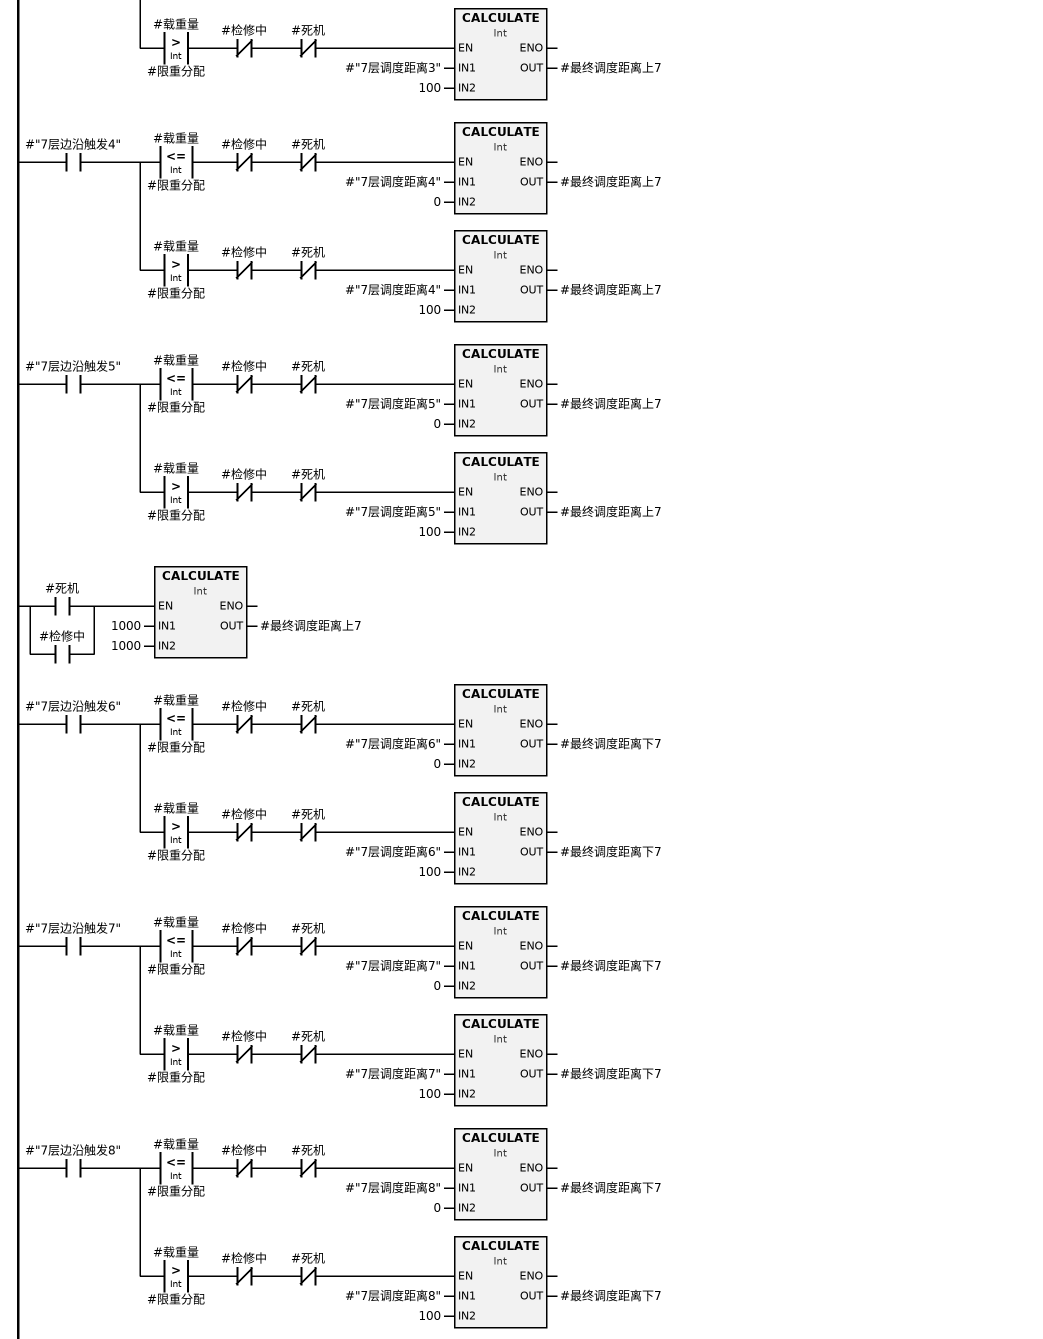
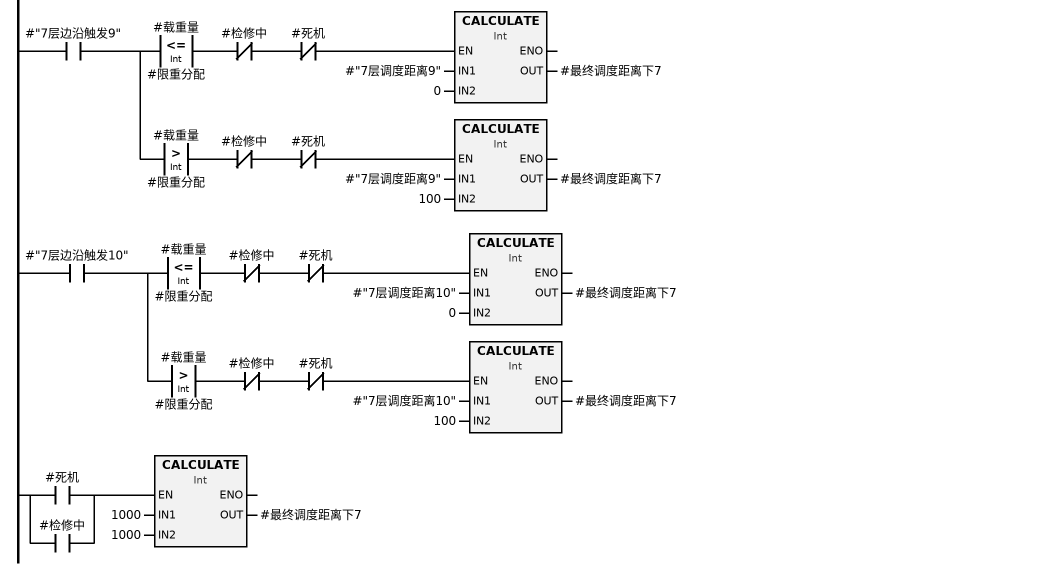
   RUNG wire#powerrail
      Contact( #上呼灯7 )
      wire#w1
      I_Contact( #上行指示 )
      I_Contact( #下行指示 )
      { S7_Templates := "SrcType := Int" } LE_Contact(in1 := #当前楼层, in2 := 7)
      wire#w2
      { S7_Templates := "SrcType := Int"; S7_Expression := "ABS(IN1-IN2)+IN3+IN3" } Calculate(in1 := #当前楼层, in2 := 7, in3 := #上行停站次数7, out => #"7层调度距离1")
      Coil( #"7层边沿触发1" )
   END_RUNG
   RUNG wire#w1
      Contact( #上行指示 )
      wire#w3
      { S7_Templates := "SrcType := Int" } EQ_Contact(in1 := 7, in2 := #当前楼层)
      Contact( #上下平层都为1 )
   END_RUNG wire#w2
   RUNG wire#w3
      { S7_Templates := "SrcType := Int" } GT_Contact(in1 := 7, in2 := #当前楼层)
   END_RUNG wire#w2
   RUNG wire#w1
      Contact( #下行指示 )
      wire#w4
      Contact( #外呼下面无目标7 )
      { S7_Templates := "SrcType := Int"; S7_Expression := "ABS(IN1-IN2)+IN3+IN3" } Calculate(in1 := #当前楼层, in2 := 7, in3 := #下行停站次数7, out => #"7层调度距离2")
      Coil( #"7层边沿触发2" )
   END_RUNG
   RUNG wire#w1
      I_Contact( #上行指示 )
      I_Contact( #下行指示 )
      { S7_Templates := "SrcType := Int" } GT_Contact(in1 := #当前楼层, in2 := 7)
   END_RUNG wire#w4
   RUNG wire#w1
      Contact( #下行指示 )
      Contact( #外呼下面有目标7 )
      { S7_Templates := "SrcType := Int"; S7_Expression := "ABS(IN3+IN3-IN1-IN2)+IN5+IN4+IN4+IN5+IN6" } Calculate(in1 := #当前楼层, in2 := 7, in3 := #外呼下面有目标最小数7, in4 := #上行停站次数7, in5 := #下行停站次数1, in6 := 2, out => #"7层调度距离3")
      Coil( #"7层边沿触发3" )
   END_RUNG
   RUNG wire#w1
      Contact( #上行指示 )
      wire#w5
      { S7_Templates := "SrcType := Int" } EQ_Contact(in1 := 7, in2 := #当前楼层)
      I_Contact( #上下平层都为1 )
      wire#w6
      Contact( #外呼下面有目标7 )
      { S7_Templates := "SrcType := Int"; S7_Expression := "ABS(IN3-IN1+IN3-IN6+IN2-IN6)+IN5+IN4+IN4+IN5+IN7+IN7+IN8" } Calculate(in1 := #当前楼层, in2 := 7, in3 := #外呼上面有目标最大数7, in4 := #上行停站次数10, in5 := #上行停站次数7, in6 := #外呼下面有目标最小数7, in7 := #下行停站次数1, in8 := 4, out => #"7层调度距离4")
      Coil( #"7层边沿触发4" )
   END_RUNG
   RUNG wire#w5
      { S7_Templates := "SrcType := Int" } LT_Contact(in1 := 7, in2 := #当前楼层)
   END_RUNG wire#w6
   RUNG wire#w6
      Contact( #外呼下面无目标7 )
      { S7_Templates := "SrcType := Int"; S7_Expression := "ABS(IN3-IN1+IN3-IN2)+IN5+IN4+IN4+IN5+IN6" } Calculate(in1 := #当前楼层, in2 := 7, in3 := #外呼上面有目标最大数7, in4 := #上行停站次数10, in5 := #下行停站次数7, in6 := 2, out => #"7层调度距离5")
      Coil( #"7层边沿触发5" )
   END_RUNG
   RUNG wire#powerrail
      Contact( #下呼灯7 )
      wire#w7
      I_Contact( #上行指示 )
      I_Contact( #下行指示 )
      { S7_Templates := "SrcType := Int" } GE_Contact(in1 := #当前楼层, in2 := 7)
      wire#w8
      { S7_Templates := "SrcType := Int"; S7_Expression := "ABS(IN1-IN2)+IN3+IN3" } Calculate(in1 := #当前楼层, in2 := 7, in3 := #下行停站次数7, out => #"7层调度距离6")
      Coil( #"7层边沿触发6" )
   END_RUNG
   RUNG wire#w7
      Contact( #下行指示 )
      wire#w9
      { S7_Templates := "SrcType := Int" } EQ_Contact(in1 := 7, in2 := #当前楼层)
      Contact( #上下平层都为1 )
   END_RUNG wire#w8
   RUNG wire#w9
      { S7_Templates := "SrcType := Int" } LT_Contact(in1 := 7, in2 := #当前楼层)
   END_RUNG wire#w8
   RUNG wire#w7
      Contact( #上行指示 )
      wire#w10
      Contact( #外呼上面无目标7 )
      { S7_Templates := "SrcType := Int"; S7_Expression := "ABS(IN1-IN2)+IN3+IN3" } Calculate(in1 := #当前楼层, in2 := 7, in3 := #上行停站次数7, out => #"7层调度距离7")
      Coil( #"7层边沿触发7" )
   END_RUNG
   RUNG wire#w7
      I_Contact( #上行指示 )
      I_Contact( #下行指示 )
      { S7_Templates := "SrcType := Int" } LE_Contact(in1 := #当前楼层, in2 := 7)
   END_RUNG wire#w10
   RUNG wire#w7
      Contact( #上行指示 )
      Contact( #外呼上面有目标7 )
      { S7_Templates := "SrcType := Int"; S7_Expression := "ABS(IN3+IN3-IN1-IN2)+IN4+IN5+IN4+IN5+IN6" } Calculate(in1 := #当前楼层, in2 := 7, in3 := #外呼上面有目标最大数7, in4 := #下行停站次数7, in5 := #上行停站次数10, in6 := 2, out => #"7层调度距离8")
      Coil( #"7层边沿触发8" )
   END_RUNG
   RUNG wire#w7
      Contact( #下行指示 )
      wire#w11
      { S7_Templates := "SrcType := Int" } EQ_Contact(in1 := 7, in2 := #当前楼层)
      I_Contact( #上下平层都为1 )
      wire#w12
      Contact( #外呼上面有目标7 )
      { S7_Templates := "SrcType := Int"; S7_Expression := "ABS(IN1-IN6+IN3-IN6+IN3-IN2)+IN5+IN4+IN4+IN5+IN7+IN7+IN8" } Calculate(in1 := #当前楼层, in2 := 7, in3 := #外呼上面有目标最大数7, in4 := #下行停站次数7, in5 := #下行停站次数1, in6 := #外呼下面有目标最小数7, in7 := #上行停站次数10, in8 := 4, out => #"7层调度距离9")
      Coil( #"7层边沿触发9" )
   END_RUNG
   RUNG wire#w11
      { S7_Templates := "SrcType := Int" } GT_Contact(in1 := 7, in2 := #当前楼层)
   END_RUNG wire#w12
   RUNG wire#w12
      Contact( #外呼上面无目标7 )
      { S7_Templates := "SrcType := Int"; S7_Expression := "ABS(IN1-IN3+IN2-IN3)+IN5+IN4+IN4+IN5+IN6" } Calculate(in1 := #当前楼层, in2 := 7, in3 := #外呼下面有目标最小数7, in4 := #上行停站次数7, in5 := #下行停站次数1, in6 := 2, out => #"7层调度距离10")
      Coil( #"7层边沿触发10" )
   END_RUNG
   RUNG wire#powerrail
      Contact( #"7层边沿触发1" )
      wire#w13
      { S7_Templates := "SrcType := Int" } LE_Contact(in1 := #载重量, in2 := #限重分配)
      I_Contact( #检修中 )
      I_Contact( #死机 )
      { S7_Templates := "SrcType := Int"; S7_Expression := "ABS(IN1+IN2)" } Calculate(in1 := #"7层调度距离1", in2 := 0, out => #最终调度距离上7)
   END_RUNG
   RUNG wire#w13
      { S7_Templates := "SrcType := Int" } GT_Contact(in1 := #载重量, in2 := #限重分配)
      I_Contact( #检修中 )
      I_Contact( #死机 )
      { S7_Templates := "SrcType := Int"; S7_Expression := "ABS(IN1+IN2)" } Calculate(in1 := #"7层调度距离1", in2 := 100, out => #最终调度距离上7)
   END_RUNG
   RUNG wire#powerrail
      Contact( #"7层边沿触发2" )
      wire#w14
      { S7_Templates := "SrcType := Int" } LE_Contact(in1 := #载重量, in2 := #限重分配)
      I_Contact( #检修中 )
      I_Contact( #死机 )
      { S7_Templates := "SrcType := Int"; S7_Expression := "ABS(IN1+IN2)" } Calculate(in1 := #"7层调度距离2", in2 := 0, out => #最终调度距离上7)
   END_RUNG
   RUNG wire#w14
      { S7_Templates := "SrcType := Int" } GT_Contact(in1 := #载重量, in2 := #限重分配)
      I_Contact( #检修中 )
      I_Contact( #死机 )
      { S7_Templates := "SrcType := Int"; S7_Expression := "ABS(IN1+IN2)" } Calculate(in1 := #"7层调度距离2", in2 := 100, out => #最终调度距离上7)
   END_RUNG
   RUNG wire#powerrail
      Contact( #"7层边沿触发3" )
      wire#w15
      { S7_Templates := "SrcType := Int" } LE_Contact(in1 := #载重量, in2 := #限重分配)
      I_Contact( #检修中 )
      I_Contact( #死机 )
      { S7_Templates := "SrcType := Int"; S7_Expression := "ABS(IN1+IN2)" } Calculate(in1 := #"7层调度距离3", in2 := 0, out => #最终调度距离上7)
   END_RUNG
   RUNG wire#w15
      { S7_Templates := "SrcType := Int" } GT_Contact(in1 := #载重量, in2 := #限重分配)
      I_Contact( #检修中 )
      I_Contact( #死机 )
      { S7_Templates := "SrcType := Int"; S7_Expression := "ABS(IN1+IN2)" } Calculate(in1 := #"7层调度距离3", in2 := 100, out => #最终调度距离上7)
   END_RUNG
   RUNG wire#powerrail
      Contact( #"7层边沿触发4" )
      wire#w16
      { S7_Templates := "SrcType := Int" } LE_Contact(in1 := #载重量, in2 := #限重分配)
      I_Contact( #检修中 )
      I_Contact( #死机 )
      { S7_Templates := "SrcType := Int"; S7_Expression := "ABS(IN1+IN2)" } Calculate(in1 := #"7层调度距离4", in2 := 0, out => #最终调度距离上7)
   END_RUNG
   RUNG wire#w16
      { S7_Templates := "SrcType := Int" } GT_Contact(in1 := #载重量, in2 := #限重分配)
      I_Contact( #检修中 )
      I_Contact( #死机 )
      { S7_Templates := "SrcType := Int"; S7_Expression := "ABS(IN1+IN2)" } Calculate(in1 := #"7层调度距离4", in2 := 100, out => #最终调度距离上7)
   END_RUNG
   RUNG wire#powerrail
      Contact( #"7层边沿触发5" )
      wire#w17
      { S7_Templates := "SrcType := Int" } LE_Contact(in1 := #载重量, in2 := #限重分配)
      I_Contact( #检修中 )
      I_Contact( #死机 )
      { S7_Templates := "SrcType := Int"; S7_Expression := "ABS(IN1+IN2)" } Calculate(in1 := #"7层调度距离5", in2 := 0, out => #最终调度距离上7)
   END_RUNG
   RUNG wire#w17
      { S7_Templates := "SrcType := Int" } GT_Contact(in1 := #载重量, in2 := #限重分配)
      I_Contact( #检修中 )
      I_Contact( #死机 )
      { S7_Templates := "SrcType := Int"; S7_Expression := "ABS(IN1+IN2)" } Calculate(in1 := #"7层调度距离5", in2 := 100, out => #最终调度距离上7)
   END_RUNG
   RUNG wire#powerrail
      Contact( #死机 )
      wire#w18
      { S7_Templates := "SrcType := Int"; S7_Expression := "ABS(IN1+IN2)" } Calculate(in1 := 1000, in2 := 1000, out => #最终调度距离上7)
   END_RUNG
   RUNG wire#powerrail
      Contact( #检修中 )
   END_RUNG wire#w18
   RUNG wire#powerrail
      Contact( #"7层边沿触发6" )
      wire#w19
      { S7_Templates := "SrcType := Int" } LE_Contact(in1 := #载重量, in2 := #限重分配)
      I_Contact( #检修中 )
      I_Contact( #死机 )
      { S7_Templates := "SrcType := Int"; S7_Expression := "ABS(IN1+IN2)" } Calculate(in1 := #"7层调度距离6", in2 := 0, out => #最终调度距离下7)
   END_RUNG
   RUNG wire#w19
      { S7_Templates := "SrcType := Int" } GT_Contact(in1 := #载重量, in2 := #限重分配)
      I_Contact( #检修中 )
      I_Contact( #死机 )
      { S7_Templates := "SrcType := Int"; S7_Expression := "ABS(IN1+IN2)" } Calculate(in1 := #"7层调度距离6", in2 := 100, out => #最终调度距离下7)
   END_RUNG
   RUNG wire#powerrail
      Contact( #"7层边沿触发7" )
      wire#w20
      { S7_Templates := "SrcType := Int" } LE_Contact(in1 := #载重量, in2 := #限重分配)
      I_Contact( #检修中 )
      I_Contact( #死机 )
      { S7_Templates := "SrcType := Int"; S7_Expression := "ABS(IN1+IN2)" } Calculate(in1 := #"7层调度距离7", in2 := 0, out => #最终调度距离下7)
   END_RUNG
   RUNG wire#w20
      { S7_Templates := "SrcType := Int" } GT_Contact(in1 := #载重量, in2 := #限重分配)
      I_Contact( #检修中 )
      I_Contact( #死机 )
      { S7_Templates := "SrcType := Int"; S7_Expression := "ABS(IN1+IN2)" } Calculate(in1 := #"7层调度距离7", in2 := 100, out => #最终调度距离下7)
   END_RUNG
   RUNG wire#powerrail
      Contact( #"7层边沿触发8" )
      wire#w21
      { S7_Templates := "SrcType := Int" } LE_Contact(in1 := #载重量, in2 := #限重分配)
      I_Contact( #检修中 )
      I_Contact( #死机 )
      { S7_Templates := "SrcType := Int"; S7_Expression := "ABS(IN1+IN2)" } Calculate(in1 := #"7层调度距离8", in2 := 0, out => #最终调度距离下7)
   END_RUNG
   RUNG wire#w21
      { S7_Templates := "SrcType := Int" } GT_Contact(in1 := #载重量, in2 := #限重分配)
      I_Contact( #检修中 )
      I_Contact( #死机 )
      { S7_Templates := "SrcType := Int"; S7_Expression := "ABS(IN1+IN2)" } Calculate(in1 := #"7层调度距离8", in2 := 100, out => #最终调度距离下7)
   END_RUNG
   RUNG wire#powerrail
      Contact( #"7层边沿触发9" )
      wire#w22
      { S7_Templates := "SrcType := Int" } LE_Contact(in1 := #载重量, in2 := #限重分配)
      I_Contact( #检修中 )
      I_Contact( #死机 )
      { S7_Templates := "SrcType := Int"; S7_Expression := "ABS(IN1+IN2)" } Calculate(in1 := #"7层调度距离9", in2 := 0, out => #最终调度距离下7)
   END_RUNG
   RUNG wire#w22
      { S7_Templates := "SrcType := Int" } GT_Contact(in1 := #载重量, in2 := #限重分配)
      I_Contact( #检修中 )
      I_Contact( #死机 )
      { S7_Templates := "SrcType := Int"; S7_Expression := "ABS(IN1+IN2)" } Calculate(in1 := #"7层调度距离9", in2 := 100, out => #最终调度距离下7)
   END_RUNG
   RUNG wire#powerrail
      Contact( #"7层边沿触发10" )
      wire#w23
      { S7_Templates := "SrcType := Int" } LE_Contact(in1 := #载重量, in2 := #限重分配)
      I_Contact( #检修中 )
      I_Contact( #死机 )
      { S7_Templates := "SrcType := Int"; S7_Expression := "ABS(IN1+IN2)" } Calculate(in1 := #"7层调度距离10", in2 := 0, out => #最终调度距离下7)
   END_RUNG
   RUNG wire#w23
      { S7_Templates := "SrcType := Int" } GT_Contact(in1 := #载重量, in2 := #限重分配)
      I_Contact( #检修中 )
      I_Contact( #死机 )
      { S7_Templates := "SrcType := Int"; S7_Expression := "ABS(IN1+IN2)" } Calculate(in1 := #"7层调度距离10", in2 := 100, out => #最终调度距离下7)
   END_RUNG
   RUNG wire#powerrail
      Contact( #死机 )
      wire#w24
      { S7_Templates := "SrcType := Int"; S7_Expression := "ABS(IN1+IN2)" } Calculate(in1 := 1000, in2 := 1000, out => #最终调度距离下7)
   END_RUNG
   RUNG wire#powerrail
      Contact( #检修中 )
   END_RUNG wire#w24
   // the same network as SCL:
   #_w1 := #上呼灯7 AND ((NOT #上行指示 AND NOT #下行指示 AND (#当前楼层 <= 7)) OR (#上行指示 AND (((7 = #当前楼层) AND #上下平层都为1) OR (7 > #当前楼层))));
   IF #_w1 THEN #"7层调度距离1" := ABS(#当前楼层-7)+#上行停站次数7+#上行停站次数7; END_IF;
   #"7层边沿触发1" := #_w1;
   #_w2 := #上呼灯7 AND (#下行指示 OR (NOT #上行指示 AND NOT #下行指示 AND (#当前楼层 > 7))) AND #外呼下面无目标7;
   IF #_w2 THEN #"7层调度距离2" := ABS(#当前楼层-7)+#下行停站次数7+#下行停站次数7; END_IF;
   #"7层边沿触发2" := #_w2;
   #_w3 := #上呼灯7 AND #下行指示 AND #外呼下面有目标7;
   IF #_w3 THEN
       #"7层调度距离3" := ABS(#外呼下面有目标最小数7+#外呼下面有目标最小数7-#当前楼层-7)+#下行停站次数1+#上行停站次数7+#上行停站次数7+#下行停站次数1+2;
   END_IF;
   #"7层边沿触发3" := #_w3;
   #_w4 := #上呼灯7 AND #上行指示 AND (((7 = #当前楼层) AND NOT #上下平层都为1) OR (7 < #当前楼层));
   #_w5 := #_w4 AND #外呼下面有目标7;
   IF #_w5 THEN
       #"7层调度距离4" := ABS(#外呼上面有目标最大数7-#当前楼层+#外呼上面有目标最大数7-#外呼下面有目标最小数7+7-#外呼下面有目标最小数7)+#上行停站次数7+#上行停站次数10+#上行停站次数10+#上行停站次数7+#下行停站次数1+#下行停站次数1+4;
   END_IF;
   #"7层边沿触发4" := #_w5;
   #_w6 := #_w4 AND #外呼下面无目标7;
   IF #_w6 THEN
       #"7层调度距离5" := ABS(#外呼上面有目标最大数7-#当前楼层+#外呼上面有目标最大数7-7)+#下行停站次数7+#上行停站次数10+#上行停站次数10+#下行停站次数7+2;
   END_IF;
   #"7层边沿触发5" := #_w6;
   #_w7 := #下呼灯7 AND ((NOT #上行指示 AND NOT #下行指示 AND (#当前楼层 >= 7)) OR (#下行指示 AND (((7 = #当前楼层) AND #上下平层都为1) OR (7 < #当前楼层))));
   IF #_w7 THEN #"7层调度距离6" := ABS(#当前楼层-7)+#下行停站次数7+#下行停站次数7; END_IF;
   #"7层边沿触发6" := #_w7;
   #_w8 := #下呼灯7 AND (#上行指示 OR (NOT #上行指示 AND NOT #下行指示 AND (#当前楼层 <= 7))) AND #外呼上面无目标7;
   IF #_w8 THEN #"7层调度距离7" := ABS(#当前楼层-7)+#上行停站次数7+#上行停站次数7; END_IF;
   #"7层边沿触发7" := #_w8;
   #_w9 := #下呼灯7 AND #上行指示 AND #外呼上面有目标7;
   IF #_w9 THEN
       #"7层调度距离8" := ABS(#外呼上面有目标最大数7+#外呼上面有目标最大数7-#当前楼层-7)+#下行停站次数7+#上行停站次数10+#下行停站次数7+#上行停站次数10+2;
   END_IF;
   #"7层边沿触发8" := #_w9;
   #_w10 := #下呼灯7 AND #下行指示 AND (((7 = #当前楼层) AND NOT #上下平层都为1) OR (7 > #当前楼层));
   #_w11 := #_w10 AND #外呼上面有目标7;
   IF #_w11 THEN
       #"7层调度距离9" := ABS(#当前楼层-#外呼下面有目标最小数7+#外呼上面有目标最大数7-#外呼下面有目标最小数7+#外呼上面有目标最大数7-7)+#下行停站次数1+#下行停站次数7+#下行停站次数7+#下行停站次数1+#上行停站次数10+#上行停站次数10+4;
   END_IF;
   #"7层边沿触发9" := #_w11;
   #_w12 := #_w10 AND #外呼上面无目标7;
   IF #_w12 THEN
       #"7层调度距离10" := ABS(#当前楼层-#外呼下面有目标最小数7+7-#外呼下面有目标最小数7)+#下行停站次数1+#上行停站次数7+#上行停站次数7+#下行停站次数1+2;
   END_IF;
   #"7层边沿触发10" := #_w12;
   IF #"7层边沿触发1" AND (#载重量 <= #限重分配) AND NOT #检修中 AND NOT #死机 THEN #最终调度距离上7 := ABS(#"7层调度距离1"+0); END_IF;
   IF #"7层边沿触发1" AND (#载重量 > #限重分配) AND NOT #检修中 AND NOT #死机 THEN #最终调度距离上7 := ABS(#"7层调度距离1"+100); END_IF;
   IF #"7层边沿触发2" AND (#载重量 <= #限重分配) AND NOT #检修中 AND NOT #死机 THEN #最终调度距离上7 := ABS(#"7层调度距离2"+0); END_IF;
   IF #"7层边沿触发2" AND (#载重量 > #限重分配) AND NOT #检修中 AND NOT #死机 THEN #最终调度距离上7 := ABS(#"7层调度距离2"+100); END_IF;
   IF #"7层边沿触发3" AND (#载重量 <= #限重分配) AND NOT #检修中 AND NOT #死机 THEN #最终调度距离上7 := ABS(#"7层调度距离3"+0); END_IF;
   IF #"7层边沿触发3" AND (#载重量 > #限重分配) AND NOT #检修中 AND NOT #死机 THEN #最终调度距离上7 := ABS(#"7层调度距离3"+100); END_IF;
   IF #"7层边沿触发4" AND (#载重量 <= #限重分配) AND NOT #检修中 AND NOT #死机 THEN #最终调度距离上7 := ABS(#"7层调度距离4"+0); END_IF;
   IF #"7层边沿触发4" AND (#载重量 > #限重分配) AND NOT #检修中 AND NOT #死机 THEN #最终调度距离上7 := ABS(#"7层调度距离4"+100); END_IF;
   IF #"7层边沿触发5" AND (#载重量 <= #限重分配) AND NOT #检修中 AND NOT #死机 THEN #最终调度距离上7 := ABS(#"7层调度距离5"+0); END_IF;
   IF #"7层边沿触发5" AND (#载重量 > #限重分配) AND NOT #检修中 AND NOT #死机 THEN #最终调度距离上7 := ABS(#"7层调度距离5"+100); END_IF;
   IF #死机 OR #检修中 THEN #最终调度距离上7 := ABS(1000+1000); END_IF;
   IF #"7层边沿触发6" AND (#载重量 <= #限重分配) AND NOT #检修中 AND NOT #死机 THEN #最终调度距离下7 := ABS(#"7层调度距离6"+0); END_IF;
   IF #"7层边沿触发6" AND (#载重量 > #限重分配) AND NOT #检修中 AND NOT #死机 THEN #最终调度距离下7 := ABS(#"7层调度距离6"+100); END_IF;
   IF #"7层边沿触发7" AND (#载重量 <= #限重分配) AND NOT #检修中 AND NOT #死机 THEN #最终调度距离下7 := ABS(#"7层调度距离7"+0); END_IF;
   IF #"7层边沿触发7" AND (#载重量 > #限重分配) AND NOT #检修中 AND NOT #死机 THEN #最终调度距离下7 := ABS(#"7层调度距离7"+100); END_IF;
   IF #"7层边沿触发8" AND (#载重量 <= #限重分配) AND NOT #检修中 AND NOT #死机 THEN #最终调度距离下7 := ABS(#"7层调度距离8"+0); END_IF;
   IF #"7层边沿触发8" AND (#载重量 > #限重分配) AND NOT #检修中 AND NOT #死机 THEN #最终调度距离下7 := ABS(#"7层调度距离8"+100); END_IF;
   IF #"7层边沿触发9" AND (#载重量 <= #限重分配) AND NOT #检修中 AND NOT #死机 THEN #最终调度距离下7 := ABS(#"7层调度距离9"+0); END_IF;
   IF #"7层边沿触发9" AND (#载重量 > #限重分配) AND NOT #检修中 AND NOT #死机 THEN #最终调度距离下7 := ABS(#"7层调度距离9"+100); END_IF;
   IF #"7层边沿触发10" AND (#载重量 <= #限重分配) AND NOT #检修中 AND NOT #死机 THEN #最终调度距离下7 := ABS(#"7层调度距离10"+0); END_IF;
   IF #"7层边沿触发10" AND (#载重量 > #限重分配) AND NOT #检修中 AND NOT #死机 THEN #最终调度距离下7 := ABS(#"7层调度距离10"+100); END_IF;
   IF #死机 OR #检修中 THEN #最终调度距离下7 := ABS(1000+1000); END_IF;
END_REGION

REGION Network 7: 8层调度距离
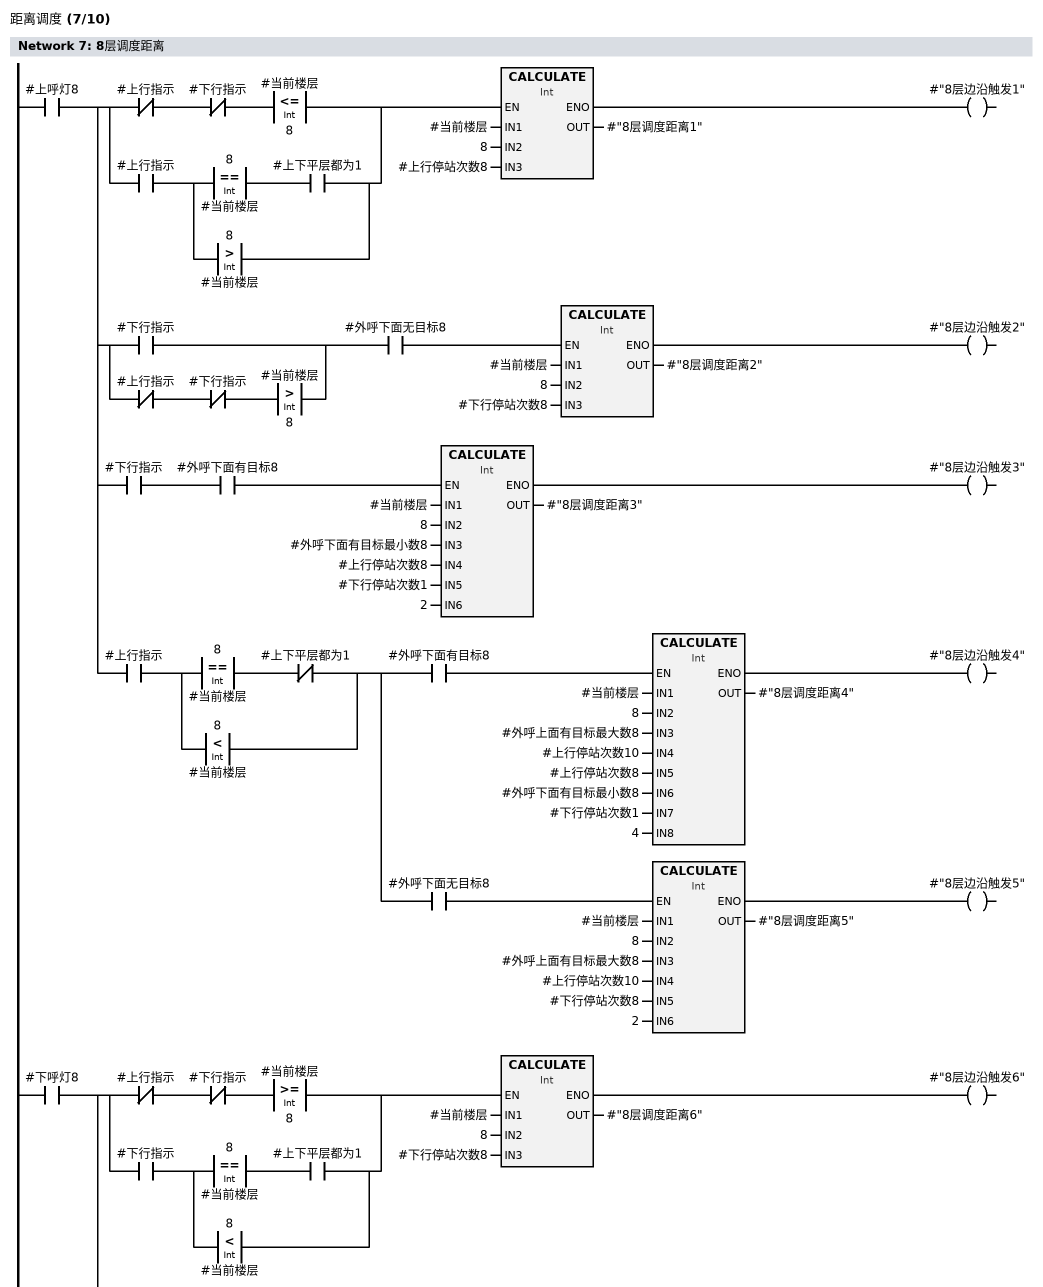
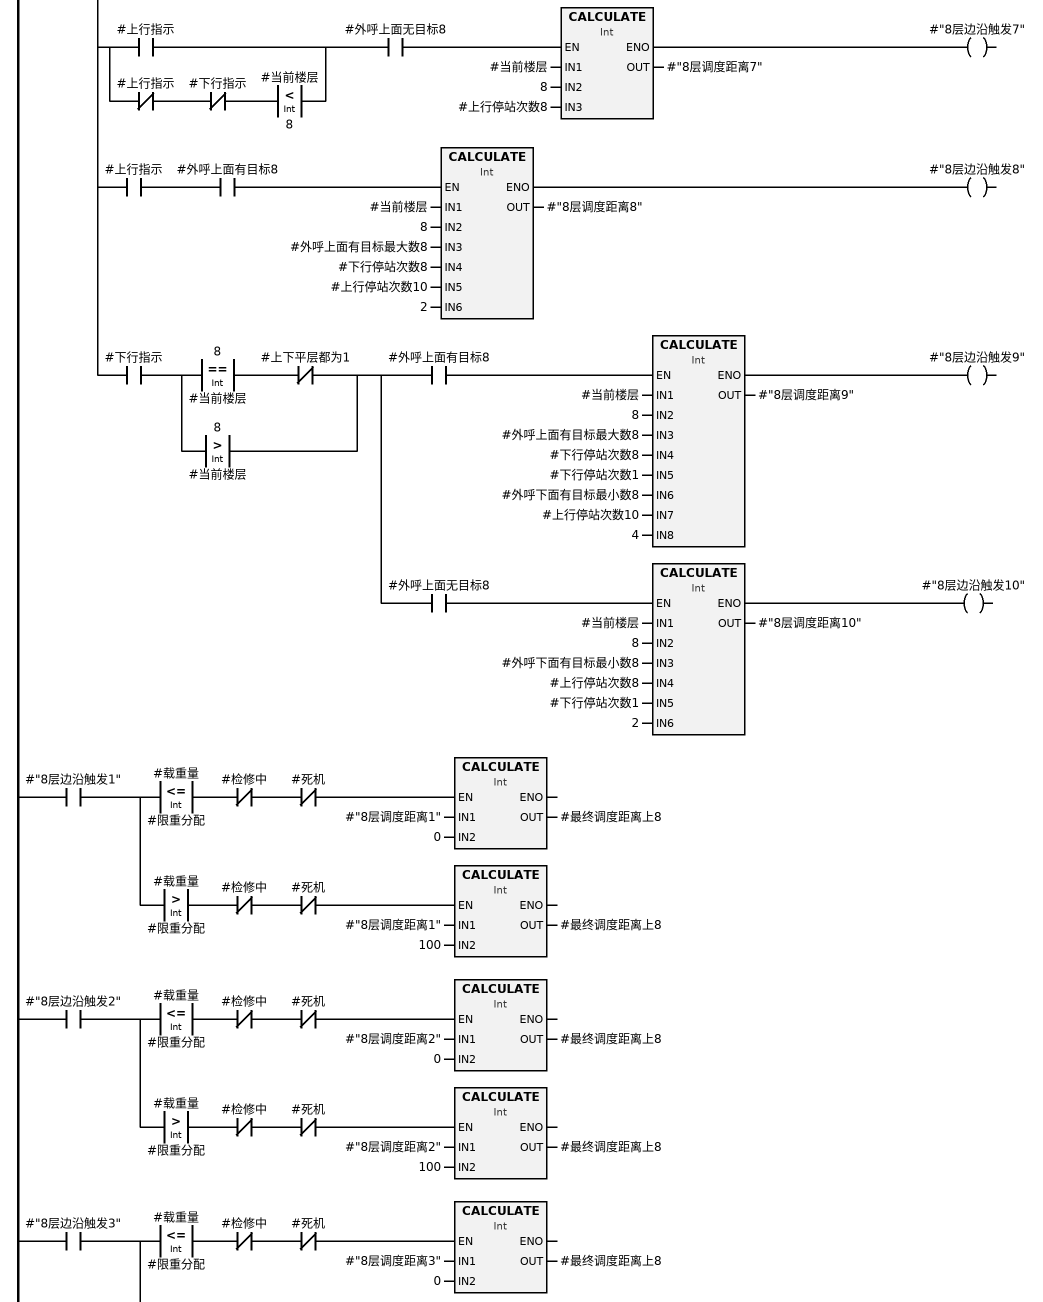
